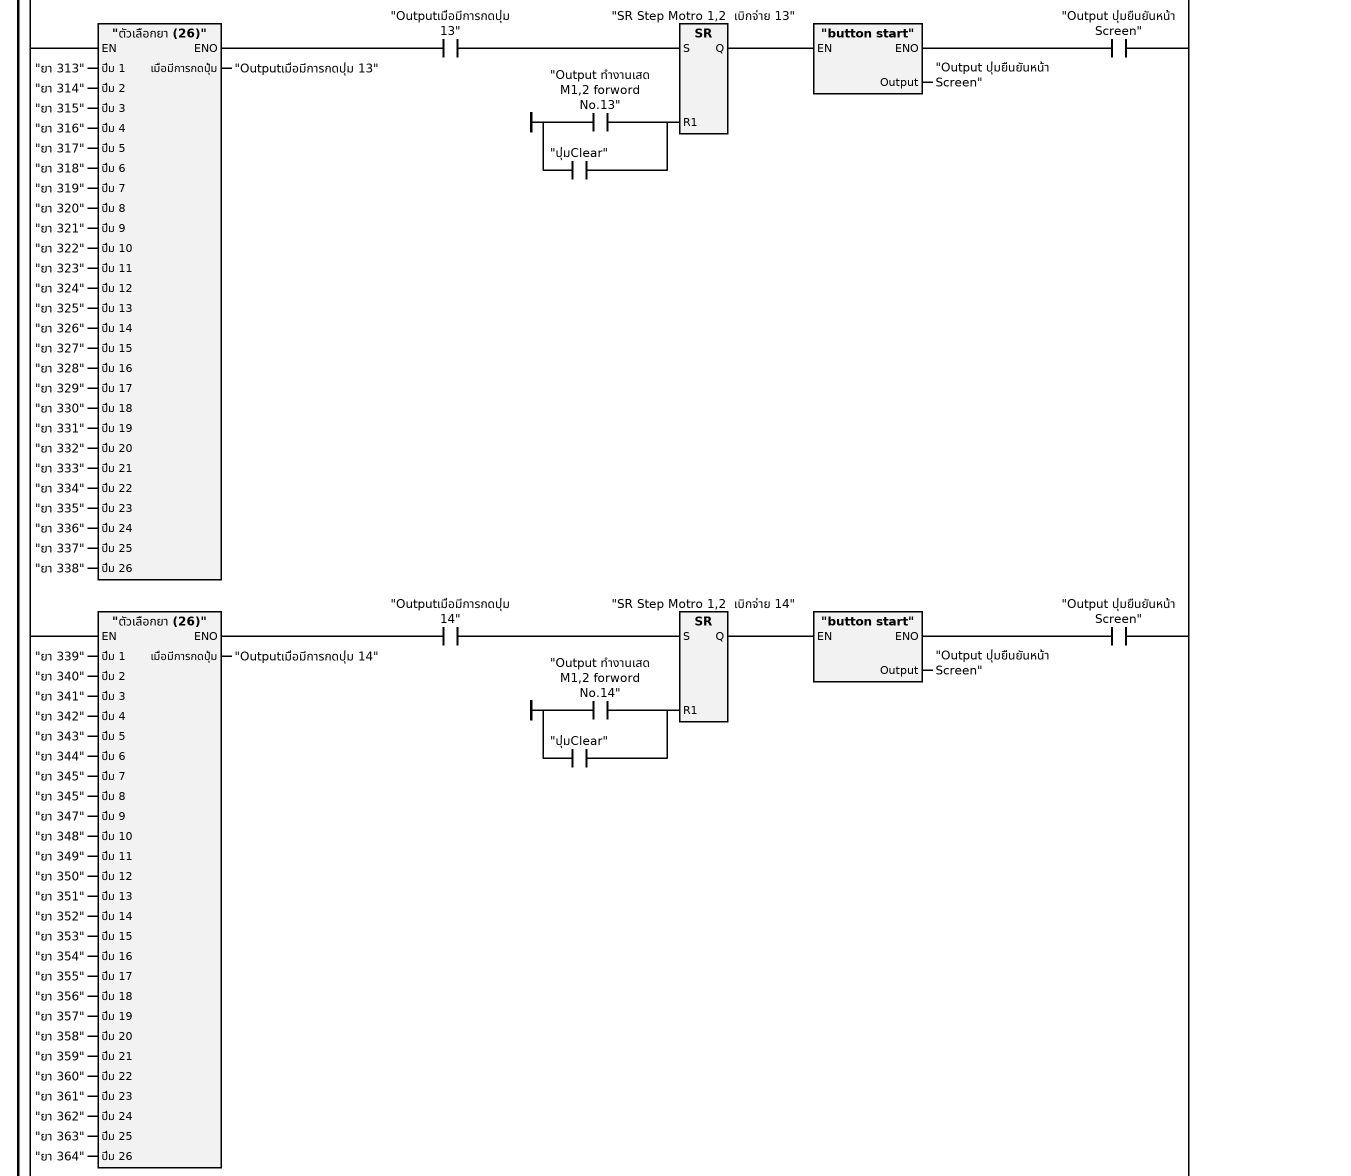
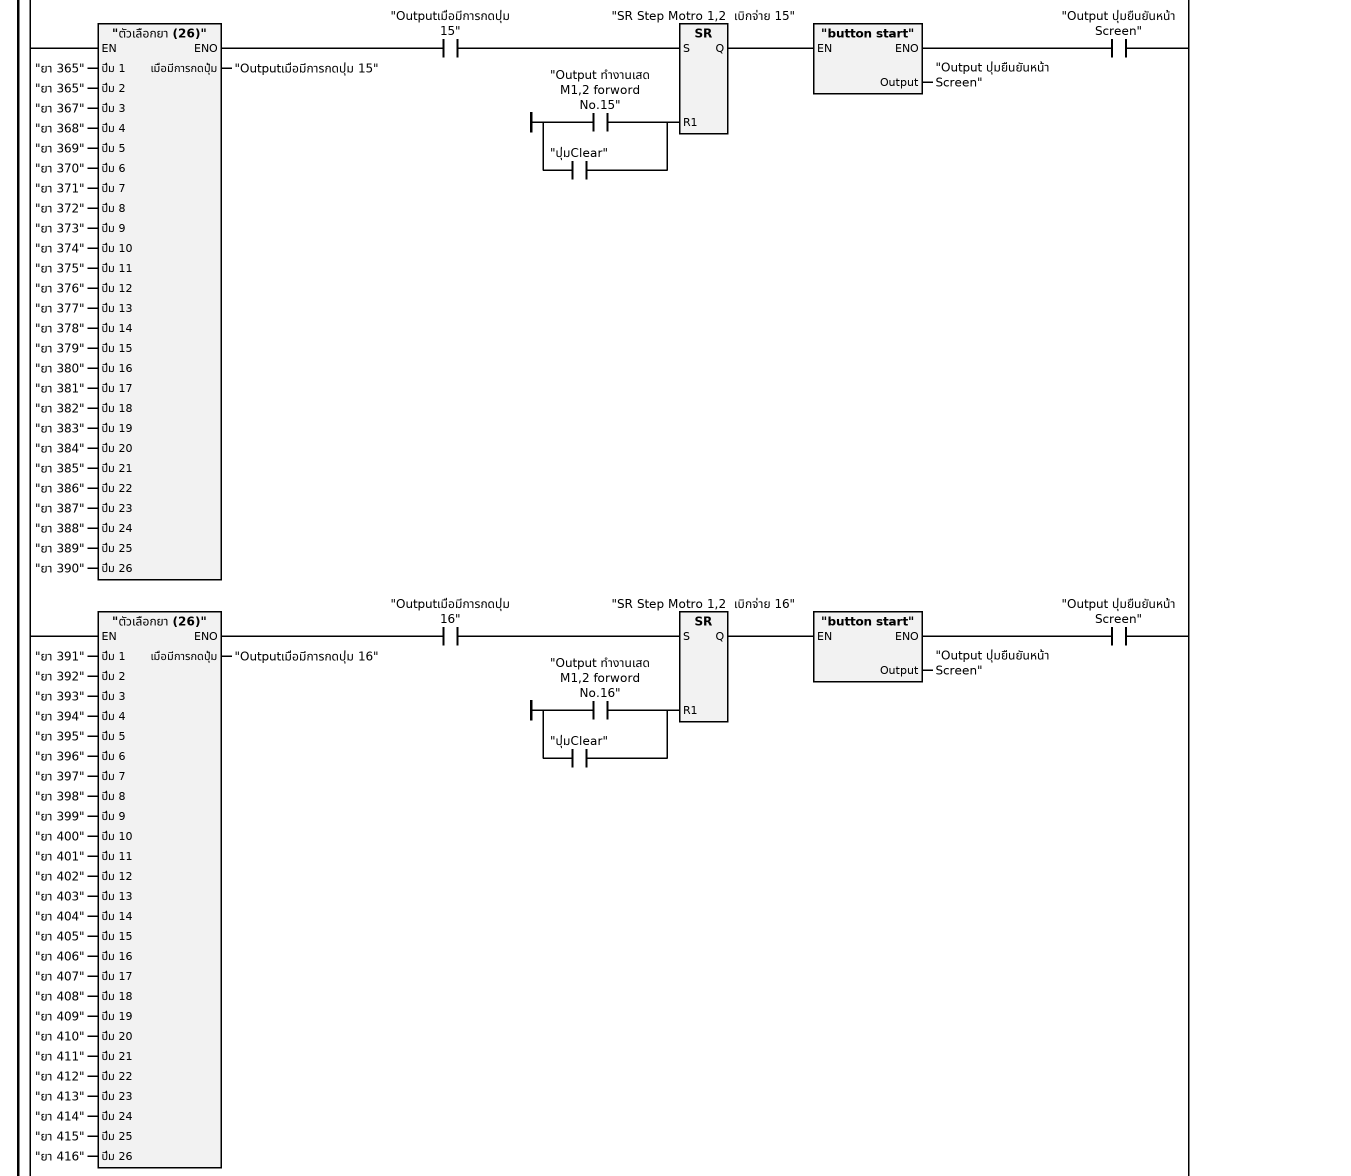
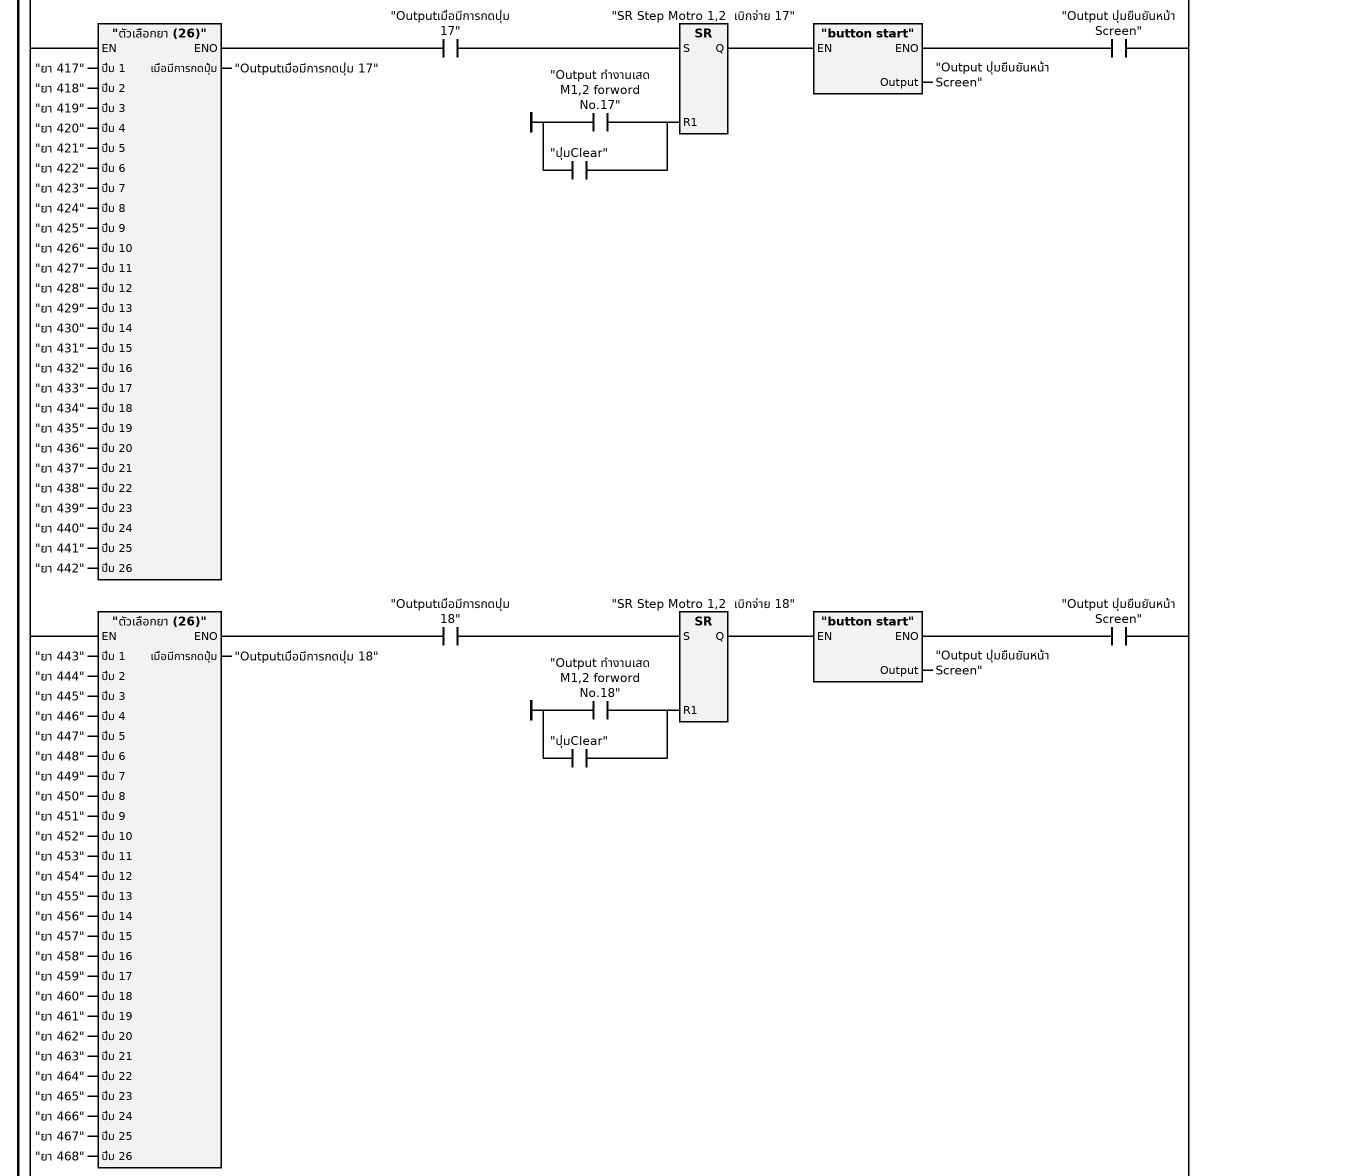
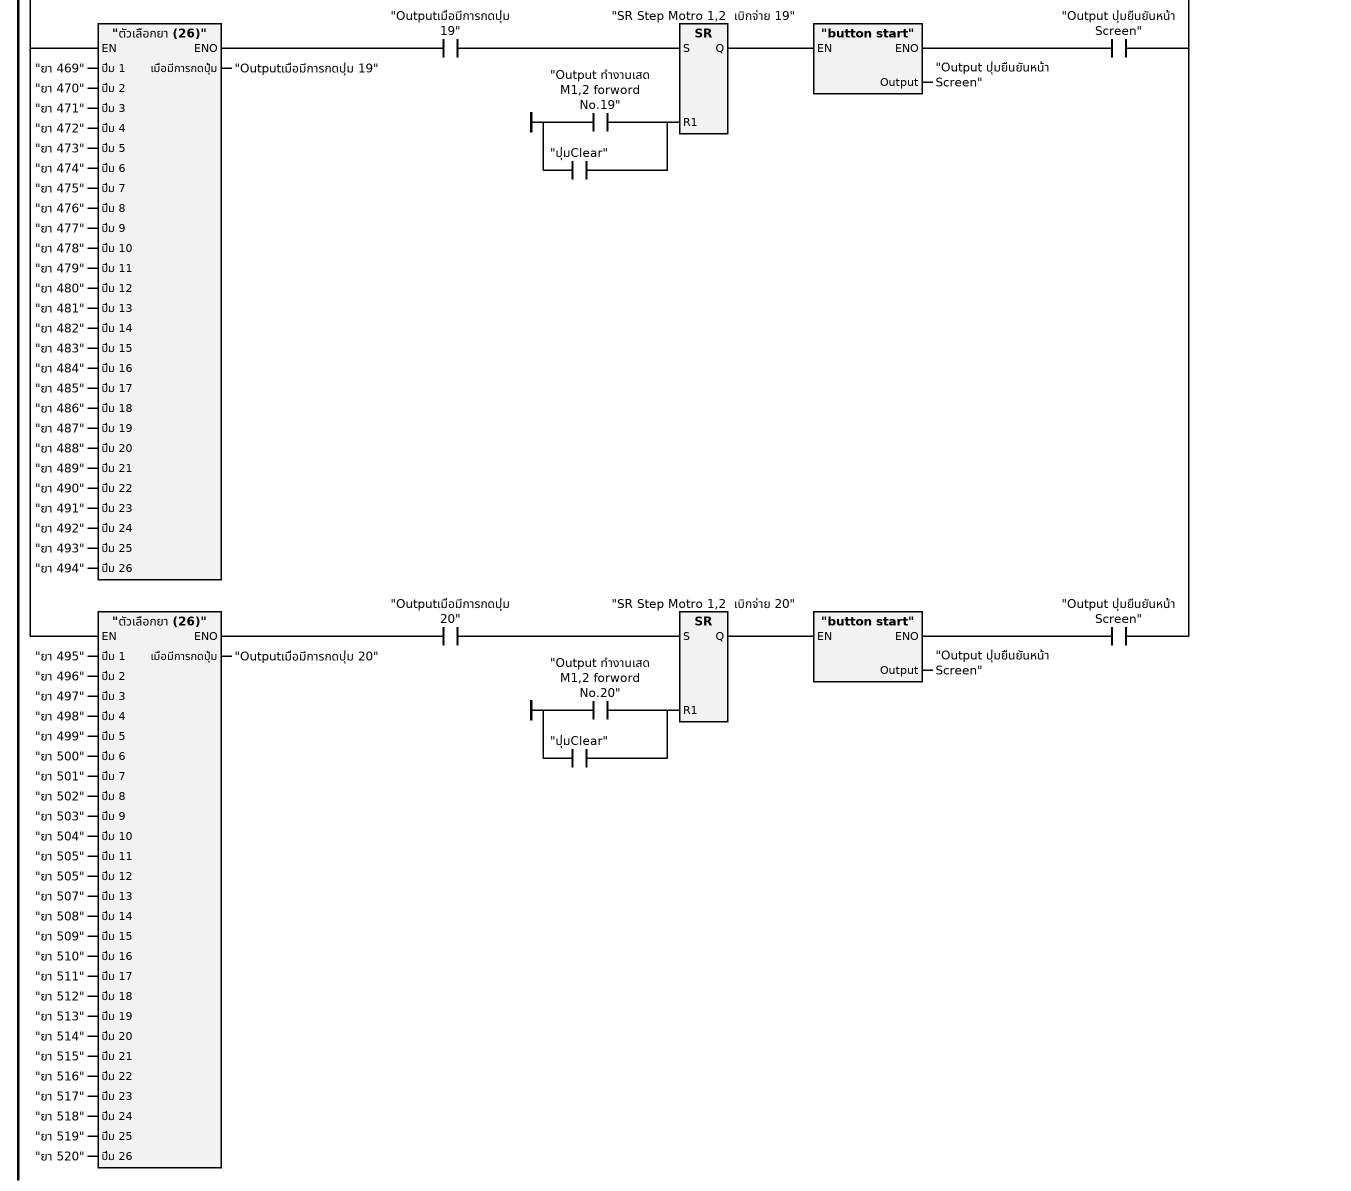
   RUNG wire#powerrail
      "ตัวเลือกยา (26)"("ปึ่ม 1" := "ยา 1", "ปึ่ม 2" := "ยา 2", "ปึ่ม 3" := "ยา 3", "ปึ่ม 4" := "ยา 4", "ปึ่ม 5" := "ยา 5", "ปึ่ม 6" := "ยา 6", "ปึ่ม 7" := "ยา 7", "ปึ่ม 8" := "ยา 8", "ปึ่ม 9" := "ยา 9", "ปึ่ม 10" := "ยา 10", "ปึ่ม 11" := "ยา 11", "ปึ่ม 12" := "ยา 12", "ปึ่ม 13" := "ยา 13", "ปึ่ม 14" := "ยา 14", "ปึ่ม 15" := "ยา 15", "ปึ่ม 16" := "ยา 16", "ปึ่ม 17" := "ยา 17", "ปึ่ม 18" := "ยา 18", "ปึ่ม 19" := "ยา 19", "ปึ่ม 20" := "ยา 20", "ปึ่ม 21" := "ยา 21", "ปึ่ม 22" := "ยา 22", "ปึ่ม 23" := "ยา 23", "ปึ่ม 24" := "ยา 24", "ปึ่ม 25" := "ยา 25", "ปึ่ม 26" := "ยา 26", "เมื่ิอมีการกดปุ้ม" => "Outputเมื่อมีการกดปุ่ม 1")
      Contact( "Outputเมื่อมีการกดปุ่ม 1" )
      S_SR(operand := "SR Step Motro 1,2  เบิกจ่าย 1", r1 := wire#w1)
      "button start"(Output => "Output ปุ่มยืนยันหน้า Screen")
      Contact( "Output ปุ่มยืนยันหน้า Screen" )
      wire#w2
      Coil( #"Stepper Motor  ทำงาน" )
   END_RUNG
   RUNG wire#powerrail
      Contact( "Output ทำงานเสด M1,2 forword No.1" )
   END_RUNG wire#w1
   RUNG wire#powerrail
      Contact( "ปุ่มClear" )
   END_RUNG wire#w1
   RUNG wire#powerrail
      "ตัวเลือกยา (26)"("ปึ่ม 1" := "ยา 27", "ปึ่ม 2" := "ยา 28", "ปึ่ม 3" := "ยา 29", "ปึ่ม 4" := "ยา 30", "ปึ่ม 5" := "ยา 31", "ปึ่ม 6" := "ยา 32", "ปึ่ม 7" := "ยา 33", "ปึ่ม 8" := "ยา 34", "ปึ่ม 9" := "ยา 35", "ปึ่ม 10" := "ยา 36", "ปึ่ม 11" := "ยา 37", "ปึ่ม 12" := "ยา 38", "ปึ่ม 13" := "ยา 39", "ปึ่ม 14" := "ยา 40", "ปึ่ม 15" := "ยา 41", "ปึ่ม 16" := "ยา 42", "ปึ่ม 17" := "ยา 43", "ปึ่ม 18" := "ยา 44", "ปึ่ม 19" := "ยา 45", "ปึ่ม 20" := "ยา 46", "ปึ่ม 21" := "ยา 47", "ปึ่ม 22" := "ยา 48", "ปึ่ม 23" := "ยา 49", "ปึ่ม 24" := "ยา 50", "ปึ่ม 25" := "ยา 51", "ปึ่ม 26" := "ยา 52", "เมื่ิอมีการกดปุ้ม" => "Outputเมื่อมีการกดปุ่ม 2")
      Contact( "Outputเมื่อมีการกดปุ่ม 2" )
      S_SR(operand := "SR Step Motro 1,2  เบิกจ่าย 2", r1 := wire#w3)
      "button start"(Output => "Output ปุ่มยืนยันหน้า Screen")
      Contact( "Output ปุ่มยืนยันหน้า Screen" )
   END_RUNG wire#w2
   RUNG wire#powerrail
      Contact( "Output ทำงานเสด M1,2 forword No.2" )
   END_RUNG wire#w3
   RUNG wire#powerrail
      Contact( "ปุ่มClear" )
   END_RUNG wire#w3
   RUNG wire#powerrail
      "ตัวเลือกยา (26)"("ปึ่ม 1" := "ยา 53", "ปึ่ม 2" := "ยา 54", "ปึ่ม 3" := "ยา 55", "ปึ่ม 4" := "ยา 56", "ปึ่ม 5" := "ยา 57", "ปึ่ม 6" := "ยา 58", "ปึ่ม 7" := "ยา 59", "ปึ่ม 8" := "ยา 60", "ปึ่ม 9" := "ยา 61", "ปึ่ม 10" := "ยา 62", "ปึ่ม 11" := "ยา 63", "ปึ่ม 12" := "ยา 64", "ปึ่ม 13" := "ยา 65", "ปึ่ม 14" := "ยา 66", "ปึ่ม 15" := "ยา 67", "ปึ่ม 16" := "ยา 68", "ปึ่ม 17" := "ยา 69", "ปึ่ม 18" := "ยา 70", "ปึ่ม 19" := "ยา 71", "ปึ่ม 20" := "ยา 72", "ปึ่ม 21" := "ยา 73", "ปึ่ม 22" := "ยา 74", "ปึ่ม 23" := "ยา 75", "ปึ่ม 24" := "ยา 76", "ปึ่ม 25" := "ยา 77", "ปึ่ม 26" := "ยา 78", "เมื่ิอมีการกดปุ้ม" => "Outputเมื่อมีการกดปุ่ม 3")
      Contact( "Outputเมื่อมีการกดปุ่ม 3" )
      S_SR(operand := "SR Step Motro 1,2  เบิกจ่าย 3", r1 := wire#w4)
      "button start"(Output => "Output ปุ่มยืนยันหน้า Screen")
      Contact( "Output ปุ่มยืนยันหน้า Screen" )
   END_RUNG wire#w2
   RUNG wire#powerrail
      Contact( "Output ทำงานเสด M1,2 forword No.3" )
   END_RUNG wire#w4
   RUNG wire#powerrail
      Contact( "ปุ่มClear" )
   END_RUNG wire#w4
   RUNG wire#powerrail
      "ตัวเลือกยา (26)"("ปึ่ม 1" := "ยา 79", "ปึ่ม 2" := "ยา 80", "ปึ่ม 3" := "ยา 81", "ปึ่ม 4" := "ยา 82", "ปึ่ม 5" := "ยา 83", "ปึ่ม 6" := "ยา 84", "ปึ่ม 7" := "ยา 85", "ปึ่ม 8" := "ยา 86", "ปึ่ม 9" := "ยา 87", "ปึ่ม 10" := "ยา 88", "ปึ่ม 11" := "ยา 89", "ปึ่ม 12" := "ยา 90", "ปึ่ม 13" := "ยา 91", "ปึ่ม 14" := "ยา 92", "ปึ่ม 15" := "ยา 93", "ปึ่ม 16" := "ยา 94", "ปึ่ม 17" := "ยา 95", "ปึ่ม 18" := "ยา 96", "ปึ่ม 19" := "ยา 97", "ปึ่ม 20" := "ยา 98", "ปึ่ม 21" := "ยา 99", "ปึ่ม 22" := "ยา 100", "ปึ่ม 23" := "ยา 101", "ปึ่ม 24" := "ยา 102", "ปึ่ม 25" := "ยา 103", "ปึ่ม 26" := "ยา 104", "เมื่ิอมีการกดปุ้ม" => "Outputเมื่อมีการกดปุ่ม 4")
      Contact( "Outputเมื่อมีการกดปุ่ม 4" )
      S_SR(operand := "SR Step Motro 1,2  เบิกจ่าย 4", r1 := wire#w5)
      "button start"(Output => "Output ปุ่มยืนยันหน้า Screen")
      Contact( "Output ปุ่มยืนยันหน้า Screen" )
   END_RUNG wire#w2
   RUNG wire#powerrail
      Contact( "Output ทำงานเสด M1,2 forword No.4" )
   END_RUNG wire#w5
   RUNG wire#powerrail
      Contact( "ปุ่มClear" )
   END_RUNG wire#w5
   RUNG wire#powerrail
      "ตัวเลือกยา (26)"("ปึ่ม 1" := "ยา 105", "ปึ่ม 2" := "ยา 106", "ปึ่ม 3" := "ยา 107", "ปึ่ม 4" := "ยา 108", "ปึ่ม 5" := "ยา 109", "ปึ่ม 6" := "ยา 110", "ปึ่ม 7" := "ยา 111", "ปึ่ม 8" := "ยา 112", "ปึ่ม 9" := "ยา 113", "ปึ่ม 10" := "ยา 114", "ปึ่ม 11" := "ยา 115", "ปึ่ม 12" := "ยา 116", "ปึ่ม 13" := "ยา 117", "ปึ่ม 14" := "ยา 118", "ปึ่ม 15" := "ยา 119", "ปึ่ม 16" := "ยา 120", "ปึ่ม 17" := "ยา 121", "ปึ่ม 18" := "ยา 122", "ปึ่ม 19" := "ยา 123", "ปึ่ม 20" := "ยา 124", "ปึ่ม 21" := "ยา 125", "ปึ่ม 22" := "ยา 126", "ปึ่ม 23" := "ยา 127", "ปึ่ม 24" := "ยา 128", "ปึ่ม 25" := "ยา 129", "ปึ่ม 26" := "ยา 130", "เมื่ิอมีการกดปุ้ม" => "Outputเมื่อมีการกดปุ่ม 5")
      Contact( "Outputเมื่อมีการกดปุ่ม 5" )
      S_SR(operand := "SR Step Motro 1,2  เบิกจ่าย 5", r1 := wire#w6)
      "button start"(Output => "Output ปุ่มยืนยันหน้า Screen")
      Contact( "Output ปุ่มยืนยันหน้า Screen" )
   END_RUNG wire#w2
   RUNG wire#powerrail
      Contact( "Output ทำงานเสด M1,2 forword No.5" )
   END_RUNG wire#w6
   RUNG wire#powerrail
      Contact( "ปุ่มClear" )
   END_RUNG wire#w6
   RUNG wire#powerrail
      "ตัวเลือกยา (26)"("ปึ่ม 1" := "ยา 131", "ปึ่ม 2" := "ยา 132", "ปึ่ม 3" := "ยา 133", "ปึ่ม 4" := "ยา 134", "ปึ่ม 5" := "ยา 135", "ปึ่ม 6" := "ยา 136", "ปึ่ม 7" := "ยา 137", "ปึ่ม 8" := "ยา 138", "ปึ่ม 9" := "ยา 139", "ปึ่ม 10" := "ยา 140", "ปึ่ม 11" := "ยา 141", "ปึ่ม 12" := "ยา 142", "ปึ่ม 13" := "ยา 143", "ปึ่ม 14" := "ยา 144", "ปึ่ม 15" := "ยา 145", "ปึ่ม 16" := "ยา 146", "ปึ่ม 17" := "ยา 147", "ปึ่ม 18" := "ยา 148", "ปึ่ม 19" := "ยา 149", "ปึ่ม 20" := "ยา 150", "ปึ่ม 21" := "ยา 151", "ปึ่ม 22" := "ยา 152", "ปึ่ม 23" := "ยา 153", "ปึ่ม 24" := "ยา 154", "ปึ่ม 25" := "ยา 155", "ปึ่ม 26" := "ยา 156", "เมื่ิอมีการกดปุ้ม" => "Outputเมื่อมีการกดปุ่ม 6")
      Contact( "Outputเมื่อมีการกดปุ่ม 6" )
      S_SR(operand := "SR Step Motro 1,2  เบิกจ่าย 6", r1 := wire#w7)
      "button start"(Output => "Output ปุ่มยืนยันหน้า Screen")
      Contact( "Output ปุ่มยืนยันหน้า Screen" )
   END_RUNG wire#w2
   RUNG wire#powerrail
      Contact( "Output ทำงานเสด M1,2 forword No.6" )
   END_RUNG wire#w7
   RUNG wire#powerrail
      Contact( "ปุ่มClear" )
   END_RUNG wire#w7
   RUNG wire#powerrail
      "ตัวเลือกยา (26)"("ปึ่ม 1" := "ยา 157", "ปึ่ม 2" := "ยา 158", "ปึ่ม 3" := "ยา 159", "ปึ่ม 4" := "ยา 160", "ปึ่ม 5" := "ยา 161", "ปึ่ม 6" := "ยา 162", "ปึ่ม 7" := "ยา 163", "ปึ่ม 8" := "ยา 164", "ปึ่ม 9" := "ยา 165", "ปึ่ม 10" := "ยา 166", "ปึ่ม 11" := "ยา 167", "ปึ่ม 12" := "ยา 168", "ปึ่ม 13" := "ยา 169", "ปึ่ม 14" := "ยา 170", "ปึ่ม 15" := "ยา 171", "ปึ่ม 16" := "ยา 172", "ปึ่ม 17" := "ยา 173", "ปึ่ม 18" := "ยา 174", "ปึ่ม 19" := "ยา 175", "ปึ่ม 20" := "ยา 176", "ปึ่ม 21" := "ยา 177", "ปึ่ม 22" := "ยา 178", "ปึ่ม 23" := "ยา 179", "ปึ่ม 24" := "ยา 180", "ปึ่ม 25" := "ยา 181", "ปึ่ม 26" := "ยา 182", "เมื่ิอมีการกดปุ้ม" => "Outputเมื่อมีการกดปุ่ม 7")
      Contact( "Outputเมื่อมีการกดปุ่ม 7" )
      S_SR(operand := "SR Step Motro 1,2  เบิกจ่าย 7", r1 := wire#w8)
      "button start"(Output => "Output ปุ่มยืนยันหน้า Screen")
      Contact( "Output ปุ่มยืนยันหน้า Screen" )
   END_RUNG wire#w2
   RUNG wire#powerrail
      Contact( "Output ทำงานเสด M1,2 forword No.7" )
   END_RUNG wire#w8
   RUNG wire#powerrail
      Contact( "ปุ่มClear" )
   END_RUNG wire#w8
   RUNG wire#powerrail
      "ตัวเลือกยา (26)"("ปึ่ม 1" := "ยา 183", "ปึ่ม 2" := "ยา 184", "ปึ่ม 3" := "ยา 185", "ปึ่ม 4" := "ยา 186", "ปึ่ม 5" := "ยา 187", "ปึ่ม 6" := "ยา 188", "ปึ่ม 7" := "ยา 189", "ปึ่ม 8" := "ยา 190", "ปึ่ม 9" := "ยา 191", "ปึ่ม 10" := "ยา 192", "ปึ่ม 11" := "ยา 193", "ปึ่ม 12" := "ยา 194", "ปึ่ม 13" := "ยา 195", "ปึ่ม 14" := "ยา 196", "ปึ่ม 15" := "ยา 197", "ปึ่ม 16" := "ยา 198", "ปึ่ม 17" := "ยา 199", "ปึ่ม 18" := "ยา 200", "ปึ่ม 19" := "ยา 201", "ปึ่ม 20" := "ยา 202", "ปึ่ม 21" := "ยา 203", "ปึ่ม 22" := "ยา 204", "ปึ่ม 23" := "ยา 205", "ปึ่ม 24" := "ยา 206", "ปึ่ม 25" := "ยา 207", "ปึ่ม 26" := "ยา 208", "เมื่ิอมีการกดปุ้ม" => "Outputเมื่อมีการกดปุ่ม 8")
      Contact( "Outputเมื่อมีการกดปุ่ม 8" )
      S_SR(operand := "SR Step Motro 1,2  เบิกจ่าย 8", r1 := wire#w9)
      "button start"(Output => "Output ปุ่มยืนยันหน้า Screen")
      Contact( "Output ปุ่มยืนยันหน้า Screen" )
   END_RUNG wire#w2
   RUNG wire#powerrail
      Contact( "Output ทำงานเสด M1,2 forword No.8" )
   END_RUNG wire#w9
   RUNG wire#powerrail
      Contact( "ปุ่มClear" )
   END_RUNG wire#w9
   RUNG wire#powerrail
      "ตัวเลือกยา (26)"("ปึ่ม 1" := "ยา 209", "ปึ่ม 2" := "ยา 210", "ปึ่ม 3" := "ยา 211", "ปึ่ม 4" := "ยา 212", "ปึ่ม 5" := "ยา 213", "ปึ่ม 6" := "ยา 214", "ปึ่ม 7" := "ยา 215", "ปึ่ม 8" := "ยา 216", "ปึ่ม 9" := "ยา 217", "ปึ่ม 10" := "ยา 218", "ปึ่ม 11" := "ยา 219", "ปึ่ม 12" := "ยา 220", "ปึ่ม 13" := "ยา 221", "ปึ่ม 14" := "ยา 222", "ปึ่ม 15" := "ยา 223", "ปึ่ม 16" := "ยา 224", "ปึ่ม 17" := "ยา 225", "ปึ่ม 18" := "ยา 226", "ปึ่ม 19" := "ยา 227", "ปึ่ม 20" := "ยา 228", "ปึ่ม 21" := "ยา 229", "ปึ่ม 22" := "ยา 230", "ปึ่ม 23" := "ยา 231", "ปึ่ม 24" := "ยา 232", "ปึ่ม 25" := "ยา 233", "ปึ่ม 26" := "ยา 234", "เมื่ิอมีการกดปุ้ม" => "Outputเมื่อมีการกดปุ่ม 9")
      Contact( "Outputเมื่อมีการกดปุ่ม 9" )
      S_SR(operand := "SR Step Motro 1,2  เบิกจ่าย 9", r1 := wire#w10)
      "button start"(Output => "Output ปุ่มยืนยันหน้า Screen")
      Contact( "Output ปุ่มยืนยันหน้า Screen" )
   END_RUNG wire#w2
   RUNG wire#powerrail
      Contact( "Output ทำงานเสด M1,2 forword No.9" )
   END_RUNG wire#w10
   RUNG wire#powerrail
      Contact( "ปุ่มClear" )
   END_RUNG wire#w10
   RUNG wire#powerrail
      "ตัวเลือกยา (26)"("ปึ่ม 1" := "ยา 235", "ปึ่ม 2" := "ยา 236", "ปึ่ม 3" := "ยา 234", "ปึ่ม 4" := "ยา 238", "ปึ่ม 5" := "ยา 239", "ปึ่ม 6" := "ยา 240", "ปึ่ม 7" := "ยา 241", "ปึ่ม 8" := "ยา 242", "ปึ่ม 9" := "ยา 243", "ปึ่ม 10" := "ยา 244", "ปึ่ม 11" := "ยา 245", "ปึ่ม 12" := "ยา 246", "ปึ่ม 13" := "ยา 247", "ปึ่ม 14" := "ยา 248", "ปึ่ม 15" := "ยา 249", "ปึ่ม 16" := "ยา 250", "ปึ่ม 17" := "ยา 251", "ปึ่ม 18" := "ยา 252", "ปึ่ม 19" := "ยา 253", "ปึ่ม 20" := "ยา 254", "ปึ่ม 21" := "ยา 255", "ปึ่ม 22" := "ยา 256", "ปึ่ม 23" := "ยา 257", "ปึ่ม 24" := "ยา 258", "ปึ่ม 25" := "ยา 259", "ปึ่ม 26" := "ยา 260", "เมื่ิอมีการกดปุ้ม" => "Outputเมื่อมีการกดปุ่ม 10")
      Contact( "Outputเมื่อมีการกดปุ่ม 10" )
      S_SR(operand := "SR Step Motro 1,2  เบิกจ่าย 10", r1 := wire#w11)
      "button start"(Output => "Output ปุ่มยืนยันหน้า Screen")
      Contact( "Output ปุ่มยืนยันหน้า Screen" )
   END_RUNG wire#w2
   RUNG wire#powerrail
      Contact( "Output ทำงานเสด M1,2 forword No.10" )
   END_RUNG wire#w11
   RUNG wire#powerrail
      Contact( "ปุ่มClear" )
   END_RUNG wire#w11
   RUNG wire#powerrail
      "ตัวเลือกยา (26)"("ปึ่ม 1" := "ยา 261", "ปึ่ม 2" := "ยา 262", "ปึ่ม 3" := "ยา 263", "ปึ่ม 4" := "ยา 264", "ปึ่ม 5" := "ยา 265", "ปึ่ม 6" := "ยา 266", "ปึ่ม 7" := "ยา 267", "ปึ่ม 8" := "ยา 268", "ปึ่ม 9" := "ยา 269", "ปึ่ม 10" := "ยา 270", "ปึ่ม 11" := "ยา 271", "ปึ่ม 12" := "ยา 272", "ปึ่ม 13" := "ยา 273", "ปึ่ม 14" := "ยา 274", "ปึ่ม 15" := "ยา 275", "ปึ่ม 16" := "ยา 276", "ปึ่ม 17" := "ยา 277", "ปึ่ม 18" := "ยา 278", "ปึ่ม 19" := "ยา 279", "ปึ่ม 20" := "ยา 280", "ปึ่ม 21" := "ยา 281", "ปึ่ม 22" := "ยา 282", "ปึ่ม 23" := "ยา 283", "ปึ่ม 24" := "ยา 284", "ปึ่ม 25" := "ยา 285", "ปึ่ม 26" := "ยา 286", "เมื่ิอมีการกดปุ้ม" => "Outputเมื่อมีการกดปุ่ม 11")
      Contact( "Outputเมื่อมีการกดปุ่ม 11" )
      S_SR(operand := "SR Step Motro 1,2  เบิกจ่าย 11", r1 := wire#w12)
      "button start"(Output => "Output ปุ่มยืนยันหน้า Screen")
      Contact( "Output ปุ่มยืนยันหน้า Screen" )
   END_RUNG wire#w2
   RUNG wire#powerrail
      Contact( "Output ทำงานเสด M1,2 forword No.11" )
   END_RUNG wire#w12
   RUNG wire#powerrail
      Contact( "ปุ่มClear" )
   END_RUNG wire#w12
   RUNG wire#powerrail
      "ตัวเลือกยา (26)"("ปึ่ม 1" := "ยา 287", "ปึ่ม 2" := "ยา 288", "ปึ่ม 3" := "ยา 289", "ปึ่ม 4" := "ยา 290", "ปึ่ม 5" := "ยา 291", "ปึ่ม 6" := "ยา 292", "ปึ่ม 7" := "ยา 293", "ปึ่ม 8" := "ยา 294", "ปึ่ม 9" := "ยา 295", "ปึ่ม 10" := "ยา 296", "ปึ่ม 11" := "ยา 297", "ปึ่ม 12" := "ยา 298", "ปึ่ม 13" := "ยา 299", "ปึ่ม 14" := "ยา 300", "ปึ่ม 15" := "ยา 301", "ปึ่ม 16" := "ยา 302", "ปึ่ม 17" := "ยา 303", "ปึ่ม 18" := "ยา 304", "ปึ่ม 19" := "ยา 305", "ปึ่ม 20" := "ยา 306", "ปึ่ม 21" := "ยา 307", "ปึ่ม 22" := "ยา 308", "ปึ่ม 23" := "ยา 309", "ปึ่ม 24" := "ยา 310", "ปึ่ม 25" := "ยา 311", "ปึ่ม 26" := "ยา 312", "เมื่ิอมีการกดปุ้ม" => "Outputเมื่อมีการกดปุ่ม 12")
      Contact( "Outputเมื่อมีการกดปุ่ม 12" )
      S_SR(operand := "SR Step Motro 1,2  เบิกจ่าย 12", r1 := wire#w13)
      "button start"(Output => "Output ปุ่มยืนยันหน้า Screen")
      Contact( "Output ปุ่มยืนยันหน้า Screen" )
   END_RUNG wire#w2
   RUNG wire#powerrail
      Contact( "Output ทำงานเสด M1,2 forword No.12" )
   END_RUNG wire#w13
   RUNG wire#powerrail
      Contact( "ปุ่มClear" )
   END_RUNG wire#w13
   RUNG wire#powerrail
      "ตัวเลือกยา (26)"("ปึ่ม 1" := "ยา 313", "ปึ่ม 2" := "ยา 314", "ปึ่ม 3" := "ยา 315", "ปึ่ม 4" := "ยา 316", "ปึ่ม 5" := "ยา 317", "ปึ่ม 6" := "ยา 318", "ปึ่ม 7" := "ยา 319", "ปึ่ม 8" := "ยา 320", "ปึ่ม 9" := "ยา 321", "ปึ่ม 10" := "ยา 322", "ปึ่ม 11" := "ยา 323", "ปึ่ม 12" := "ยา 324", "ปึ่ม 13" := "ยา 325", "ปึ่ม 14" := "ยา 326", "ปึ่ม 15" := "ยา 327", "ปึ่ม 16" := "ยา 328", "ปึ่ม 17" := "ยา 329", "ปึ่ม 18" := "ยา 330", "ปึ่ม 19" := "ยา 331", "ปึ่ม 20" := "ยา 332", "ปึ่ม 21" := "ยา 333", "ปึ่ม 22" := "ยา 334", "ปึ่ม 23" := "ยา 335", "ปึ่ม 24" := "ยา 336", "ปึ่ม 25" := "ยา 337", "ปึ่ม 26" := "ยา 338", "เมื่ิอมีการกดปุ้ม" => "Outputเมื่อมีการกดปุ่ม 13")
      Contact( "Outputเมื่อมีการกดปุ่ม 13" )
      S_SR(operand := "SR Step Motro 1,2  เบิกจ่าย 13", r1 := wire#w14)
      "button start"(Output => "Output ปุ่มยืนยันหน้า Screen")
      Contact( "Output ปุ่มยืนยันหน้า Screen" )
   END_RUNG wire#w2
   RUNG wire#powerrail
      Contact( "Output ทำงานเสด M1,2 forword No.13" )
   END_RUNG wire#w14
   RUNG wire#powerrail
      Contact( "ปุ่มClear" )
   END_RUNG wire#w14
   RUNG wire#powerrail
      "ตัวเลือกยา (26)"("ปึ่ม 1" := "ยา 339", "ปึ่ม 2" := "ยา 340", "ปึ่ม 3" := "ยา 341", "ปึ่ม 4" := "ยา 342", "ปึ่ม 5" := "ยา 343", "ปึ่ม 6" := "ยา 344", "ปึ่ม 7" := "ยา 345", "ปึ่ม 8" := "ยา 345", "ปึ่ม 9" := "ยา 347", "ปึ่ม 10" := "ยา 348", "ปึ่ม 11" := "ยา 349", "ปึ่ม 12" := "ยา 350", "ปึ่ม 13" := "ยา 351", "ปึ่ม 14" := "ยา 352", "ปึ่ม 15" := "ยา 353", "ปึ่ม 16" := "ยา 354", "ปึ่ม 17" := "ยา 355", "ปึ่ม 18" := "ยา 356", "ปึ่ม 19" := "ยา 357", "ปึ่ม 20" := "ยา 358", "ปึ่ม 21" := "ยา 359", "ปึ่ม 22" := "ยา 360", "ปึ่ม 23" := "ยา 361", "ปึ่ม 24" := "ยา 362", "ปึ่ม 25" := "ยา 363", "ปึ่ม 26" := "ยา 364", "เมื่ิอมีการกดปุ้ม" => "Outputเมื่อมีการกดปุ่ม 14")
      Contact( "Outputเมื่อมีการกดปุ่ม 14" )
      S_SR(operand := "SR Step Motro 1,2  เบิกจ่าย 14", r1 := wire#w15)
      "button start"(Output => "Output ปุ่มยืนยันหน้า Screen")
      Contact( "Output ปุ่มยืนยันหน้า Screen" )
   END_RUNG wire#w2
   RUNG wire#powerrail
      Contact( "Output ทำงานเสด M1,2 forword No.14" )
   END_RUNG wire#w15
   RUNG wire#powerrail
      Contact( "ปุ่มClear" )
   END_RUNG wire#w15
   RUNG wire#powerrail
      "ตัวเลือกยา (26)"("ปึ่ม 1" := "ยา 365", "ปึ่ม 2" := "ยา 365", "ปึ่ม 3" := "ยา 367", "ปึ่ม 4" := "ยา 368", "ปึ่ม 5" := "ยา 369", "ปึ่ม 6" := "ยา 370", "ปึ่ม 7" := "ยา 371", "ปึ่ม 8" := "ยา 372", "ปึ่ม 9" := "ยา 373", "ปึ่ม 10" := "ยา 374", "ปึ่ม 11" := "ยา 375", "ปึ่ม 12" := "ยา 376", "ปึ่ม 13" := "ยา 377", "ปึ่ม 14" := "ยา 378", "ปึ่ม 15" := "ยา 379", "ปึ่ม 16" := "ยา 380", "ปึ่ม 17" := "ยา 381", "ปึ่ม 18" := "ยา 382", "ปึ่ม 19" := "ยา 383", "ปึ่ม 20" := "ยา 384", "ปึ่ม 21" := "ยา 385", "ปึ่ม 22" := "ยา 386", "ปึ่ม 23" := "ยา 387", "ปึ่ม 24" := "ยา 388", "ปึ่ม 25" := "ยา 389", "ปึ่ม 26" := "ยา 390", "เมื่ิอมีการกดปุ้ม" => "Outputเมื่อมีการกดปุ่ม 15")
      Contact( "Outputเมื่อมีการกดปุ่ม 15" )
      S_SR(operand := "SR Step Motro 1,2  เบิกจ่าย 15", r1 := wire#w16)
      "button start"(Output => "Output ปุ่มยืนยันหน้า Screen")
      Contact( "Output ปุ่มยืนยันหน้า Screen" )
   END_RUNG wire#w2
   RUNG wire#powerrail
      Contact( "Output ทำงานเสด M1,2 forword No.15" )
   END_RUNG wire#w16
   RUNG wire#powerrail
      Contact( "ปุ่มClear" )
   END_RUNG wire#w16
   RUNG wire#powerrail
      "ตัวเลือกยา (26)"("ปึ่ม 1" := "ยา 391", "ปึ่ม 2" := "ยา 392", "ปึ่ม 3" := "ยา 393", "ปึ่ม 4" := "ยา 394", "ปึ่ม 5" := "ยา 395", "ปึ่ม 6" := "ยา 396", "ปึ่ม 7" := "ยา 397", "ปึ่ม 8" := "ยา 398", "ปึ่ม 9" := "ยา 399", "ปึ่ม 10" := "ยา 400", "ปึ่ม 11" := "ยา 401", "ปึ่ม 12" := "ยา 402", "ปึ่ม 13" := "ยา 403", "ปึ่ม 14" := "ยา 404", "ปึ่ม 15" := "ยา 405", "ปึ่ม 16" := "ยา 406", "ปึ่ม 17" := "ยา 407", "ปึ่ม 18" := "ยา 408", "ปึ่ม 19" := "ยา 409", "ปึ่ม 20" := "ยา 410", "ปึ่ม 21" := "ยา 411", "ปึ่ม 22" := "ยา 412", "ปึ่ม 23" := "ยา 413", "ปึ่ม 24" := "ยา 414", "ปึ่ม 25" := "ยา 415", "ปึ่ม 26" := "ยา 416", "เมื่ิอมีการกดปุ้ม" => "Outputเมื่อมีการกดปุ่ม 16")
      Contact( "Outputเมื่อมีการกดปุ่ม 16" )
      S_SR(operand := "SR Step Motro 1,2  เบิกจ่าย 16", r1 := wire#w17)
      "button start"(Output => "Output ปุ่มยืนยันหน้า Screen")
      Contact( "Output ปุ่มยืนยันหน้า Screen" )
   END_RUNG wire#w2
   RUNG wire#powerrail
      Contact( "Output ทำงานเสด M1,2 forword No.16" )
   END_RUNG wire#w17
   RUNG wire#powerrail
      Contact( "ปุ่มClear" )
   END_RUNG wire#w17
   RUNG wire#powerrail
      "ตัวเลือกยา (26)"("ปึ่ม 1" := "ยา 417", "ปึ่ม 2" := "ยา 418", "ปึ่ม 3" := "ยา 419", "ปึ่ม 4" := "ยา 420", "ปึ่ม 5" := "ยา 421", "ปึ่ม 6" := "ยา 422", "ปึ่ม 7" := "ยา 423", "ปึ่ม 8" := "ยา 424", "ปึ่ม 9" := "ยา 425", "ปึ่ม 10" := "ยา 426", "ปึ่ม 11" := "ยา 427", "ปึ่ม 12" := "ยา 428", "ปึ่ม 13" := "ยา 429", "ปึ่ม 14" := "ยา 430", "ปึ่ม 15" := "ยา 431", "ปึ่ม 16" := "ยา 432", "ปึ่ม 17" := "ยา 433", "ปึ่ม 18" := "ยา 434", "ปึ่ม 19" := "ยา 435", "ปึ่ม 20" := "ยา 436", "ปึ่ม 21" := "ยา 437", "ปึ่ม 22" := "ยา 438", "ปึ่ม 23" := "ยา 439", "ปึ่ม 24" := "ยา 440", "ปึ่ม 25" := "ยา 441", "ปึ่ม 26" := "ยา 442", "เมื่ิอมีการกดปุ้ม" => "Outputเมื่อมีการกดปุ่ม 17")
      Contact( "Outputเมื่อมีการกดปุ่ม 17" )
      S_SR(operand := "SR Step Motro 1,2  เบิกจ่าย 17", r1 := wire#w18)
      "button start"(Output => "Output ปุ่มยืนยันหน้า Screen")
      Contact( "Output ปุ่มยืนยันหน้า Screen" )
   END_RUNG wire#w2
   RUNG wire#powerrail
      Contact( "Output ทำงานเสด M1,2 forword No.17" )
   END_RUNG wire#w18
   RUNG wire#powerrail
      Contact( "ปุ่มClear" )
   END_RUNG wire#w18
   RUNG wire#powerrail
      "ตัวเลือกยา (26)"("ปึ่ม 1" := "ยา 443", "ปึ่ม 2" := "ยา 444", "ปึ่ม 3" := "ยา 445", "ปึ่ม 4" := "ยา 446", "ปึ่ม 5" := "ยา 447", "ปึ่ม 6" := "ยา 448", "ปึ่ม 7" := "ยา 449", "ปึ่ม 8" := "ยา 450", "ปึ่ม 9" := "ยา 451", "ปึ่ม 10" := "ยา 452", "ปึ่ม 11" := "ยา 453", "ปึ่ม 12" := "ยา 454", "ปึ่ม 13" := "ยา 455", "ปึ่ม 14" := "ยา 456", "ปึ่ม 15" := "ยา 457", "ปึ่ม 16" := "ยา 458", "ปึ่ม 17" := "ยา 459", "ปึ่ม 18" := "ยา 460", "ปึ่ม 19" := "ยา 461", "ปึ่ม 20" := "ยา 462", "ปึ่ม 21" := "ยา 463", "ปึ่ม 22" := "ยา 464", "ปึ่ม 23" := "ยา 465", "ปึ่ม 24" := "ยา 466", "ปึ่ม 25" := "ยา 467", "ปึ่ม 26" := "ยา 468", "เมื่ิอมีการกดปุ้ม" => "Outputเมื่อมีการกดปุ่ม 18")
      Contact( "Outputเมื่อมีการกดปุ่ม 18" )
      S_SR(operand := "SR Step Motro 1,2  เบิกจ่าย 18", r1 := wire#w19)
      "button start"(Output => "Output ปุ่มยืนยันหน้า Screen")
      Contact( "Output ปุ่มยืนยันหน้า Screen" )
   END_RUNG wire#w2
   RUNG wire#powerrail
      Contact( "Output ทำงานเสด M1,2 forword No.18" )
   END_RUNG wire#w19
   RUNG wire#powerrail
      Contact( "ปุ่มClear" )
   END_RUNG wire#w19
   RUNG wire#powerrail
      "ตัวเลือกยา (26)"("ปึ่ม 1" := "ยา 469", "ปึ่ม 2" := "ยา 470", "ปึ่ม 3" := "ยา 471", "ปึ่ม 4" := "ยา 472", "ปึ่ม 5" := "ยา 473", "ปึ่ม 6" := "ยา 474", "ปึ่ม 7" := "ยา 475", "ปึ่ม 8" := "ยา 476", "ปึ่ม 9" := "ยา 477", "ปึ่ม 10" := "ยา 478", "ปึ่ม 11" := "ยา 479", "ปึ่ม 12" := "ยา 480", "ปึ่ม 13" := "ยา 481", "ปึ่ม 14" := "ยา 482", "ปึ่ม 15" := "ยา 483", "ปึ่ม 16" := "ยา 484", "ปึ่ม 17" := "ยา 485", "ปึ่ม 18" := "ยา 486", "ปึ่ม 19" := "ยา 487", "ปึ่ม 20" := "ยา 488", "ปึ่ม 21" := "ยา 489", "ปึ่ม 22" := "ยา 490", "ปึ่ม 23" := "ยา 491", "ปึ่ม 24" := "ยา 492", "ปึ่ม 25" := "ยา 493", "ปึ่ม 26" := "ยา 494", "เมื่ิอมีการกดปุ้ม" => "Outputเมื่อมีการกดปุ่ม 19")
      Contact( "Outputเมื่อมีการกดปุ่ม 19" )
      S_SR(operand := "SR Step Motro 1,2  เบิกจ่าย 19", r1 := wire#w20)
      "button start"(Output => "Output ปุ่มยืนยันหน้า Screen")
      Contact( "Output ปุ่มยืนยันหน้า Screen" )
   END_RUNG wire#w2
   RUNG wire#powerrail
      Contact( "Output ทำงานเสด M1,2 forword No.19" )
   END_RUNG wire#w20
   RUNG wire#powerrail
      Contact( "ปุ่มClear" )
   END_RUNG wire#w20
   RUNG wire#powerrail
      "ตัวเลือกยา (26)"("ปึ่ม 1" := "ยา 495", "ปึ่ม 2" := "ยา 496", "ปึ่ม 3" := "ยา 497", "ปึ่ม 4" := "ยา 498", "ปึ่ม 5" := "ยา 499", "ปึ่ม 6" := "ยา 500", "ปึ่ม 7" := "ยา 501", "ปึ่ม 8" := "ยา 502", "ปึ่ม 9" := "ยา 503", "ปึ่ม 10" := "ยา 504", "ปึ่ม 11" := "ยา 505", "ปึ่ม 12" := "ยา 505", "ปึ่ม 13" := "ยา 507", "ปึ่ม 14" := "ยา 508", "ปึ่ม 15" := "ยา 509", "ปึ่ม 16" := "ยา 510", "ปึ่ม 17" := "ยา 511", "ปึ่ม 18" := "ยา 512", "ปึ่ม 19" := "ยา 513", "ปึ่ม 20" := "ยา 514", "ปึ่ม 21" := "ยา 515", "ปึ่ม 22" := "ยา 516", "ปึ่ม 23" := "ยา 517", "ปึ่ม 24" := "ยา 518", "ปึ่ม 25" := "ยา 519", "ปึ่ม 26" := "ยา 520", "เมื่ิอมีการกดปุ้ม" => "Outputเมื่อมีการกดปุ่ม 20")
      Contact( "Outputเมื่อมีการกดปุ่ม 20" )
      S_SR(operand := "SR Step Motro 1,2  เบิกจ่าย 20", r1 := wire#w21)
      "button start"(Output => "Output ปุ่มยืนยันหน้า Screen")
      Contact( "Output ปุ่มยืนยันหน้า Screen" )
   END_RUNG wire#w2
   RUNG wire#powerrail
      Contact( "Output ทำงานเสด M1,2 forword No.20" )
   END_RUNG wire#w21
   RUNG wire#powerrail
      Contact( "ปุ่มClear" )
   END_RUNG wire#w21
   // the same network as SCL:
   "ตัวเลือกยา (26)"("ปึ่ม 1" := "ยา 1",
                     "ปึ่ม 2" := "ยา 2",
                     "ปึ่ม 3" := "ยา 3",
                     "ปึ่ม 4" := "ยา 4",
                     "ปึ่ม 5" := "ยา 5",
                     "ปึ่ม 6" := "ยา 6",
                     "ปึ่ม 7" := "ยา 7",
                     "ปึ่ม 8" := "ยา 8",
                     "ปึ่ม 9" := "ยา 9",
                     "ปึ่ม 10" := "ยา 10",
                     "ปึ่ม 11" := "ยา 11",
                     "ปึ่ม 12" := "ยา 12",
                     "ปึ่ม 13" := "ยา 13",
                     "ปึ่ม 14" := "ยา 14",
                     "ปึ่ม 15" := "ยา 15",
                     "ปึ่ม 16" := "ยา 16",
                     "ปึ่ม 17" := "ยา 17",
                     "ปึ่ม 18" := "ยา 18",
                     "ปึ่ม 19" := "ยา 19",
                     "ปึ่ม 20" := "ยา 20",
                     "ปึ่ม 21" := "ยา 21",
                     "ปึ่ม 22" := "ยา 22",
                     "ปึ่ม 23" := "ยา 23",
                     "ปึ่ม 24" := "ยา 24",
                     "ปึ่ม 25" := "ยา 25",
                     "ปึ่ม 26" := "ยา 26",
                     "เมื่ิอมีการกดปุ้ม" => "Outputเมื่อมีการกดปุ่ม 1",
                     ENO => #_w1);
   IF #_w1 AND "Outputเมื่อมีการกดปุ่ม 1" THEN
       "SR Step Motro 1,2  เบิกจ่าย 1" := TRUE;   // SR flip-flop
   END_IF;
   IF "Output ทำงานเสด M1,2 forword No.1" OR "ปุ่มClear" THEN
       "SR Step Motro 1,2  เบิกจ่าย 1" := FALSE;
   END_IF;
   "button start"(EN := "SR Step Motro 1,2  เบิกจ่าย 1", Output => "Output ปุ่มยืนยันหน้า Screen", ENO => #_w2);
   #_w4 := #_w2 AND "Output ปุ่มยืนยันหน้า Screen";
   "ตัวเลือกยา (26)"("ปึ่ม 1" := "ยา 27",
                     "ปึ่ม 2" := "ยา 28",
                     "ปึ่ม 3" := "ยา 29",
                     "ปึ่ม 4" := "ยา 30",
                     "ปึ่ม 5" := "ยา 31",
                     "ปึ่ม 6" := "ยา 32",
                     "ปึ่ม 7" := "ยา 33",
                     "ปึ่ม 8" := "ยา 34",
                     "ปึ่ม 9" := "ยา 35",
                     "ปึ่ม 10" := "ยา 36",
                     "ปึ่ม 11" := "ยา 37",
                     "ปึ่ม 12" := "ยา 38",
                     "ปึ่ม 13" := "ยา 39",
                     "ปึ่ม 14" := "ยา 40",
                     "ปึ่ม 15" := "ยา 41",
                     "ปึ่ม 16" := "ยา 42",
                     "ปึ่ม 17" := "ยา 43",
                     "ปึ่ม 18" := "ยา 44",
                     "ปึ่ม 19" := "ยา 45",
                     "ปึ่ม 20" := "ยา 46",
                     "ปึ่ม 21" := "ยา 47",
                     "ปึ่ม 22" := "ยา 48",
                     "ปึ่ม 23" := "ยา 49",
                     "ปึ่ม 24" := "ยา 50",
                     "ปึ่ม 25" := "ยา 51",
                     "ปึ่ม 26" := "ยา 52",
                     "เมื่ิอมีการกดปุ้ม" => "Outputเมื่อมีการกดปุ่ม 2",
                     ENO => #_w3);
   IF #_w3 AND "Outputเมื่อมีการกดปุ่ม 2" THEN
       "SR Step Motro 1,2  เบิกจ่าย 2" := TRUE;   // SR flip-flop
   END_IF;
   IF "Output ทำงานเสด M1,2 forword No.2" OR "ปุ่มClear" THEN
       "SR Step Motro 1,2  เบิกจ่าย 2" := FALSE;
   END_IF;
   "button start"(EN := "SR Step Motro 1,2  เบิกจ่าย 2", Output => "Output ปุ่มยืนยันหน้า Screen", ENO => #_w5);
   #_w7 := #_w5 AND "Output ปุ่มยืนยันหน้า Screen";
   "ตัวเลือกยา (26)"("ปึ่ม 1" := "ยา 53",
                     "ปึ่ม 2" := "ยา 54",
                     "ปึ่ม 3" := "ยา 55",
                     "ปึ่ม 4" := "ยา 56",
                     "ปึ่ม 5" := "ยา 57",
                     "ปึ่ม 6" := "ยา 58",
                     "ปึ่ม 7" := "ยา 59",
                     "ปึ่ม 8" := "ยา 60",
                     "ปึ่ม 9" := "ยา 61",
                     "ปึ่ม 10" := "ยา 62",
                     "ปึ่ม 11" := "ยา 63",
                     "ปึ่ม 12" := "ยา 64",
                     "ปึ่ม 13" := "ยา 65",
                     "ปึ่ม 14" := "ยา 66",
                     "ปึ่ม 15" := "ยา 67",
                     "ปึ่ม 16" := "ยา 68",
                     "ปึ่ม 17" := "ยา 69",
                     "ปึ่ม 18" := "ยา 70",
                     "ปึ่ม 19" := "ยา 71",
                     "ปึ่ม 20" := "ยา 72",
                     "ปึ่ม 21" := "ยา 73",
                     "ปึ่ม 22" := "ยา 74",
                     "ปึ่ม 23" := "ยา 75",
                     "ปึ่ม 24" := "ยา 76",
                     "ปึ่ม 25" := "ยา 77",
                     "ปึ่ม 26" := "ยา 78",
                     "เมื่ิอมีการกดปุ้ม" => "Outputเมื่อมีการกดปุ่ม 3",
                     ENO => #_w6);
   IF #_w6 AND "Outputเมื่อมีการกดปุ่ม 3" THEN
       "SR Step Motro 1,2  เบิกจ่าย 3" := TRUE;   // SR flip-flop
   END_IF;
   IF "Output ทำงานเสด M1,2 forword No.3" OR "ปุ่มClear" THEN
       "SR Step Motro 1,2  เบิกจ่าย 3" := FALSE;
   END_IF;
   "button start"(EN := "SR Step Motro 1,2  เบิกจ่าย 3", Output => "Output ปุ่มยืนยันหน้า Screen", ENO => #_w8);
   #_w10 := #_w8 AND "Output ปุ่มยืนยันหน้า Screen";
   "ตัวเลือกยา (26)"("ปึ่ม 1" := "ยา 79",
                     "ปึ่ม 2" := "ยา 80",
                     "ปึ่ม 3" := "ยา 81",
                     "ปึ่ม 4" := "ยา 82",
                     "ปึ่ม 5" := "ยา 83",
                     "ปึ่ม 6" := "ยา 84",
                     "ปึ่ม 7" := "ยา 85",
                     "ปึ่ม 8" := "ยา 86",
                     "ปึ่ม 9" := "ยา 87",
                     "ปึ่ม 10" := "ยา 88",
                     "ปึ่ม 11" := "ยา 89",
                     "ปึ่ม 12" := "ยา 90",
                     "ปึ่ม 13" := "ยา 91",
                     "ปึ่ม 14" := "ยา 92",
                     "ปึ่ม 15" := "ยา 93",
                     "ปึ่ม 16" := "ยา 94",
                     "ปึ่ม 17" := "ยา 95",
                     "ปึ่ม 18" := "ยา 96",
                     "ปึ่ม 19" := "ยา 97",
                     "ปึ่ม 20" := "ยา 98",
                     "ปึ่ม 21" := "ยา 99",
                     "ปึ่ม 22" := "ยา 100",
                     "ปึ่ม 23" := "ยา 101",
                     "ปึ่ม 24" := "ยา 102",
                     "ปึ่ม 25" := "ยา 103",
                     "ปึ่ม 26" := "ยา 104",
                     "เมื่ิอมีการกดปุ้ม" => "Outputเมื่อมีการกดปุ่ม 4",
                     ENO => #_w9);
   IF #_w9 AND "Outputเมื่อมีการกดปุ่ม 4" THEN
       "SR Step Motro 1,2  เบิกจ่าย 4" := TRUE;   // SR flip-flop
   END_IF;
   IF "Output ทำงานเสด M1,2 forword No.4" OR "ปุ่มClear" THEN
       "SR Step Motro 1,2  เบิกจ่าย 4" := FALSE;
   END_IF;
   "button start"(EN := "SR Step Motro 1,2  เบิกจ่าย 4", Output => "Output ปุ่มยืนยันหน้า Screen", ENO => #_w11);
   #_w13 := #_w11 AND "Output ปุ่มยืนยันหน้า Screen";
   "ตัวเลือกยา (26)"("ปึ่ม 1" := "ยา 105",
                     "ปึ่ม 2" := "ยา 106",
                     "ปึ่ม 3" := "ยา 107",
                     "ปึ่ม 4" := "ยา 108",
                     "ปึ่ม 5" := "ยา 109",
                     "ปึ่ม 6" := "ยา 110",
                     "ปึ่ม 7" := "ยา 111",
                     "ปึ่ม 8" := "ยา 112",
                     "ปึ่ม 9" := "ยา 113",
                     "ปึ่ม 10" := "ยา 114",
                     "ปึ่ม 11" := "ยา 115",
                     "ปึ่ม 12" := "ยา 116",
                     "ปึ่ม 13" := "ยา 117",
                     "ปึ่ม 14" := "ยา 118",
                     "ปึ่ม 15" := "ยา 119",
                     "ปึ่ม 16" := "ยา 120",
                     "ปึ่ม 17" := "ยา 121",
                     "ปึ่ม 18" := "ยา 122",
                     "ปึ่ม 19" := "ยา 123",
                     "ปึ่ม 20" := "ยา 124",
                     "ปึ่ม 21" := "ยา 125",
                     "ปึ่ม 22" := "ยา 126",
                     "ปึ่ม 23" := "ยา 127",
                     "ปึ่ม 24" := "ยา 128",
                     "ปึ่ม 25" := "ยา 129",
                     "ปึ่ม 26" := "ยา 130",
                     "เมื่ิอมีการกดปุ้ม" => "Outputเมื่อมีการกดปุ่ม 5",
                     ENO => #_w12);
   IF #_w12 AND "Outputเมื่อมีการกดปุ่ม 5" THEN
       "SR Step Motro 1,2  เบิกจ่าย 5" := TRUE;   // SR flip-flop
   END_IF;
   IF "Output ทำงานเสด M1,2 forword No.5" OR "ปุ่มClear" THEN
       "SR Step Motro 1,2  เบิกจ่าย 5" := FALSE;
   END_IF;
   "button start"(EN := "SR Step Motro 1,2  เบิกจ่าย 5", Output => "Output ปุ่มยืนยันหน้า Screen", ENO => #_w14);
   #_w16 := #_w14 AND "Output ปุ่มยืนยันหน้า Screen";
   "ตัวเลือกยา (26)"("ปึ่ม 1" := "ยา 131",
                     "ปึ่ม 2" := "ยา 132",
                     "ปึ่ม 3" := "ยา 133",
                     "ปึ่ม 4" := "ยา 134",
                     "ปึ่ม 5" := "ยา 135",
                     "ปึ่ม 6" := "ยา 136",
                     "ปึ่ม 7" := "ยา 137",
                     "ปึ่ม 8" := "ยา 138",
                     "ปึ่ม 9" := "ยา 139",
                     "ปึ่ม 10" := "ยา 140",
                     "ปึ่ม 11" := "ยา 141",
                     "ปึ่ม 12" := "ยา 142",
                     "ปึ่ม 13" := "ยา 143",
                     "ปึ่ม 14" := "ยา 144",
                     "ปึ่ม 15" := "ยา 145",
                     "ปึ่ม 16" := "ยา 146",
                     "ปึ่ม 17" := "ยา 147",
                     "ปึ่ม 18" := "ยา 148",
                     "ปึ่ม 19" := "ยา 149",
                     "ปึ่ม 20" := "ยา 150",
                     "ปึ่ม 21" := "ยา 151",
                     "ปึ่ม 22" := "ยา 152",
                     "ปึ่ม 23" := "ยา 153",
                     "ปึ่ม 24" := "ยา 154",
                     "ปึ่ม 25" := "ยา 155",
                     "ปึ่ม 26" := "ยา 156",
                     "เมื่ิอมีการกดปุ้ม" => "Outputเมื่อมีการกดปุ่ม 6",
                     ENO => #_w15);
   IF #_w15 AND "Outputเมื่อมีการกดปุ่ม 6" THEN
       "SR Step Motro 1,2  เบิกจ่าย 6" := TRUE;   // SR flip-flop
   END_IF;
   IF "Output ทำงานเสด M1,2 forword No.6" OR "ปุ่มClear" THEN
       "SR Step Motro 1,2  เบิกจ่าย 6" := FALSE;
   END_IF;
   "button start"(EN := "SR Step Motro 1,2  เบิกจ่าย 6", Output => "Output ปุ่มยืนยันหน้า Screen", ENO => #_w17);
   #_w19 := #_w17 AND "Output ปุ่มยืนยันหน้า Screen";
   "ตัวเลือกยา (26)"("ปึ่ม 1" := "ยา 157",
                     "ปึ่ม 2" := "ยา 158",
                     "ปึ่ม 3" := "ยา 159",
                     "ปึ่ม 4" := "ยา 160",
                     "ปึ่ม 5" := "ยา 161",
                     "ปึ่ม 6" := "ยา 162",
                     "ปึ่ม 7" := "ยา 163",
                     "ปึ่ม 8" := "ยา 164",
                     "ปึ่ม 9" := "ยา 165",
                     "ปึ่ม 10" := "ยา 166",
                     "ปึ่ม 11" := "ยา 167",
                     "ปึ่ม 12" := "ยา 168",
                     "ปึ่ม 13" := "ยา 169",
                     "ปึ่ม 14" := "ยา 170",
                     "ปึ่ม 15" := "ยา 171",
                     "ปึ่ม 16" := "ยา 172",
                     "ปึ่ม 17" := "ยา 173",
                     "ปึ่ม 18" := "ยา 174",
                     "ปึ่ม 19" := "ยา 175",
                     "ปึ่ม 20" := "ยา 176",
                     "ปึ่ม 21" := "ยา 177",
                     "ปึ่ม 22" := "ยา 178",
                     "ปึ่ม 23" := "ยา 179",
                     "ปึ่ม 24" := "ยา 180",
                     "ปึ่ม 25" := "ยา 181",
                     "ปึ่ม 26" := "ยา 182",
                     "เมื่ิอมีการกดปุ้ม" => "Outputเมื่อมีการกดปุ่ม 7",
                     ENO => #_w18);
   IF #_w18 AND "Outputเมื่อมีการกดปุ่ม 7" THEN
       "SR Step Motro 1,2  เบิกจ่าย 7" := TRUE;   // SR flip-flop
   END_IF;
   IF "Output ทำงานเสด M1,2 forword No.7" OR "ปุ่มClear" THEN
       "SR Step Motro 1,2  เบิกจ่าย 7" := FALSE;
   END_IF;
   "button start"(EN := "SR Step Motro 1,2  เบิกจ่าย 7", Output => "Output ปุ่มยืนยันหน้า Screen", ENO => #_w20);
   #_w22 := #_w20 AND "Output ปุ่มยืนยันหน้า Screen";
   "ตัวเลือกยา (26)"("ปึ่ม 1" := "ยา 183",
                     "ปึ่ม 2" := "ยา 184",
                     "ปึ่ม 3" := "ยา 185",
                     "ปึ่ม 4" := "ยา 186",
                     "ปึ่ม 5" := "ยา 187",
                     "ปึ่ม 6" := "ยา 188",
                     "ปึ่ม 7" := "ยา 189",
                     "ปึ่ม 8" := "ยา 190",
                     "ปึ่ม 9" := "ยา 191",
                     "ปึ่ม 10" := "ยา 192",
                     "ปึ่ม 11" := "ยา 193",
                     "ปึ่ม 12" := "ยา 194",
                     "ปึ่ม 13" := "ยา 195",
                     "ปึ่ม 14" := "ยา 196",
                     "ปึ่ม 15" := "ยา 197",
                     "ปึ่ม 16" := "ยา 198",
                     "ปึ่ม 17" := "ยา 199",
                     "ปึ่ม 18" := "ยา 200",
                     "ปึ่ม 19" := "ยา 201",
                     "ปึ่ม 20" := "ยา 202",
                     "ปึ่ม 21" := "ยา 203",
                     "ปึ่ม 22" := "ยา 204",
                     "ปึ่ม 23" := "ยา 205",
                     "ปึ่ม 24" := "ยา 206",
                     "ปึ่ม 25" := "ยา 207",
                     "ปึ่ม 26" := "ยา 208",
                     "เมื่ิอมีการกดปุ้ม" => "Outputเมื่อมีการกดปุ่ม 8",
                     ENO => #_w21);
   IF #_w21 AND "Outputเมื่อมีการกดปุ่ม 8" THEN
       "SR Step Motro 1,2  เบิกจ่าย 8" := TRUE;   // SR flip-flop
   END_IF;
   IF "Output ทำงานเสด M1,2 forword No.8" OR "ปุ่มClear" THEN
       "SR Step Motro 1,2  เบิกจ่าย 8" := FALSE;
   END_IF;
   "button start"(EN := "SR Step Motro 1,2  เบิกจ่าย 8", Output => "Output ปุ่มยืนยันหน้า Screen", ENO => #_w23);
   #_w25 := #_w23 AND "Output ปุ่มยืนยันหน้า Screen";
   "ตัวเลือกยา (26)"("ปึ่ม 1" := "ยา 209",
                     "ปึ่ม 2" := "ยา 210",
                     "ปึ่ม 3" := "ยา 211",
                     "ปึ่ม 4" := "ยา 212",
                     "ปึ่ม 5" := "ยา 213",
                     "ปึ่ม 6" := "ยา 214",
                     "ปึ่ม 7" := "ยา 215",
                     "ปึ่ม 8" := "ยา 216",
                     "ปึ่ม 9" := "ยา 217",
                     "ปึ่ม 10" := "ยา 218",
                     "ปึ่ม 11" := "ยา 219",
                     "ปึ่ม 12" := "ยา 220",
                     "ปึ่ม 13" := "ยา 221",
                     "ปึ่ม 14" := "ยา 222",
                     "ปึ่ม 15" := "ยา 223",
                     "ปึ่ม 16" := "ยา 224",
                     "ปึ่ม 17" := "ยา 225",
                     "ปึ่ม 18" := "ยา 226",
                     "ปึ่ม 19" := "ยา 227",
                     "ปึ่ม 20" := "ยา 228",
                     "ปึ่ม 21" := "ยา 229",
                     "ปึ่ม 22" := "ยา 230",
                     "ปึ่ม 23" := "ยา 231",
                     "ปึ่ม 24" := "ยา 232",
                     "ปึ่ม 25" := "ยา 233",
                     "ปึ่ม 26" := "ยา 234",
                     "เมื่ิอมีการกดปุ้ม" => "Outputเมื่อมีการกดปุ่ม 9",
                     ENO => #_w24);
   IF #_w24 AND "Outputเมื่อมีการกดปุ่ม 9" THEN
       "SR Step Motro 1,2  เบิกจ่าย 9" := TRUE;   // SR flip-flop
   END_IF;
   IF "Output ทำงานเสด M1,2 forword No.9" OR "ปุ่มClear" THEN
       "SR Step Motro 1,2  เบิกจ่าย 9" := FALSE;
   END_IF;
   "button start"(EN := "SR Step Motro 1,2  เบิกจ่าย 9", Output => "Output ปุ่มยืนยันหน้า Screen", ENO => #_w26);
   #_w28 := #_w26 AND "Output ปุ่มยืนยันหน้า Screen";
   "ตัวเลือกยา (26)"("ปึ่ม 1" := "ยา 235",
                     "ปึ่ม 2" := "ยา 236",
                     "ปึ่ม 3" := "ยา 234",
                     "ปึ่ม 4" := "ยา 238",
                     "ปึ่ม 5" := "ยา 239",
                     "ปึ่ม 6" := "ยา 240",
                     "ปึ่ม 7" := "ยา 241",
                     "ปึ่ม 8" := "ยา 242",
                     "ปึ่ม 9" := "ยา 243",
                     "ปึ่ม 10" := "ยา 244",
                     "ปึ่ม 11" := "ยา 245",
                     "ปึ่ม 12" := "ยา 246",
                     "ปึ่ม 13" := "ยา 247",
                     "ปึ่ม 14" := "ยา 248",
                     "ปึ่ม 15" := "ยา 249",
                     "ปึ่ม 16" := "ยา 250",
                     "ปึ่ม 17" := "ยา 251",
                     "ปึ่ม 18" := "ยา 252",
                     "ปึ่ม 19" := "ยา 253",
                     "ปึ่ม 20" := "ยา 254",
                     "ปึ่ม 21" := "ยา 255",
                     "ปึ่ม 22" := "ยา 256",
                     "ปึ่ม 23" := "ยา 257",
                     "ปึ่ม 24" := "ยา 258",
                     "ปึ่ม 25" := "ยา 259",
                     "ปึ่ม 26" := "ยา 260",
                     "เมื่ิอมีการกดปุ้ม" => "Outputเมื่อมีการกดปุ่ม 10",
                     ENO => #_w27);
   IF #_w27 AND "Outputเมื่อมีการกดปุ่ม 10" THEN
       "SR Step Motro 1,2  เบิกจ่าย 10" := TRUE;   // SR flip-flop
   END_IF;
   IF "Output ทำงานเสด M1,2 forword No.10" OR "ปุ่มClear" THEN
       "SR Step Motro 1,2  เบิกจ่าย 10" := FALSE;
   END_IF;
   "button start"(EN := "SR Step Motro 1,2  เบิกจ่าย 10",
                  Output => "Output ปุ่มยืนยันหน้า Screen",
                  ENO => #_w29);
   #_w31 := #_w29 AND "Output ปุ่มยืนยันหน้า Screen";
   "ตัวเลือกยา (26)"("ปึ่ม 1" := "ยา 261",
                     "ปึ่ม 2" := "ยา 262",
                     "ปึ่ม 3" := "ยา 263",
                     "ปึ่ม 4" := "ยา 264",
                     "ปึ่ม 5" := "ยา 265",
                     "ปึ่ม 6" := "ยา 266",
                     "ปึ่ม 7" := "ยา 267",
                     "ปึ่ม 8" := "ยา 268",
                     "ปึ่ม 9" := "ยา 269",
                     "ปึ่ม 10" := "ยา 270",
                     "ปึ่ม 11" := "ยา 271",
                     "ปึ่ม 12" := "ยา 272",
                     "ปึ่ม 13" := "ยา 273",
                     "ปึ่ม 14" := "ยา 274",
                     "ปึ่ม 15" := "ยา 275",
                     "ปึ่ม 16" := "ยา 276",
                     "ปึ่ม 17" := "ยา 277",
                     "ปึ่ม 18" := "ยา 278",
                     "ปึ่ม 19" := "ยา 279",
                     "ปึ่ม 20" := "ยา 280",
                     "ปึ่ม 21" := "ยา 281",
                     "ปึ่ม 22" := "ยา 282",
                     "ปึ่ม 23" := "ยา 283",
                     "ปึ่ม 24" := "ยา 284",
                     "ปึ่ม 25" := "ยา 285",
                     "ปึ่ม 26" := "ยา 286",
                     "เมื่ิอมีการกดปุ้ม" => "Outputเมื่อมีการกดปุ่ม 11",
                     ENO => #_w30);
   IF #_w30 AND "Outputเมื่อมีการกดปุ่ม 11" THEN
       "SR Step Motro 1,2  เบิกจ่าย 11" := TRUE;   // SR flip-flop
   END_IF;
   IF "Output ทำงานเสด M1,2 forword No.11" OR "ปุ่มClear" THEN
       "SR Step Motro 1,2  เบิกจ่าย 11" := FALSE;
   END_IF;
   "button start"(EN := "SR Step Motro 1,2  เบิกจ่าย 11",
                  Output => "Output ปุ่มยืนยันหน้า Screen",
                  ENO => #_w32);
   #_w34 := #_w32 AND "Output ปุ่มยืนยันหน้า Screen";
   "ตัวเลือกยา (26)"("ปึ่ม 1" := "ยา 287",
                     "ปึ่ม 2" := "ยา 288",
                     "ปึ่ม 3" := "ยา 289",
                     "ปึ่ม 4" := "ยา 290",
                     "ปึ่ม 5" := "ยา 291",
                     "ปึ่ม 6" := "ยา 292",
                     "ปึ่ม 7" := "ยา 293",
                     "ปึ่ม 8" := "ยา 294",
                     "ปึ่ม 9" := "ยา 295",
                     "ปึ่ม 10" := "ยา 296",
                     "ปึ่ม 11" := "ยา 297",
                     "ปึ่ม 12" := "ยา 298",
                     "ปึ่ม 13" := "ยา 299",
                     "ปึ่ม 14" := "ยา 300",
                     "ปึ่ม 15" := "ยา 301",
                     "ปึ่ม 16" := "ยา 302",
                     "ปึ่ม 17" := "ยา 303",
                     "ปึ่ม 18" := "ยา 304",
                     "ปึ่ม 19" := "ยา 305",
                     "ปึ่ม 20" := "ยา 306",
                     "ปึ่ม 21" := "ยา 307",
                     "ปึ่ม 22" := "ยา 308",
                     "ปึ่ม 23" := "ยา 309",
                     "ปึ่ม 24" := "ยา 310",
                     "ปึ่ม 25" := "ยา 311",
                     "ปึ่ม 26" := "ยา 312",
                     "เมื่ิอมีการกดปุ้ม" => "Outputเมื่อมีการกดปุ่ม 12",
                     ENO => #_w33);
   IF #_w33 AND "Outputเมื่อมีการกดปุ่ม 12" THEN
       "SR Step Motro 1,2  เบิกจ่าย 12" := TRUE;   // SR flip-flop
   END_IF;
   IF "Output ทำงานเสด M1,2 forword No.12" OR "ปุ่มClear" THEN
       "SR Step Motro 1,2  เบิกจ่าย 12" := FALSE;
   END_IF;
   "button start"(EN := "SR Step Motro 1,2  เบิกจ่าย 12",
                  Output => "Output ปุ่มยืนยันหน้า Screen",
                  ENO => #_w35);
   #_w37 := #_w35 AND "Output ปุ่มยืนยันหน้า Screen";
   "ตัวเลือกยา (26)"("ปึ่ม 1" := "ยา 313",
                     "ปึ่ม 2" := "ยา 314",
                     "ปึ่ม 3" := "ยา 315",
                     "ปึ่ม 4" := "ยา 316",
                     "ปึ่ม 5" := "ยา 317",
                     "ปึ่ม 6" := "ยา 318",
                     "ปึ่ม 7" := "ยา 319",
                     "ปึ่ม 8" := "ยา 320",
                     "ปึ่ม 9" := "ยา 321",
                     "ปึ่ม 10" := "ยา 322",
                     "ปึ่ม 11" := "ยา 323",
                     "ปึ่ม 12" := "ยา 324",
                     "ปึ่ม 13" := "ยา 325",
                     "ปึ่ม 14" := "ยา 326",
                     "ปึ่ม 15" := "ยา 327",
                     "ปึ่ม 16" := "ยา 328",
                     "ปึ่ม 17" := "ยา 329",
                     "ปึ่ม 18" := "ยา 330",
                     "ปึ่ม 19" := "ยา 331",
                     "ปึ่ม 20" := "ยา 332",
                     "ปึ่ม 21" := "ยา 333",
                     "ปึ่ม 22" := "ยา 334",
                     "ปึ่ม 23" := "ยา 335",
                     "ปึ่ม 24" := "ยา 336",
                     "ปึ่ม 25" := "ยา 337",
                     "ปึ่ม 26" := "ยา 338",
                     "เมื่ิอมีการกดปุ้ม" => "Outputเมื่อมีการกดปุ่ม 13",
                     ENO => #_w36);
   IF #_w36 AND "Outputเมื่อมีการกดปุ่ม 13" THEN
       "SR Step Motro 1,2  เบิกจ่าย 13" := TRUE;   // SR flip-flop
   END_IF;
   IF "Output ทำงานเสด M1,2 forword No.13" OR "ปุ่มClear" THEN
       "SR Step Motro 1,2  เบิกจ่าย 13" := FALSE;
   END_IF;
   "button start"(EN := "SR Step Motro 1,2  เบิกจ่าย 13",
                  Output => "Output ปุ่มยืนยันหน้า Screen",
                  ENO => #_w38);
   #_w40 := #_w38 AND "Output ปุ่มยืนยันหน้า Screen";
   "ตัวเลือกยา (26)"("ปึ่ม 1" := "ยา 339",
                     "ปึ่ม 2" := "ยา 340",
                     "ปึ่ม 3" := "ยา 341",
                     "ปึ่ม 4" := "ยา 342",
                     "ปึ่ม 5" := "ยา 343",
                     "ปึ่ม 6" := "ยา 344",
                     "ปึ่ม 7" := "ยา 345",
                     "ปึ่ม 8" := "ยา 345",
                     "ปึ่ม 9" := "ยา 347",
                     "ปึ่ม 10" := "ยา 348",
                     "ปึ่ม 11" := "ยา 349",
                     "ปึ่ม 12" := "ยา 350",
                     "ปึ่ม 13" := "ยา 351",
                     "ปึ่ม 14" := "ยา 352",
                     "ปึ่ม 15" := "ยา 353",
                     "ปึ่ม 16" := "ยา 354",
                     "ปึ่ม 17" := "ยา 355",
                     "ปึ่ม 18" := "ยา 356",
                     "ปึ่ม 19" := "ยา 357",
                     "ปึ่ม 20" := "ยา 358",
                     "ปึ่ม 21" := "ยา 359",
                     "ปึ่ม 22" := "ยา 360",
                     "ปึ่ม 23" := "ยา 361",
                     "ปึ่ม 24" := "ยา 362",
                     "ปึ่ม 25" := "ยา 363",
                     "ปึ่ม 26" := "ยา 364",
                     "เมื่ิอมีการกดปุ้ม" => "Outputเมื่อมีการกดปุ่ม 14",
                     ENO => #_w39);
   IF #_w39 AND "Outputเมื่อมีการกดปุ่ม 14" THEN
       "SR Step Motro 1,2  เบิกจ่าย 14" := TRUE;   // SR flip-flop
   END_IF;
   IF "Output ทำงานเสด M1,2 forword No.14" OR "ปุ่มClear" THEN
       "SR Step Motro 1,2  เบิกจ่าย 14" := FALSE;
   END_IF;
   "button start"(EN := "SR Step Motro 1,2  เบิกจ่าย 14",
                  Output => "Output ปุ่มยืนยันหน้า Screen",
                  ENO => #_w41);
   #_w43 := #_w41 AND "Output ปุ่มยืนยันหน้า Screen";
   "ตัวเลือกยา (26)"("ปึ่ม 1" := "ยา 365",
                     "ปึ่ม 2" := "ยา 365",
                     "ปึ่ม 3" := "ยา 367",
                     "ปึ่ม 4" := "ยา 368",
                     "ปึ่ม 5" := "ยา 369",
                     "ปึ่ม 6" := "ยา 370",
                     "ปึ่ม 7" := "ยา 371",
                     "ปึ่ม 8" := "ยา 372",
                     "ปึ่ม 9" := "ยา 373",
                     "ปึ่ม 10" := "ยา 374",
                     "ปึ่ม 11" := "ยา 375",
                     "ปึ่ม 12" := "ยา 376",
                     "ปึ่ม 13" := "ยา 377",
                     "ปึ่ม 14" := "ยา 378",
                     "ปึ่ม 15" := "ยา 379",
                     "ปึ่ม 16" := "ยา 380",
                     "ปึ่ม 17" := "ยา 381",
                     "ปึ่ม 18" := "ยา 382",
                     "ปึ่ม 19" := "ยา 383",
                     "ปึ่ม 20" := "ยา 384",
                     "ปึ่ม 21" := "ยา 385",
                     "ปึ่ม 22" := "ยา 386",
                     "ปึ่ม 23" := "ยา 387",
                     "ปึ่ม 24" := "ยา 388",
                     "ปึ่ม 25" := "ยา 389",
                     "ปึ่ม 26" := "ยา 390",
                     "เมื่ิอมีการกดปุ้ม" => "Outputเมื่อมีการกดปุ่ม 15",
                     ENO => #_w42);
   IF #_w42 AND "Outputเมื่อมีการกดปุ่ม 15" THEN
       "SR Step Motro 1,2  เบิกจ่าย 15" := TRUE;   // SR flip-flop
   END_IF;
   IF "Output ทำงานเสด M1,2 forword No.15" OR "ปุ่มClear" THEN
       "SR Step Motro 1,2  เบิกจ่าย 15" := FALSE;
   END_IF;
   "button start"(EN := "SR Step Motro 1,2  เบิกจ่าย 15",
                  Output => "Output ปุ่มยืนยันหน้า Screen",
                  ENO => #_w44);
   #_w46 := #_w44 AND "Output ปุ่มยืนยันหน้า Screen";
   "ตัวเลือกยา (26)"("ปึ่ม 1" := "ยา 391",
                     "ปึ่ม 2" := "ยา 392",
                     "ปึ่ม 3" := "ยา 393",
                     "ปึ่ม 4" := "ยา 394",
                     "ปึ่ม 5" := "ยา 395",
                     "ปึ่ม 6" := "ยา 396",
                     "ปึ่ม 7" := "ยา 397",
                     "ปึ่ม 8" := "ยา 398",
                     "ปึ่ม 9" := "ยา 399",
                     "ปึ่ม 10" := "ยา 400",
                     "ปึ่ม 11" := "ยา 401",
                     "ปึ่ม 12" := "ยา 402",
                     "ปึ่ม 13" := "ยา 403",
                     "ปึ่ม 14" := "ยา 404",
                     "ปึ่ม 15" := "ยา 405",
                     "ปึ่ม 16" := "ยา 406",
                     "ปึ่ม 17" := "ยา 407",
                     "ปึ่ม 18" := "ยา 408",
                     "ปึ่ม 19" := "ยา 409",
                     "ปึ่ม 20" := "ยา 410",
                     "ปึ่ม 21" := "ยา 411",
                     "ปึ่ม 22" := "ยา 412",
                     "ปึ่ม 23" := "ยา 413",
                     "ปึ่ม 24" := "ยา 414",
                     "ปึ่ม 25" := "ยา 415",
                     "ปึ่ม 26" := "ยา 416",
                     "เมื่ิอมีการกดปุ้ม" => "Outputเมื่อมีการกดปุ่ม 16",
                     ENO => #_w45);
   IF #_w45 AND "Outputเมื่อมีการกดปุ่ม 16" THEN
       "SR Step Motro 1,2  เบิกจ่าย 16" := TRUE;   // SR flip-flop
   END_IF;
   IF "Output ทำงานเสด M1,2 forword No.16" OR "ปุ่มClear" THEN
       "SR Step Motro 1,2  เบิกจ่าย 16" := FALSE;
   END_IF;
   "button start"(EN := "SR Step Motro 1,2  เบิกจ่าย 16",
                  Output => "Output ปุ่มยืนยันหน้า Screen",
                  ENO => #_w47);
   #_w49 := #_w47 AND "Output ปุ่มยืนยันหน้า Screen";
   "ตัวเลือกยา (26)"("ปึ่ม 1" := "ยา 417",
                     "ปึ่ม 2" := "ยา 418",
                     "ปึ่ม 3" := "ยา 419",
                     "ปึ่ม 4" := "ยา 420",
                     "ปึ่ม 5" := "ยา 421",
                     "ปึ่ม 6" := "ยา 422",
                     "ปึ่ม 7" := "ยา 423",
                     "ปึ่ม 8" := "ยา 424",
                     "ปึ่ม 9" := "ยา 425",
                     "ปึ่ม 10" := "ยา 426",
                     "ปึ่ม 11" := "ยา 427",
                     "ปึ่ม 12" := "ยา 428",
                     "ปึ่ม 13" := "ยา 429",
                     "ปึ่ม 14" := "ยา 430",
                     "ปึ่ม 15" := "ยา 431",
                     "ปึ่ม 16" := "ยา 432",
                     "ปึ่ม 17" := "ยา 433",
                     "ปึ่ม 18" := "ยา 434",
                     "ปึ่ม 19" := "ยา 435",
                     "ปึ่ม 20" := "ยา 436",
                     "ปึ่ม 21" := "ยา 437",
                     "ปึ่ม 22" := "ยา 438",
                     "ปึ่ม 23" := "ยา 439",
                     "ปึ่ม 24" := "ยา 440",
                     "ปึ่ม 25" := "ยา 441",
                     "ปึ่ม 26" := "ยา 442",
                     "เมื่ิอมีการกดปุ้ม" => "Outputเมื่อมีการกดปุ่ม 17",
                     ENO => #_w48);
   IF #_w48 AND "Outputเมื่อมีการกดปุ่ม 17" THEN
       "SR Step Motro 1,2  เบิกจ่าย 17" := TRUE;   // SR flip-flop
   END_IF;
   IF "Output ทำงานเสด M1,2 forword No.17" OR "ปุ่มClear" THEN
       "SR Step Motro 1,2  เบิกจ่าย 17" := FALSE;
   END_IF;
   "button start"(EN := "SR Step Motro 1,2  เบิกจ่าย 17",
                  Output => "Output ปุ่มยืนยันหน้า Screen",
                  ENO => #_w50);
   #_w52 := #_w50 AND "Output ปุ่มยืนยันหน้า Screen";
   "ตัวเลือกยา (26)"("ปึ่ม 1" := "ยา 443",
                     "ปึ่ม 2" := "ยา 444",
                     "ปึ่ม 3" := "ยา 445",
                     "ปึ่ม 4" := "ยา 446",
                     "ปึ่ม 5" := "ยา 447",
                     "ปึ่ม 6" := "ยา 448",
                     "ปึ่ม 7" := "ยา 449",
                     "ปึ่ม 8" := "ยา 450",
                     "ปึ่ม 9" := "ยา 451",
                     "ปึ่ม 10" := "ยา 452",
                     "ปึ่ม 11" := "ยา 453",
                     "ปึ่ม 12" := "ยา 454",
                     "ปึ่ม 13" := "ยา 455",
                     "ปึ่ม 14" := "ยา 456",
                     "ปึ่ม 15" := "ยา 457",
                     "ปึ่ม 16" := "ยา 458",
                     "ปึ่ม 17" := "ยา 459",
                     "ปึ่ม 18" := "ยา 460",
                     "ปึ่ม 19" := "ยา 461",
                     "ปึ่ม 20" := "ยา 462",
                     "ปึ่ม 21" := "ยา 463",
                     "ปึ่ม 22" := "ยา 464",
                     "ปึ่ม 23" := "ยา 465",
                     "ปึ่ม 24" := "ยา 466",
                     "ปึ่ม 25" := "ยา 467",
                     "ปึ่ม 26" := "ยา 468",
                     "เมื่ิอมีการกดปุ้ม" => "Outputเมื่อมีการกดปุ่ม 18",
                     ENO => #_w51);
   IF #_w51 AND "Outputเมื่อมีการกดปุ่ม 18" THEN
       "SR Step Motro 1,2  เบิกจ่าย 18" := TRUE;   // SR flip-flop
   END_IF;
   IF "Output ทำงานเสด M1,2 forword No.18" OR "ปุ่มClear" THEN
       "SR Step Motro 1,2  เบิกจ่าย 18" := FALSE;
   END_IF;
   "button start"(EN := "SR Step Motro 1,2  เบิกจ่าย 18",
                  Output => "Output ปุ่มยืนยันหน้า Screen",
                  ENO => #_w53);
   #_w55 := #_w53 AND "Output ปุ่มยืนยันหน้า Screen";
   "ตัวเลือกยา (26)"("ปึ่ม 1" := "ยา 469",
                     "ปึ่ม 2" := "ยา 470",
                     "ปึ่ม 3" := "ยา 471",
                     "ปึ่ม 4" := "ยา 472",
                     "ปึ่ม 5" := "ยา 473",
                     "ปึ่ม 6" := "ยา 474",
                     "ปึ่ม 7" := "ยา 475",
                     "ปึ่ม 8" := "ยา 476",
                     "ปึ่ม 9" := "ยา 477",
                     "ปึ่ม 10" := "ยา 478",
                     "ปึ่ม 11" := "ยา 479",
                     "ปึ่ม 12" := "ยา 480",
                     "ปึ่ม 13" := "ยา 481",
                     "ปึ่ม 14" := "ยา 482",
                     "ปึ่ม 15" := "ยา 483",
                     "ปึ่ม 16" := "ยา 484",
                     "ปึ่ม 17" := "ยา 485",
                     "ปึ่ม 18" := "ยา 486",
                     "ปึ่ม 19" := "ยา 487",
                     "ปึ่ม 20" := "ยา 488",
                     "ปึ่ม 21" := "ยา 489",
                     "ปึ่ม 22" := "ยา 490",
                     "ปึ่ม 23" := "ยา 491",
                     "ปึ่ม 24" := "ยา 492",
                     "ปึ่ม 25" := "ยา 493",
                     "ปึ่ม 26" := "ยา 494",
                     "เมื่ิอมีการกดปุ้ม" => "Outputเมื่อมีการกดปุ่ม 19",
                     ENO => #_w54);
   IF #_w54 AND "Outputเมื่อมีการกดปุ่ม 19" THEN
       "SR Step Motro 1,2  เบิกจ่าย 19" := TRUE;   // SR flip-flop
   END_IF;
   IF "Output ทำงานเสด M1,2 forword No.19" OR "ปุ่มClear" THEN
       "SR Step Motro 1,2  เบิกจ่าย 19" := FALSE;
   END_IF;
   "button start"(EN := "SR Step Motro 1,2  เบิกจ่าย 19",
                  Output => "Output ปุ่มยืนยันหน้า Screen",
                  ENO => #_w56);
   #_w58 := #_w56 AND "Output ปุ่มยืนยันหน้า Screen";
   "ตัวเลือกยา (26)"("ปึ่ม 1" := "ยา 495",
                     "ปึ่ม 2" := "ยา 496",
                     "ปึ่ม 3" := "ยา 497",
                     "ปึ่ม 4" := "ยา 498",
                     "ปึ่ม 5" := "ยา 499",
                     "ปึ่ม 6" := "ยา 500",
                     "ปึ่ม 7" := "ยา 501",
                     "ปึ่ม 8" := "ยา 502",
                     "ปึ่ม 9" := "ยา 503",
                     "ปึ่ม 10" := "ยา 504",
                     "ปึ่ม 11" := "ยา 505",
                     "ปึ่ม 12" := "ยา 505",
                     "ปึ่ม 13" := "ยา 507",
                     "ปึ่ม 14" := "ยา 508",
                     "ปึ่ม 15" := "ยา 509",
                     "ปึ่ม 16" := "ยา 510",
                     "ปึ่ม 17" := "ยา 511",
                     "ปึ่ม 18" := "ยา 512",
                     "ปึ่ม 19" := "ยา 513",
                     "ปึ่ม 20" := "ยา 514",
                     "ปึ่ม 21" := "ยา 515",
                     "ปึ่ม 22" := "ยา 516",
                     "ปึ่ม 23" := "ยา 517",
                     "ปึ่ม 24" := "ยา 518",
                     "ปึ่ม 25" := "ยา 519",
                     "ปึ่ม 26" := "ยา 520",
                     "เมื่ิอมีการกดปุ้ม" => "Outputเมื่อมีการกดปุ่ม 20",
                     ENO => #_w57);
   IF #_w57 AND "Outputเมื่อมีการกดปุ่ม 20" THEN
       "SR Step Motro 1,2  เบิกจ่าย 20" := TRUE;   // SR flip-flop
   END_IF;
   IF "Output ทำงานเสด M1,2 forword No.20" OR "ปุ่มClear" THEN
       "SR Step Motro 1,2  เบิกจ่าย 20" := FALSE;
   END_IF;
   "button start"(EN := "SR Step Motro 1,2  เบิกจ่าย 20",
                  Output => "Output ปุ่มยืนยันหน้า Screen",
                  ENO => #_w59);
   #"Stepper Motor  ทำงาน" := #_w4 OR #_w7 OR #_w10 OR #_w13 OR #_w16 OR #_w19 OR #_w22 OR #_w25 OR #_w28 OR #_w31 OR #_w34 OR #_w37 OR #_w40 OR #_w43 OR #_w46 OR #_w49 OR #_w52 OR #_w55 OR #_w58 OR (#_w59 AND "Output ปุ่มยืนยันหน้า Screen");
END_REGION

REGION Network 2
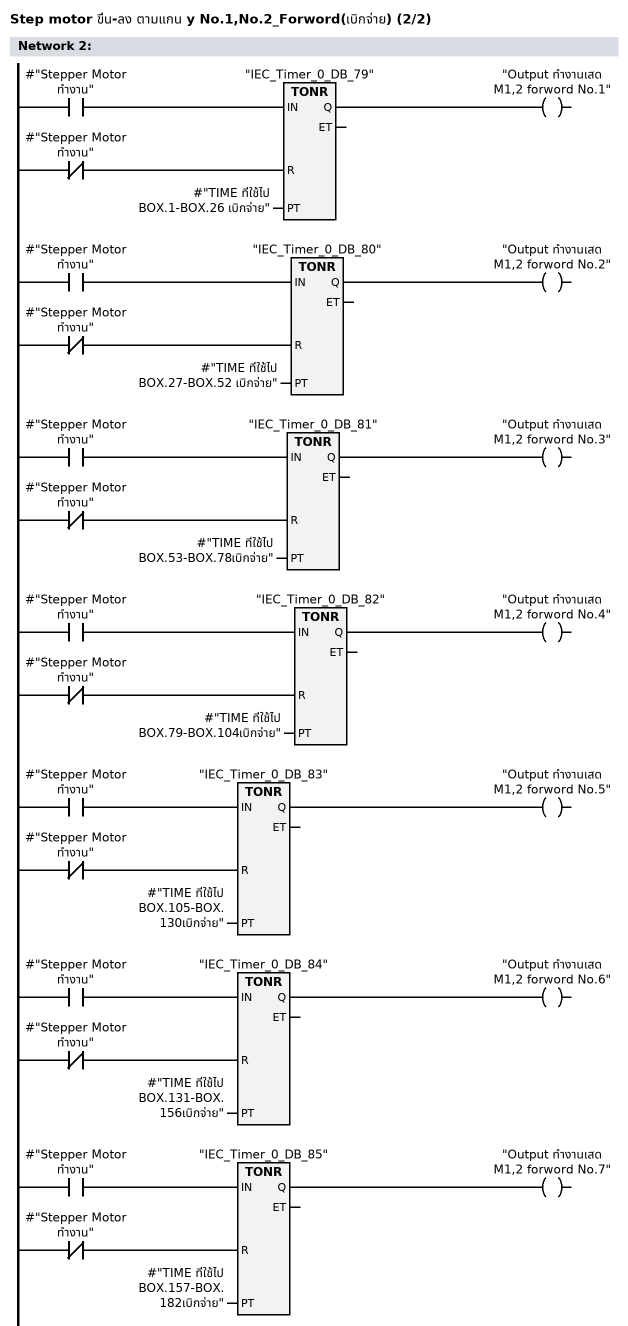
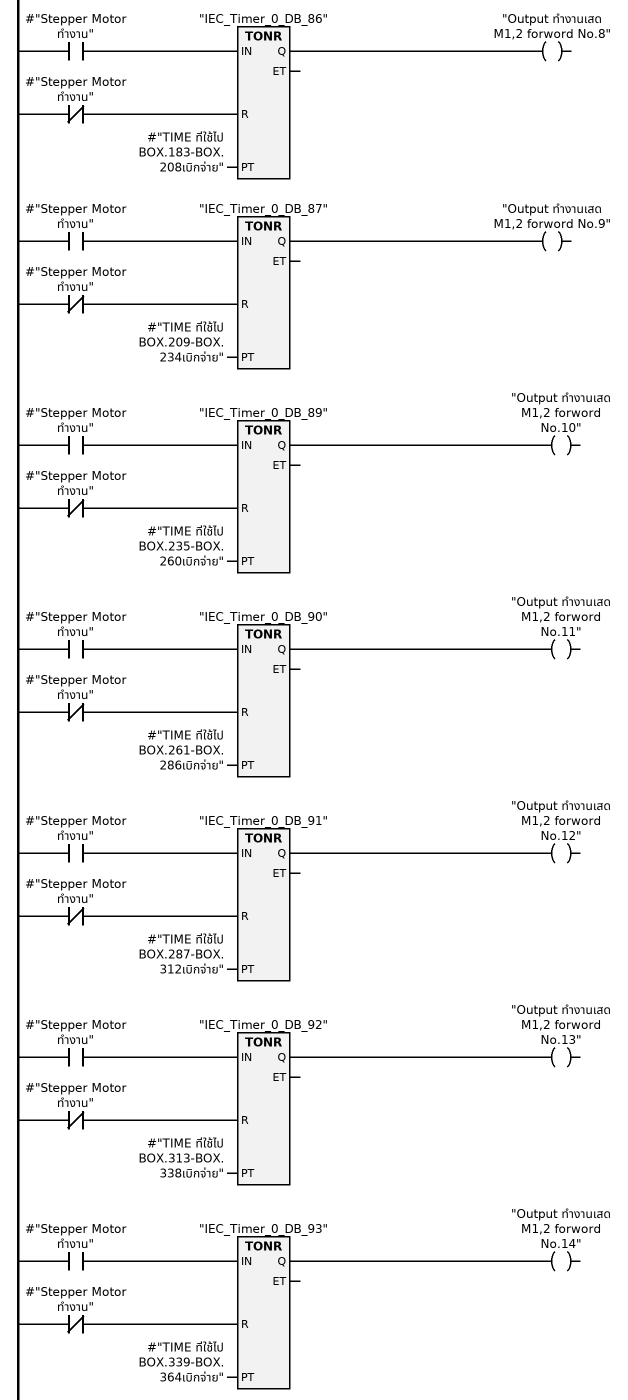
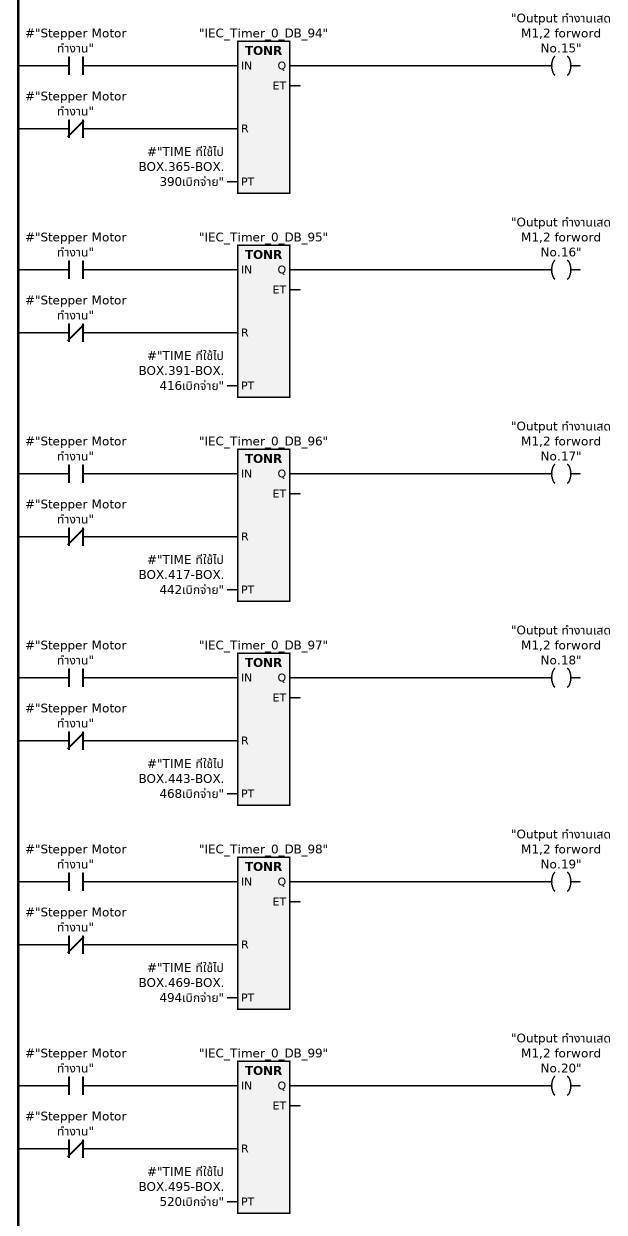
   "IEC_Timer_0_DB_79".TONR(IN := #"Stepper Motor  ทำงาน",
                           R := NOT #"Stepper Motor  ทำงาน",
                           PT := #"TIME ที่ใช้ไป BOX.1-BOX.26 เบิกจ่าย");
   "Output ทำงานเสด M1,2 forword No.1" := "IEC_Timer_0_DB_79".Q;
   "IEC_Timer_0_DB_80".TONR(IN := #"Stepper Motor  ทำงาน",
                           R := NOT #"Stepper Motor  ทำงาน",
                           PT := #"TIME ที่ใช้ไป BOX.27-BOX.52 เบิกจ่าย");
   "Output ทำงานเสด M1,2 forword No.2" := "IEC_Timer_0_DB_80".Q;
   "IEC_Timer_0_DB_81".TONR(IN := #"Stepper Motor  ทำงาน",
                           R := NOT #"Stepper Motor  ทำงาน",
                           PT := #"TIME ที่ใช้ไป BOX.53-BOX.78เบิกจ่าย");
   "Output ทำงานเสด M1,2 forword No.3" := "IEC_Timer_0_DB_81".Q;
   "IEC_Timer_0_DB_82".TONR(IN := #"Stepper Motor  ทำงาน",
                           R := NOT #"Stepper Motor  ทำงาน",
                           PT := #"TIME ที่ใช้ไป BOX.79-BOX.104เบิกจ่าย");
   "Output ทำงานเสด M1,2 forword No.4" := "IEC_Timer_0_DB_82".Q;
   "IEC_Timer_0_DB_83".TONR(IN := #"Stepper Motor  ทำงาน",
                           R := NOT #"Stepper Motor  ทำงาน",
                           PT := #"TIME ที่ใช้ไป BOX.105-BOX.130เบิกจ่าย");
   "Output ทำงานเสด M1,2 forword No.5" := "IEC_Timer_0_DB_83".Q;
   "IEC_Timer_0_DB_84".TONR(IN := #"Stepper Motor  ทำงาน",
                           R := NOT #"Stepper Motor  ทำงาน",
                           PT := #"TIME ที่ใช้ไป BOX.131-BOX.156เบิกจ่าย");
   "Output ทำงานเสด M1,2 forword No.6" := "IEC_Timer_0_DB_84".Q;
   "IEC_Timer_0_DB_85".TONR(IN := #"Stepper Motor  ทำงาน",
                           R := NOT #"Stepper Motor  ทำงาน",
                           PT := #"TIME ที่ใช้ไป BOX.157-BOX.182เบิกจ่าย");
   "Output ทำงานเสด M1,2 forword No.7" := "IEC_Timer_0_DB_85".Q;
   "IEC_Timer_0_DB_86".TONR(IN := #"Stepper Motor  ทำงาน",
                           R := NOT #"Stepper Motor  ทำงาน",
                           PT := #"TIME ที่ใช้ไป BOX.183-BOX.208เบิกจ่าย");
   "Output ทำงานเสด M1,2 forword No.8" := "IEC_Timer_0_DB_86".Q;
   "IEC_Timer_0_DB_87".TONR(IN := #"Stepper Motor  ทำงาน",
                           R := NOT #"Stepper Motor  ทำงาน",
                           PT := #"TIME ที่ใช้ไป BOX.209-BOX.234เบิกจ่าย");
   "Output ทำงานเสด M1,2 forword No.9" := "IEC_Timer_0_DB_87".Q;
   "IEC_Timer_0_DB_89".TONR(IN := #"Stepper Motor  ทำงาน",
                           R := NOT #"Stepper Motor  ทำงาน",
                           PT := #"TIME ที่ใช้ไป BOX.235-BOX.260เบิกจ่าย");
   "Output ทำงานเสด M1,2 forword No.10" := "IEC_Timer_0_DB_89".Q;
   "IEC_Timer_0_DB_90".TONR(IN := #"Stepper Motor  ทำงาน",
                           R := NOT #"Stepper Motor  ทำงาน",
                           PT := #"TIME ที่ใช้ไป BOX.261-BOX.286เบิกจ่าย");
   "Output ทำงานเสด M1,2 forword No.11" := "IEC_Timer_0_DB_90".Q;
   "IEC_Timer_0_DB_91".TONR(IN := #"Stepper Motor  ทำงาน",
                           R := NOT #"Stepper Motor  ทำงาน",
                           PT := #"TIME ที่ใช้ไป BOX.287-BOX.312เบิกจ่าย");
   "Output ทำงานเสด M1,2 forword No.12" := "IEC_Timer_0_DB_91".Q;
   "IEC_Timer_0_DB_92".TONR(IN := #"Stepper Motor  ทำงาน",
                           R := NOT #"Stepper Motor  ทำงาน",
                           PT := #"TIME ที่ใช้ไป BOX.313-BOX.338เบิกจ่าย");
   "Output ทำงานเสด M1,2 forword No.13" := "IEC_Timer_0_DB_92".Q;
   "IEC_Timer_0_DB_93".TONR(IN := #"Stepper Motor  ทำงาน",
                           R := NOT #"Stepper Motor  ทำงาน",
                           PT := #"TIME ที่ใช้ไป BOX.339-BOX.364เบิกจ่าย");
   "Output ทำงานเสด M1,2 forword No.14" := "IEC_Timer_0_DB_93".Q;
   "IEC_Timer_0_DB_94".TONR(IN := #"Stepper Motor  ทำงาน",
                           R := NOT #"Stepper Motor  ทำงาน",
                           PT := #"TIME ที่ใช้ไป BOX.365-BOX.390เบิกจ่าย");
   "Output ทำงานเสด M1,2 forword No.15" := "IEC_Timer_0_DB_94".Q;
   "IEC_Timer_0_DB_95".TONR(IN := #"Stepper Motor  ทำงาน",
                           R := NOT #"Stepper Motor  ทำงาน",
                           PT := #"TIME ที่ใช้ไป BOX.391-BOX.416เบิกจ่าย");
   "Output ทำงานเสด M1,2 forword No.16" := "IEC_Timer_0_DB_95".Q;
   "IEC_Timer_0_DB_96".TONR(IN := #"Stepper Motor  ทำงาน",
                           R := NOT #"Stepper Motor  ทำงาน",
                           PT := #"TIME ที่ใช้ไป BOX.417-BOX.442เบิกจ่าย");
   "Output ทำงานเสด M1,2 forword No.17" := "IEC_Timer_0_DB_96".Q;
   "IEC_Timer_0_DB_97".TONR(IN := #"Stepper Motor  ทำงาน",
                           R := NOT #"Stepper Motor  ทำงาน",
                           PT := #"TIME ที่ใช้ไป BOX.443-BOX.468เบิกจ่าย");
   "Output ทำงานเสด M1,2 forword No.18" := "IEC_Timer_0_DB_97".Q;
   "IEC_Timer_0_DB_98".TONR(IN := #"Stepper Motor  ทำงาน",
                           R := NOT #"Stepper Motor  ทำงาน",
                           PT := #"TIME ที่ใช้ไป BOX.469-BOX.494เบิกจ่าย");
   "Output ทำงานเสด M1,2 forword No.19" := "IEC_Timer_0_DB_98".Q;
   "IEC_Timer_0_DB_99".TONR(IN := #"Stepper Motor  ทำงาน",
                           R := NOT #"Stepper Motor  ทำงาน",
                           PT := #"TIME ที่ใช้ไป BOX.495-BOX.520เบิกจ่าย");
   "Output ทำงานเสด M1,2 forword No.20" := "IEC_Timer_0_DB_99".Q;
END_REGION
END_FUNCTION_BLOCK

FUNCTION_BLOCK "Step motor ขึ่น-ลง ตามแกน y No.1,No.2_Blackword(เบิกจ่าย)"   // FB7, LAD
{ S7_Optimized_Access := 'TRUE' }
VERSION : 0.1
   VAR_INPUT
      "TIME ที่ใช้ไป BOX.1-BOX.26" : Time;
      "TIME ที่ใช้ไป BOX.27-BOX.52" : Time;
      "TIME ที่ใช้ไป BOX.53-BOX.78" : Time;
      "TIME ที่ใช้ไป BOX.79-BOX.104" : Time;
      "TIME ที่ใช้ไป BOX.105-BOX.130" : Time;
      "TIME ที่ใช้ไป BOX.131-BOX.156" : Time;
      "TIME ที่ใช้ไป BOX.157-BOX.182" : Time;
      "TIME ที่ใช้ไป BOX.183-BOX.208" : Time;
      "TIME ที่ใช้ไป BOX.209-BOX.234" : Time;
      "TIME ที่ใช้ไป BOX.235-BOX.260" : Time;
      "TIME ที่ใช้ไป BOX.261-BOX.286" : Time;
      "TIME ที่ใช้ไป BOX.287-BOX.312" : Time;
      "TIME ที่ใช้ไป BOX.313-BOX.338" : Time;
      "TIME ที่ใช้ไป BOX.339-BOX.364" : Time;
      "TIME ที่ใช้ไป BOX.365-BOX.390" : Time;
      "TIME ที่ใช้ไป BOX.391-BOX.416" : Time;
      "TIME ที่ใช้ไป BOX.417-BOX.442" : Time;
      "TIME ที่ใช้ไป BOX.443-BOX.468" : Time;
      "TIME ที่ใช้ไป BOX.469-BOX.494" : Time;
      "TIME ที่ใช้ไป BOX.495-BOX.520" : Time;
   END_VAR
   VAR_IN_OUT
      "Stepper Motor  ทำงาน" : Bool;
   END_VAR
   VAR_TEMP   // added for the SCL form of the ladder/FBD networks
      _w1 : Bool;
      _w2 : Bool;
      _w3 : Bool;
      _w4 : Bool;
      _w5 : Bool;
      _w6 : Bool;
      _w7 : Bool;
      _w8 : Bool;
      _w9 : Bool;
      _w10 : Bool;
      _w11 : Bool;
      _w12 : Bool;
      _w13 : Bool;
      _w14 : Bool;
      _w15 : Bool;
      _w16 : Bool;
      _w17 : Bool;
      _w18 : Bool;
      _w19 : Bool;
      _w20 : Bool;
      _w21 : Bool;
      _w22 : Bool;
      _w23 : Bool;
      _w24 : Bool;
      _w25 : Bool;
      _w26 : Bool;
      _w27 : Bool;
      _w28 : Bool;
      _w29 : Bool;
      _w30 : Bool;
      _w31 : Bool;
      _w32 : Bool;
      _w33 : Bool;
      _w34 : Bool;
      _w35 : Bool;
      _w36 : Bool;
      _w37 : Bool;
      _w38 : Bool;
      _w39 : Bool;
      _w40 : Bool;
      _w41 : Bool;
      _w42 : Bool;
      _w43 : Bool;
      _w44 : Bool;
      _w45 : Bool;
      _w46 : Bool;
      _w47 : Bool;
      _w48 : Bool;
      _w49 : Bool;
      _w50 : Bool;
      _w51 : Bool;
      _w52 : Bool;
      _w53 : Bool;
      _w54 : Bool;
      _w55 : Bool;
      _w56 : Bool;
      _w57 : Bool;
      _w58 : Bool;
      _w59 : Bool;
   END_VAR
BEGIN

REGION Network 1
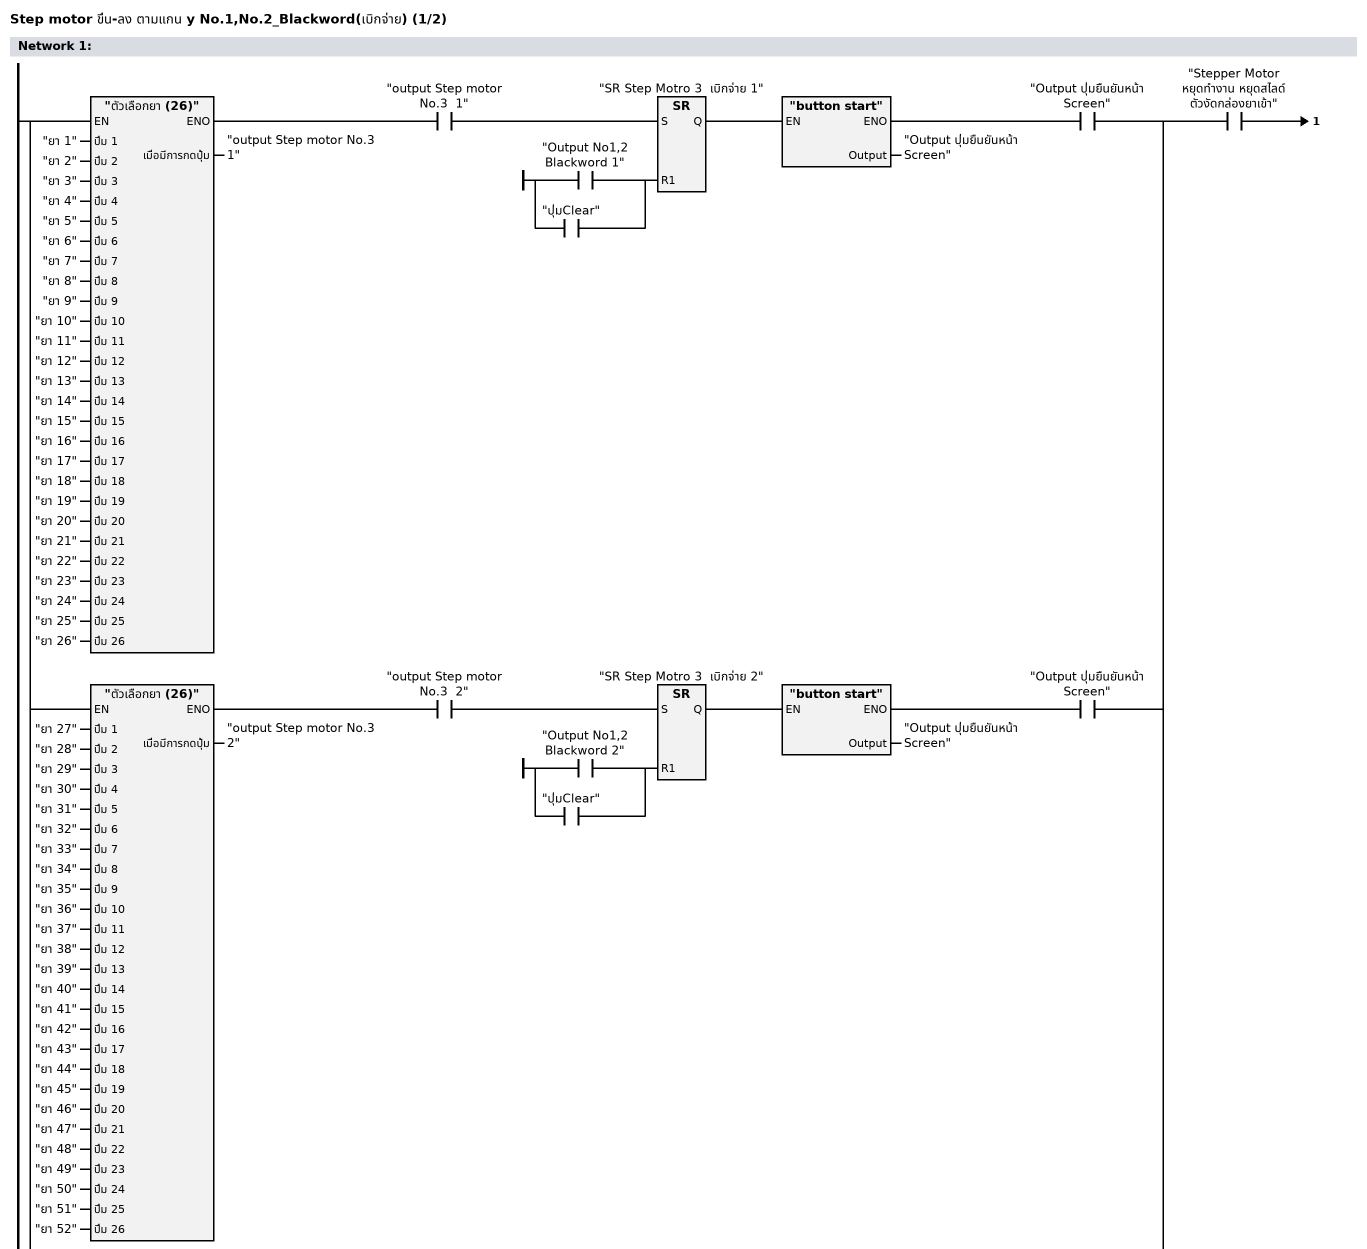
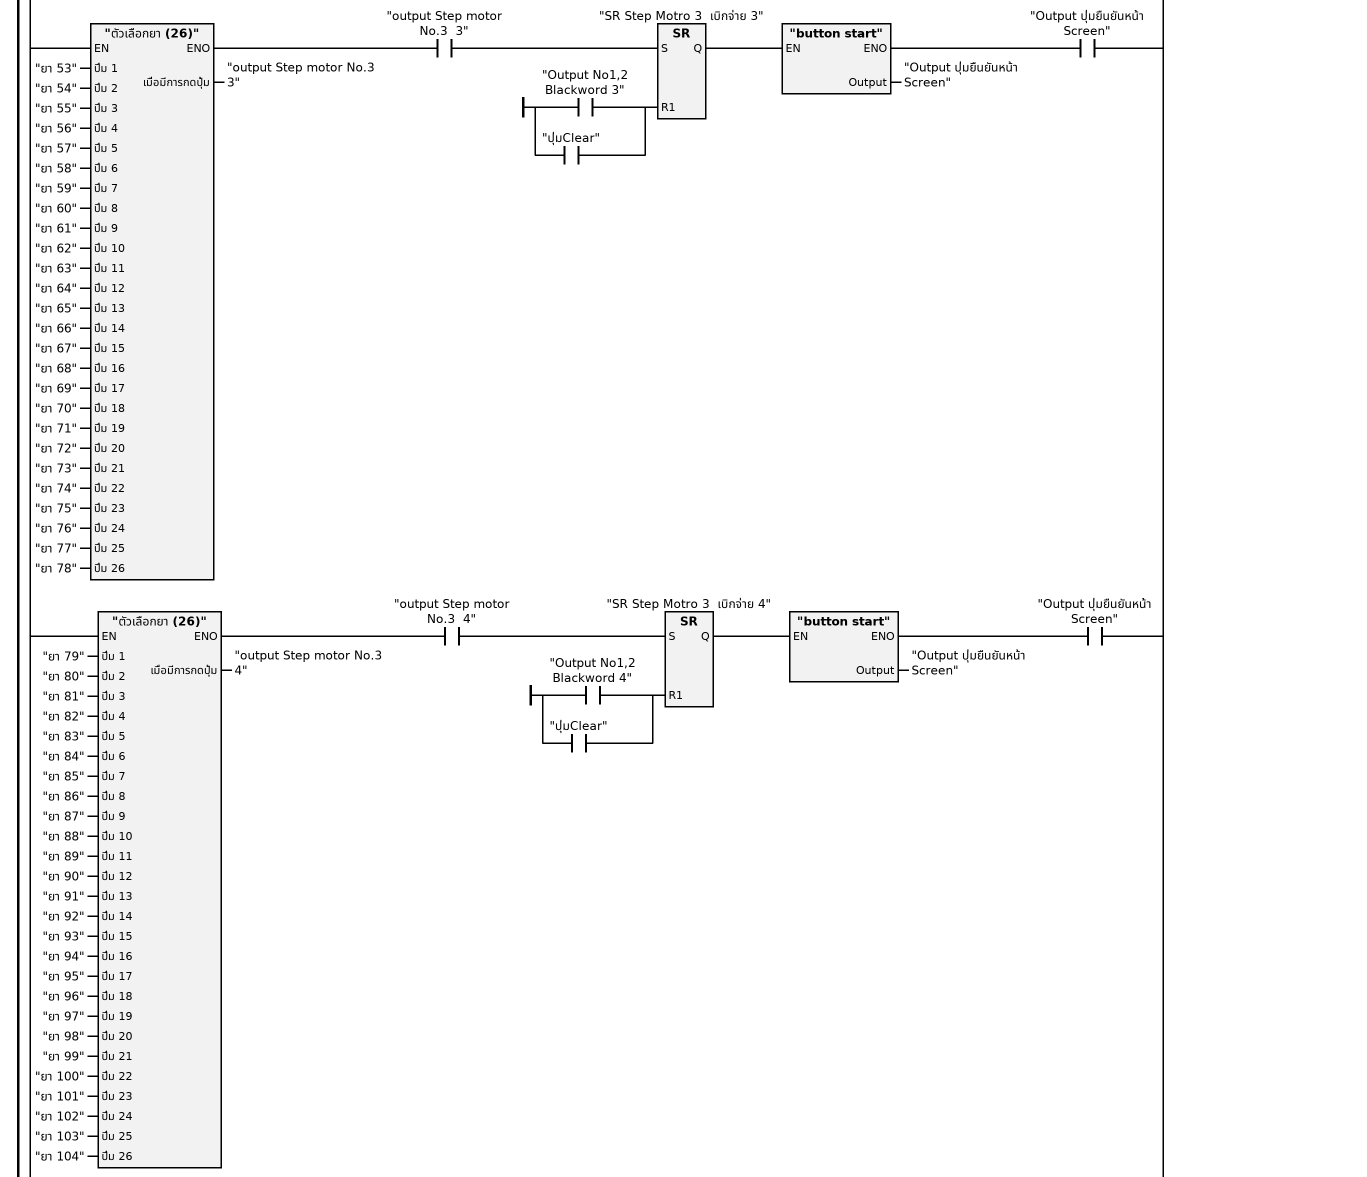
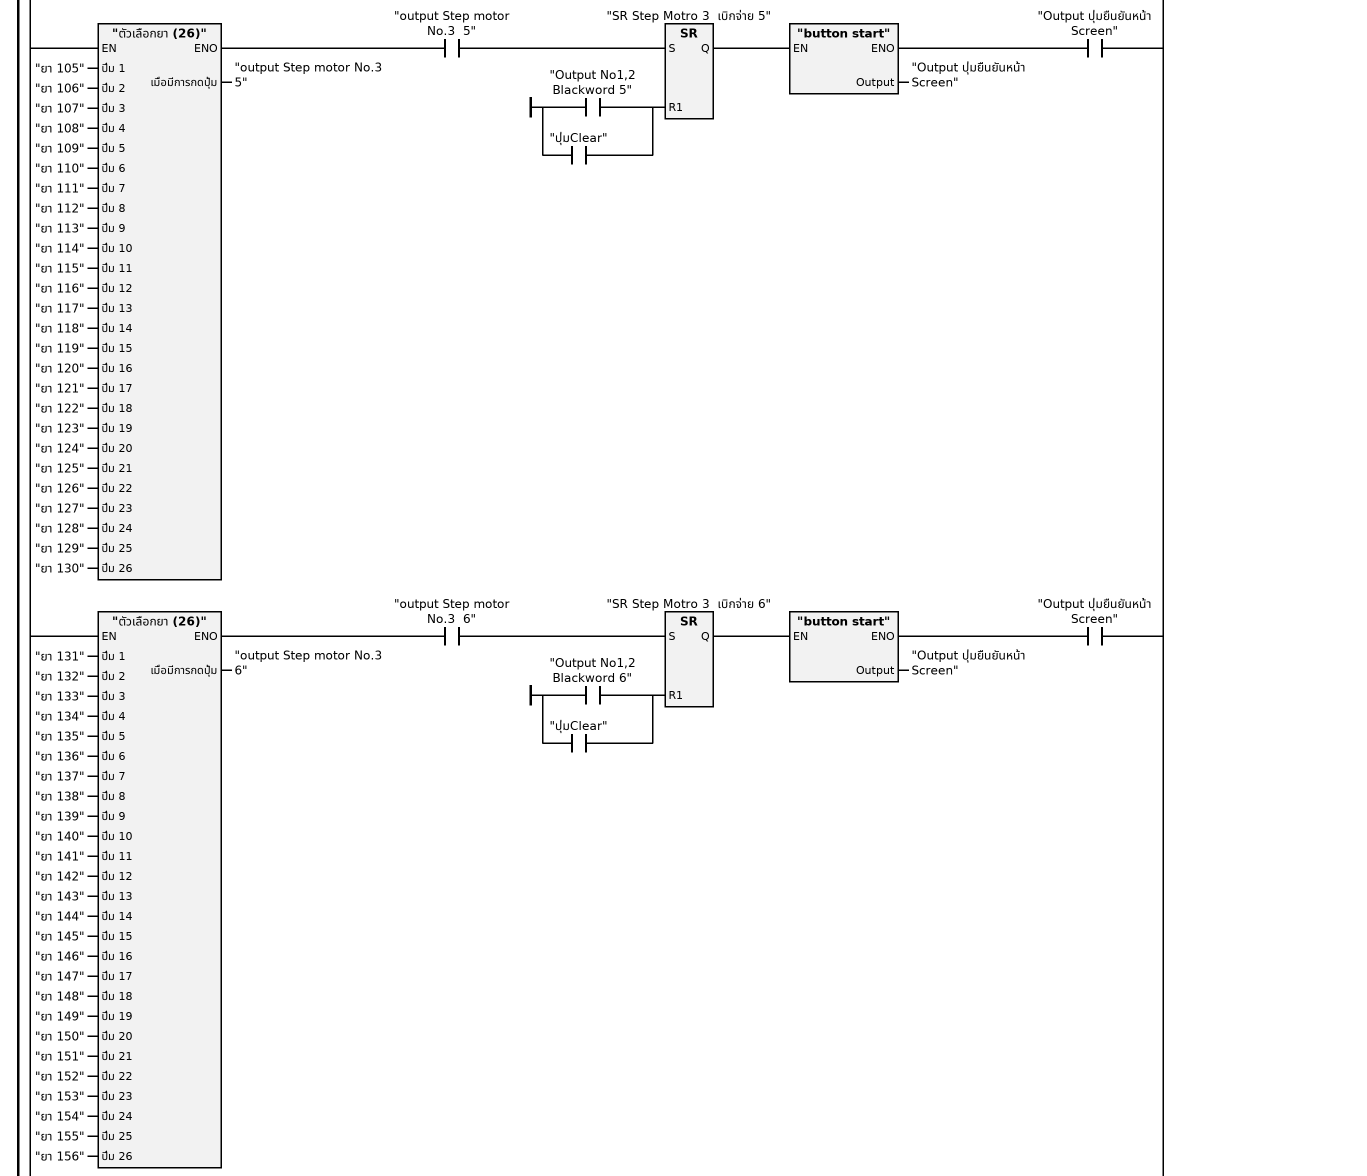
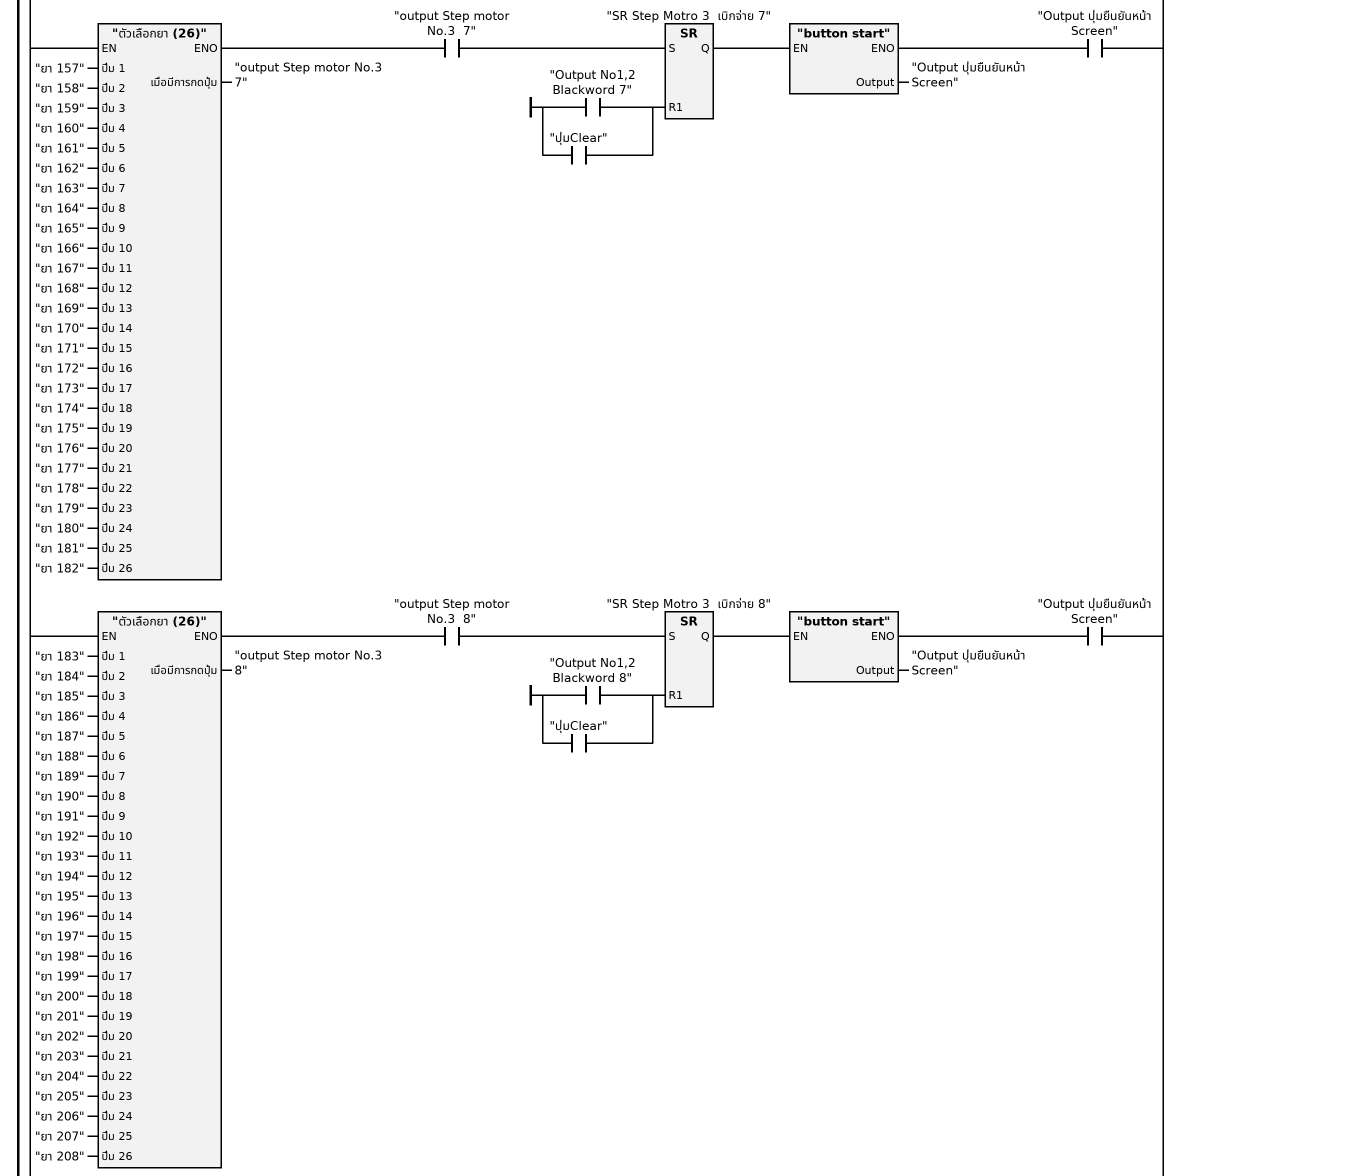
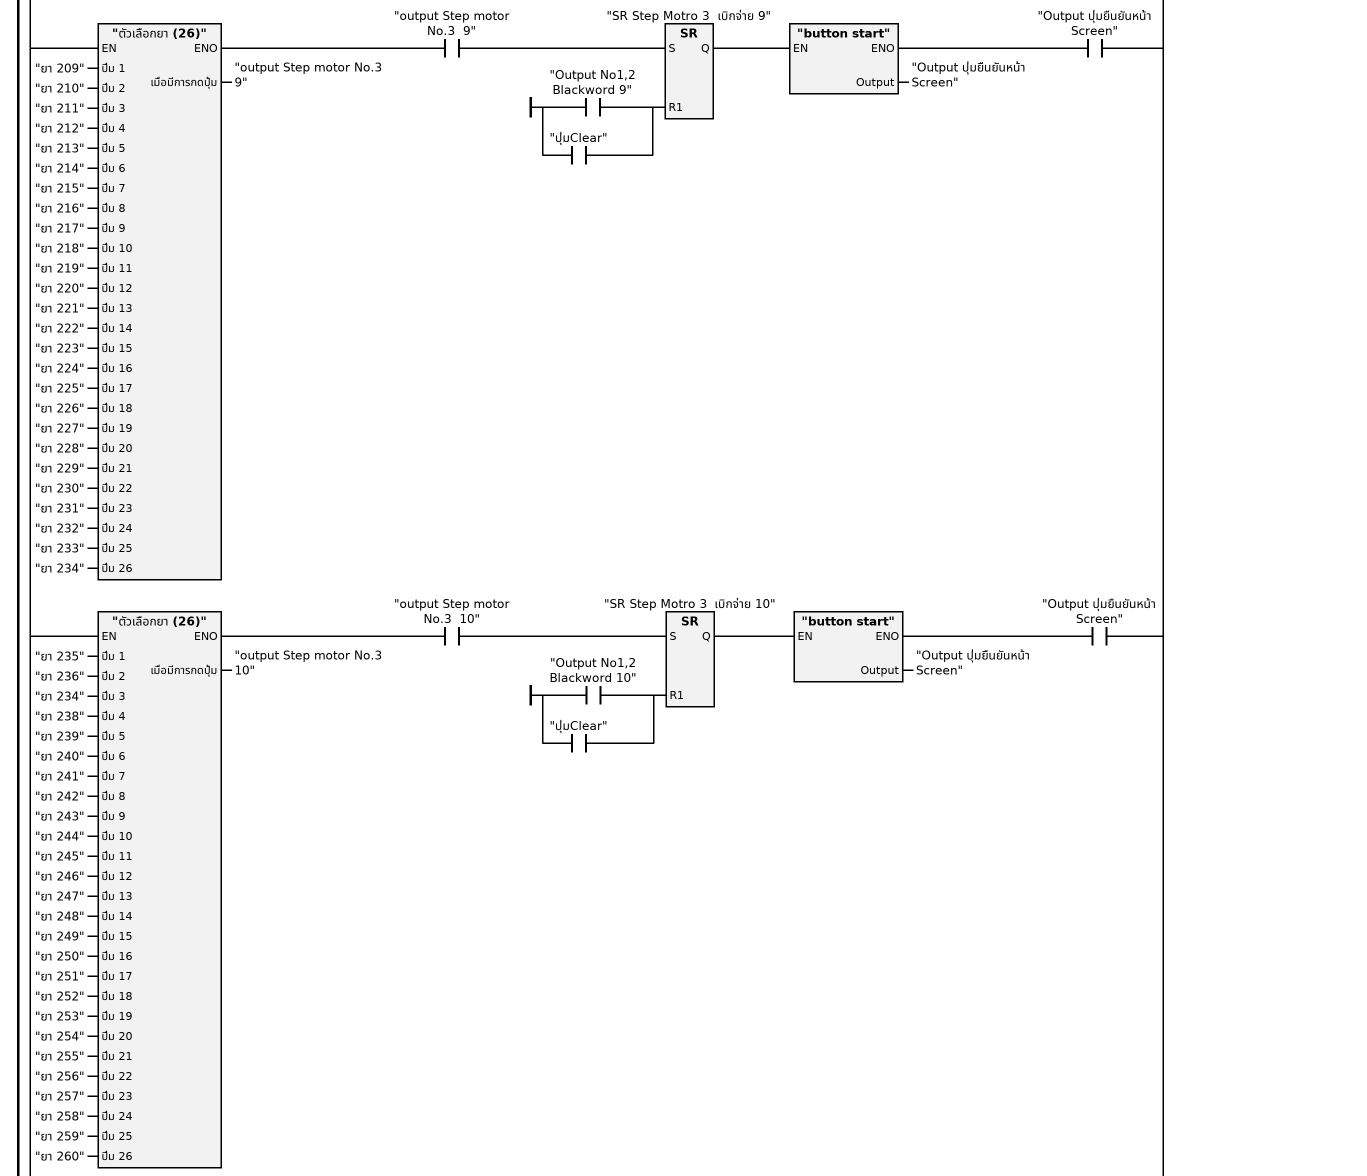
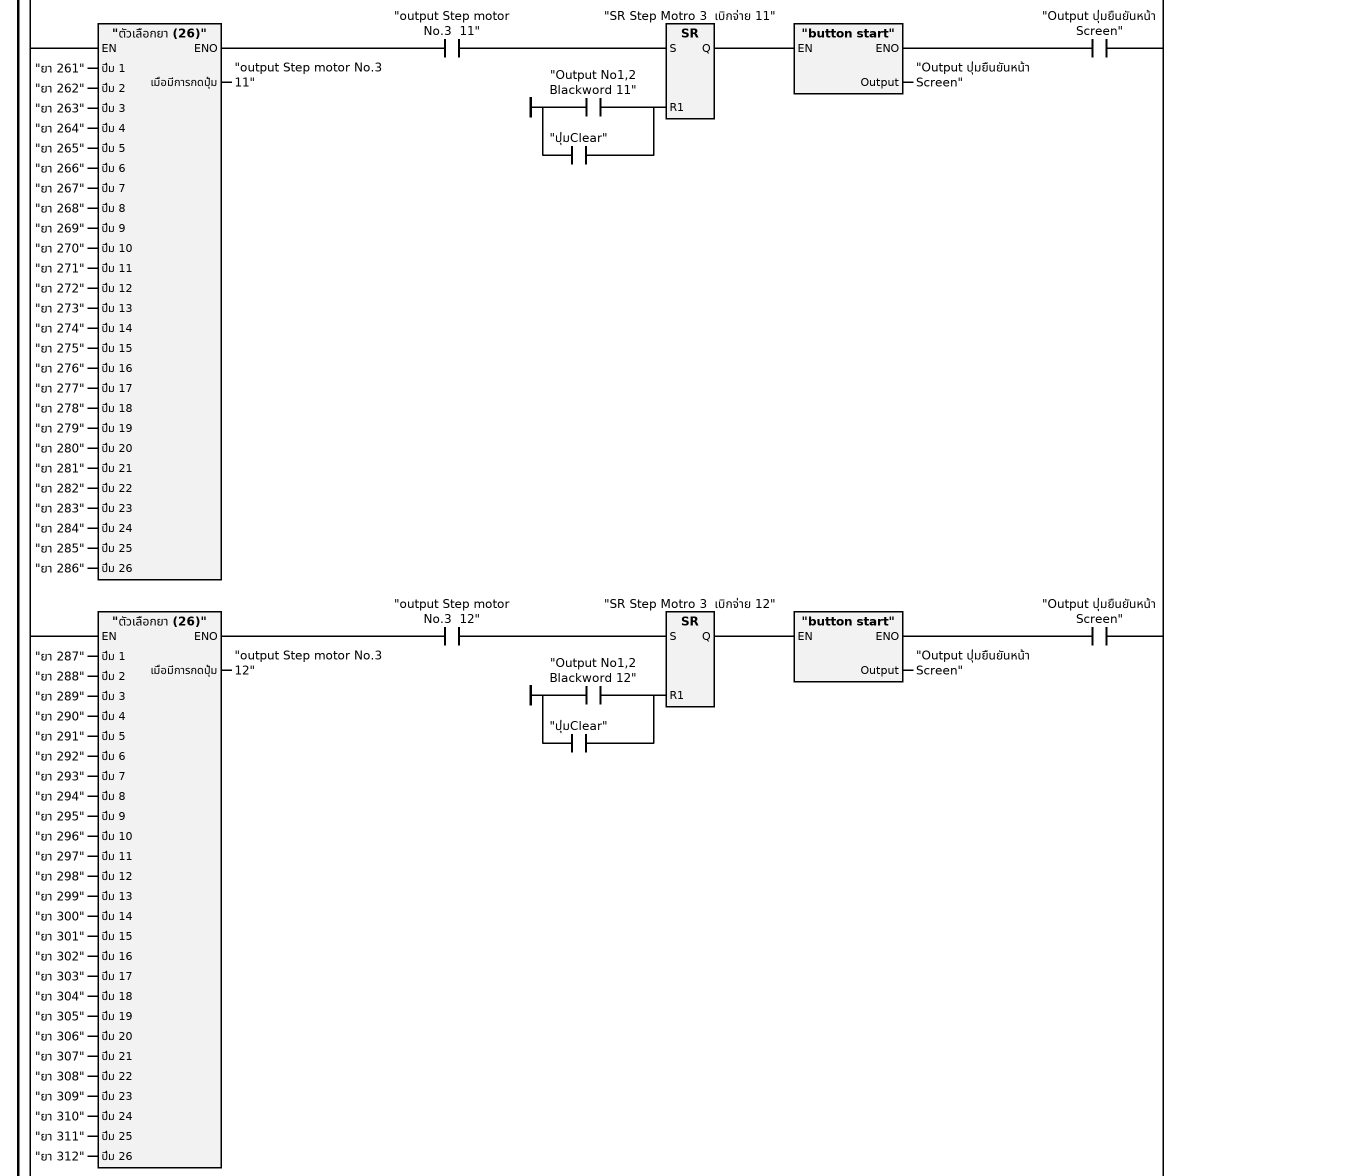
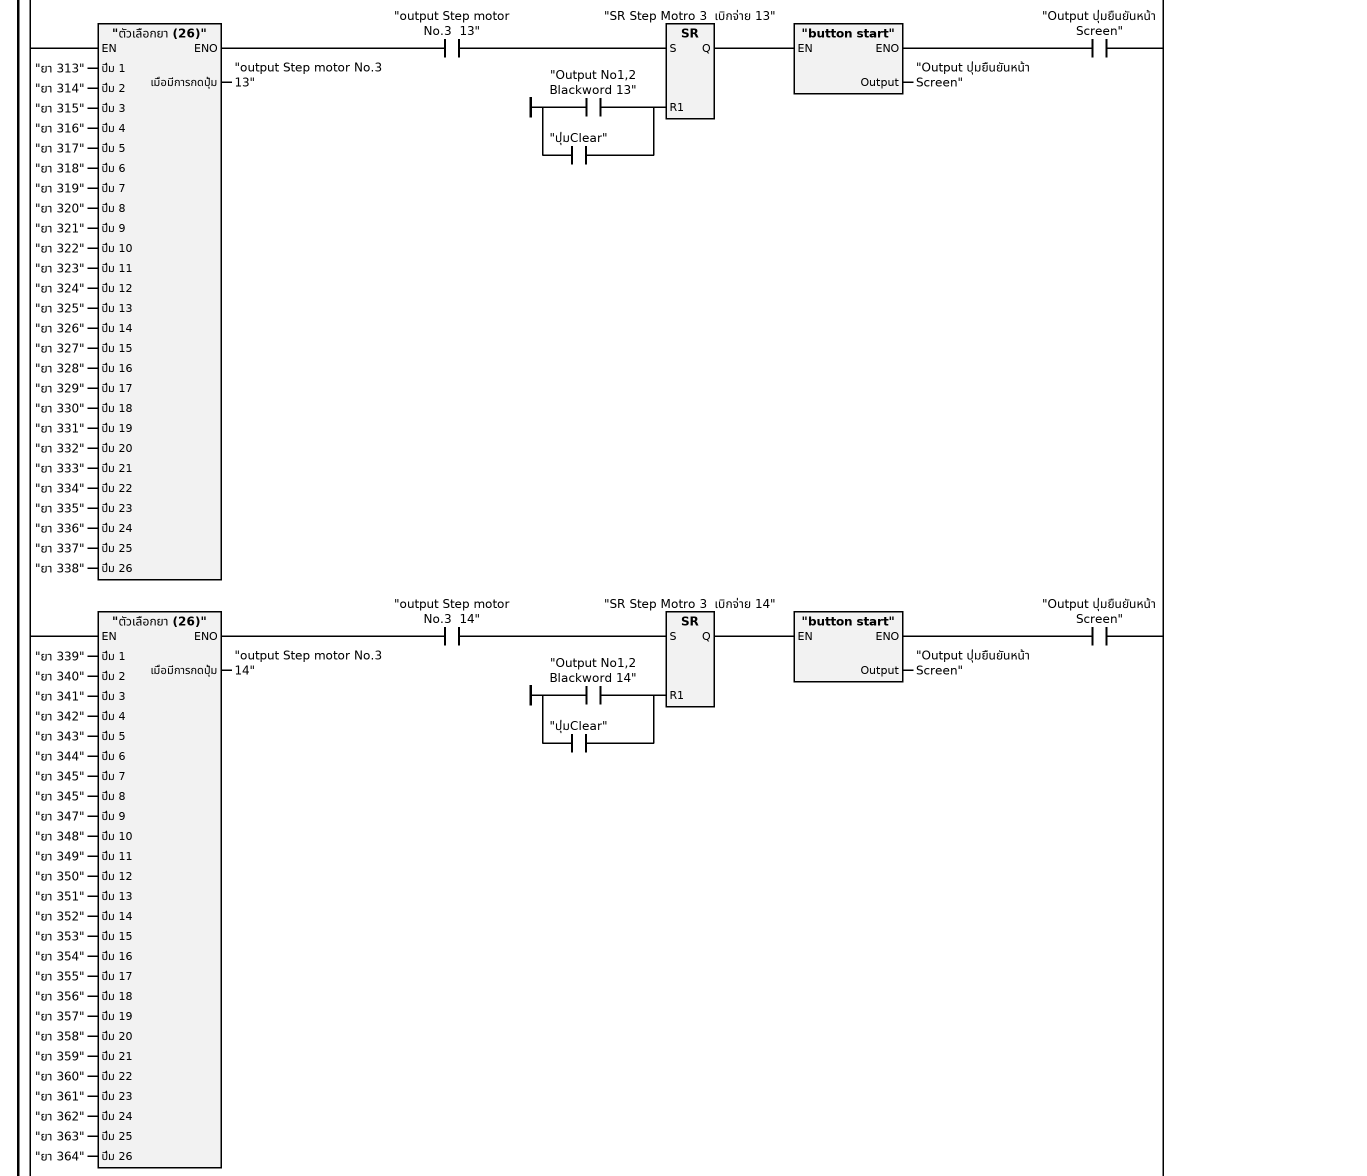
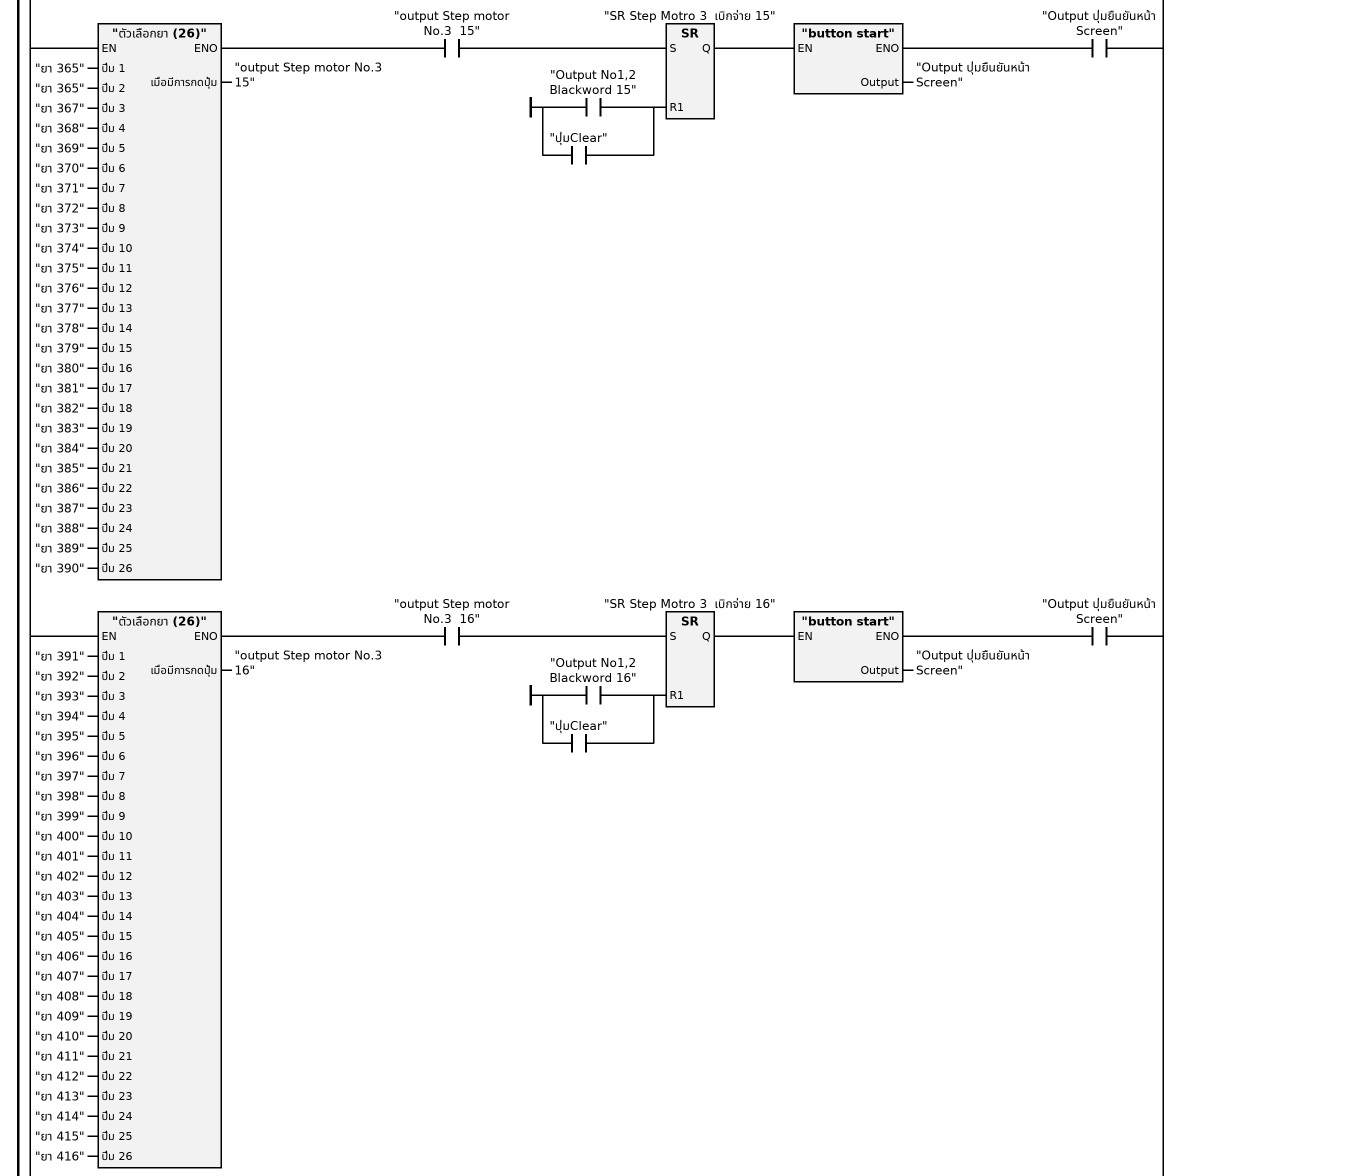
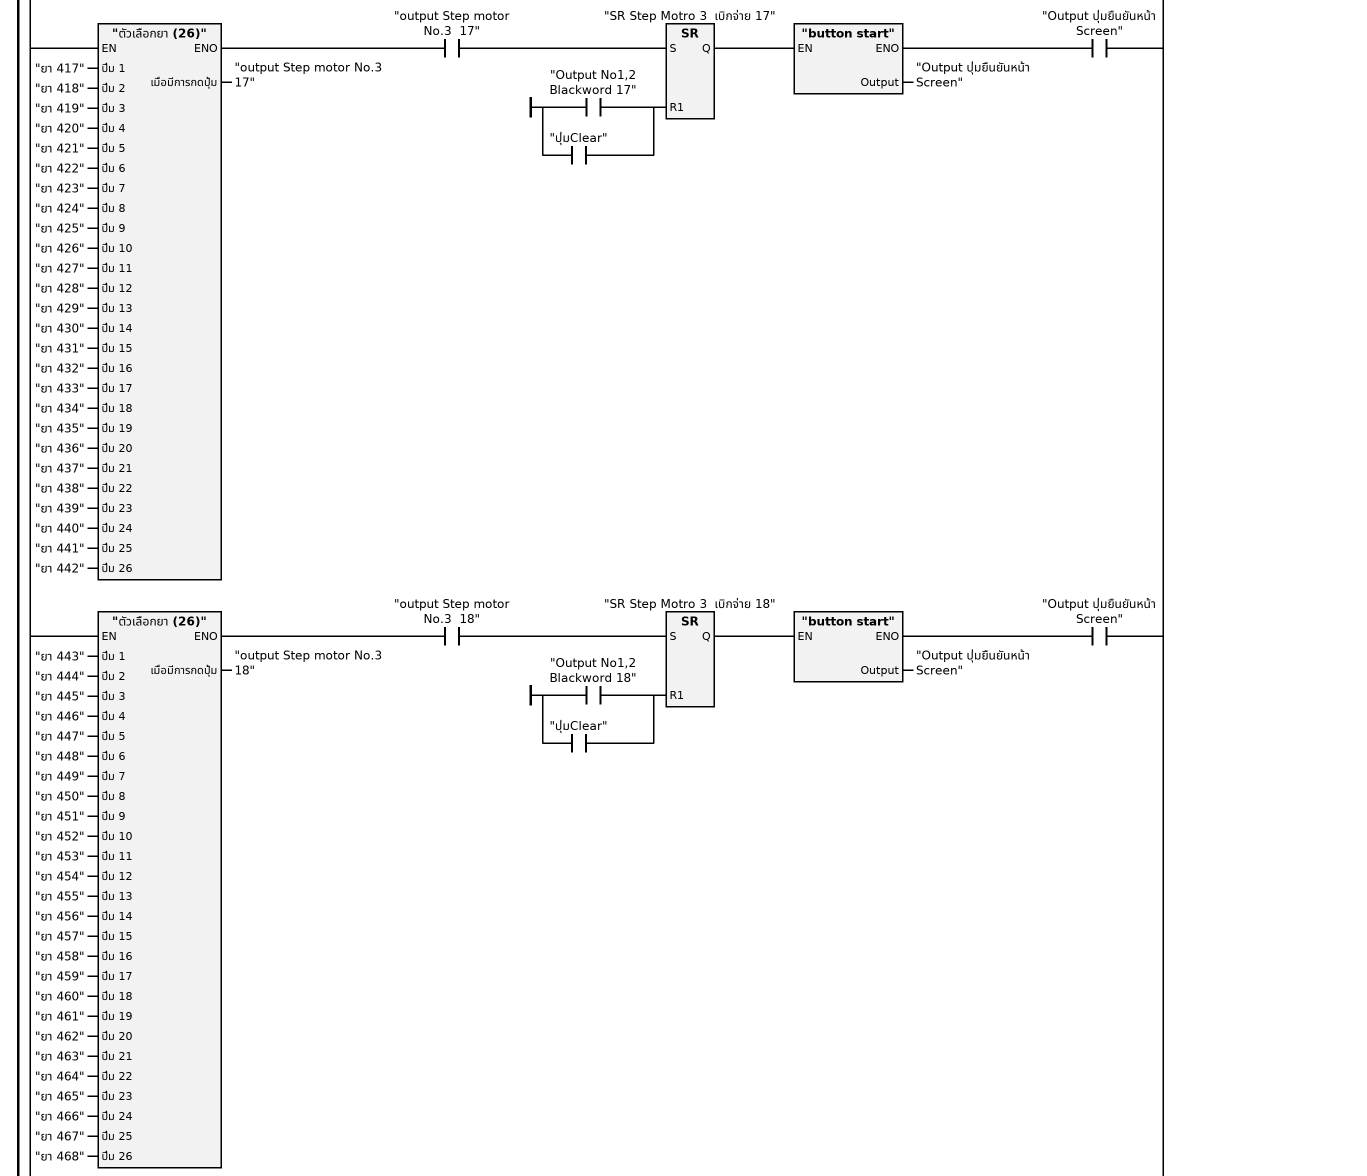
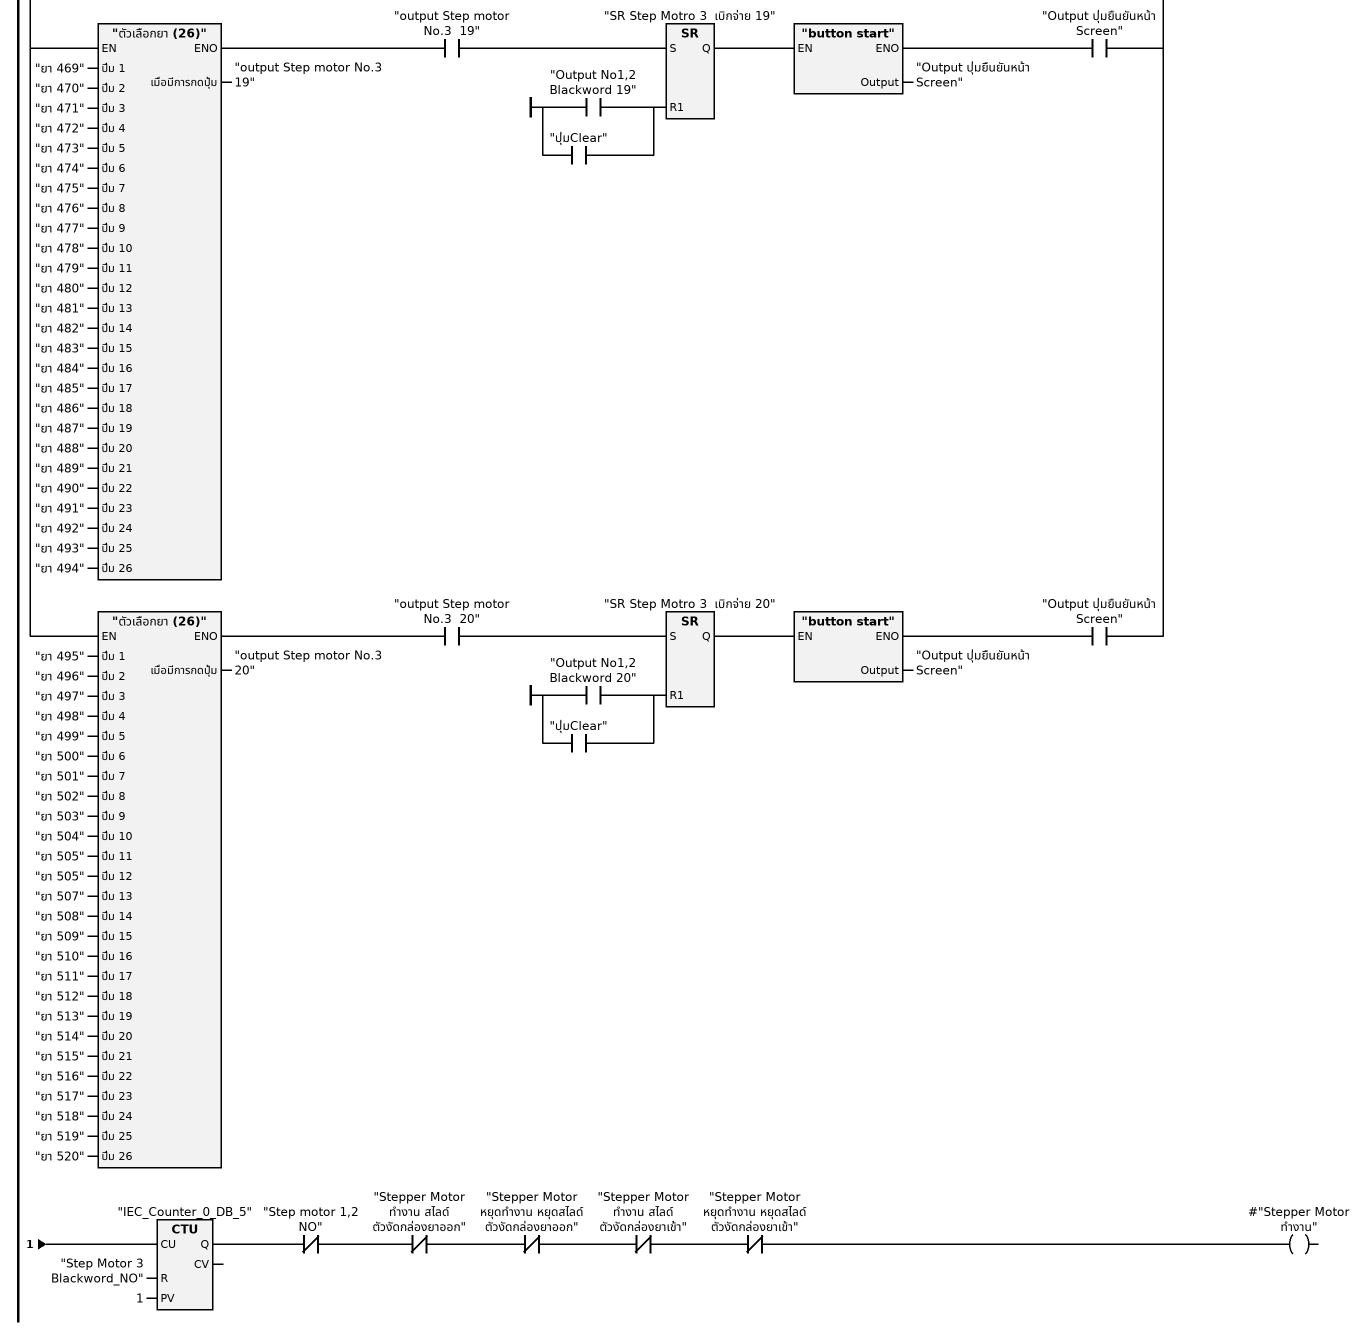
   "ตัวเลือกยา (26)"("ปึ่ม 1" := "ยา 1",
                     "ปึ่ม 2" := "ยา 2",
                     "ปึ่ม 3" := "ยา 3",
                     "ปึ่ม 4" := "ยา 4",
                     "ปึ่ม 5" := "ยา 5",
                     "ปึ่ม 6" := "ยา 6",
                     "ปึ่ม 7" := "ยา 7",
                     "ปึ่ม 8" := "ยา 8",
                     "ปึ่ม 9" := "ยา 9",
                     "ปึ่ม 10" := "ยา 10",
                     "ปึ่ม 11" := "ยา 11",
                     "ปึ่ม 12" := "ยา 12",
                     "ปึ่ม 13" := "ยา 13",
                     "ปึ่ม 14" := "ยา 14",
                     "ปึ่ม 15" := "ยา 15",
                     "ปึ่ม 16" := "ยา 16",
                     "ปึ่ม 17" := "ยา 17",
                     "ปึ่ม 18" := "ยา 18",
                     "ปึ่ม 19" := "ยา 19",
                     "ปึ่ม 20" := "ยา 20",
                     "ปึ่ม 21" := "ยา 21",
                     "ปึ่ม 22" := "ยา 22",
                     "ปึ่ม 23" := "ยา 23",
                     "ปึ่ม 24" := "ยา 24",
                     "ปึ่ม 25" := "ยา 25",
                     "ปึ่ม 26" := "ยา 26",
                     "เมื่ิอมีการกดปุ้ม" => "output Step motor No.3  1",
                     ENO => #_w1);
   IF #_w1 AND "output Step motor No.3  1" THEN
       "SR Step Motro 3  เบิกจ่าย 1" := TRUE;   // SR flip-flop
   END_IF;
   IF "Output No1,2 Blackword 1" OR "ปุ่มClear" THEN "SR Step Motro 3  เบิกจ่าย 1" := FALSE; END_IF;
   "button start"(EN := "SR Step Motro 3  เบิกจ่าย 1", Output => "Output ปุ่มยืนยันหน้า Screen", ENO => #_w2);
   #_w4 := #_w2 AND "Output ปุ่มยืนยันหน้า Screen";
   "ตัวเลือกยา (26)"("ปึ่ม 1" := "ยา 27",
                     "ปึ่ม 2" := "ยา 28",
                     "ปึ่ม 3" := "ยา 29",
                     "ปึ่ม 4" := "ยา 30",
                     "ปึ่ม 5" := "ยา 31",
                     "ปึ่ม 6" := "ยา 32",
                     "ปึ่ม 7" := "ยา 33",
                     "ปึ่ม 8" := "ยา 34",
                     "ปึ่ม 9" := "ยา 35",
                     "ปึ่ม 10" := "ยา 36",
                     "ปึ่ม 11" := "ยา 37",
                     "ปึ่ม 12" := "ยา 38",
                     "ปึ่ม 13" := "ยา 39",
                     "ปึ่ม 14" := "ยา 40",
                     "ปึ่ม 15" := "ยา 41",
                     "ปึ่ม 16" := "ยา 42",
                     "ปึ่ม 17" := "ยา 43",
                     "ปึ่ม 18" := "ยา 44",
                     "ปึ่ม 19" := "ยา 45",
                     "ปึ่ม 20" := "ยา 46",
                     "ปึ่ม 21" := "ยา 47",
                     "ปึ่ม 22" := "ยา 48",
                     "ปึ่ม 23" := "ยา 49",
                     "ปึ่ม 24" := "ยา 50",
                     "ปึ่ม 25" := "ยา 51",
                     "ปึ่ม 26" := "ยา 52",
                     "เมื่ิอมีการกดปุ้ม" => "output Step motor No.3  2",
                     ENO => #_w3);
   IF #_w3 AND "output Step motor No.3  2" THEN
       "SR Step Motro 3  เบิกจ่าย 2" := TRUE;   // SR flip-flop
   END_IF;
   IF "Output No1,2 Blackword 2" OR "ปุ่มClear" THEN "SR Step Motro 3  เบิกจ่าย 2" := FALSE; END_IF;
   "button start"(EN := "SR Step Motro 3  เบิกจ่าย 2", Output => "Output ปุ่มยืนยันหน้า Screen", ENO => #_w5);
   #_w7 := #_w5 AND "Output ปุ่มยืนยันหน้า Screen";
   "ตัวเลือกยา (26)"("ปึ่ม 1" := "ยา 53",
                     "ปึ่ม 2" := "ยา 54",
                     "ปึ่ม 3" := "ยา 55",
                     "ปึ่ม 4" := "ยา 56",
                     "ปึ่ม 5" := "ยา 57",
                     "ปึ่ม 6" := "ยา 58",
                     "ปึ่ม 7" := "ยา 59",
                     "ปึ่ม 8" := "ยา 60",
                     "ปึ่ม 9" := "ยา 61",
                     "ปึ่ม 10" := "ยา 62",
                     "ปึ่ม 11" := "ยา 63",
                     "ปึ่ม 12" := "ยา 64",
                     "ปึ่ม 13" := "ยา 65",
                     "ปึ่ม 14" := "ยา 66",
                     "ปึ่ม 15" := "ยา 67",
                     "ปึ่ม 16" := "ยา 68",
                     "ปึ่ม 17" := "ยา 69",
                     "ปึ่ม 18" := "ยา 70",
                     "ปึ่ม 19" := "ยา 71",
                     "ปึ่ม 20" := "ยา 72",
                     "ปึ่ม 21" := "ยา 73",
                     "ปึ่ม 22" := "ยา 74",
                     "ปึ่ม 23" := "ยา 75",
                     "ปึ่ม 24" := "ยา 76",
                     "ปึ่ม 25" := "ยา 77",
                     "ปึ่ม 26" := "ยา 78",
                     "เมื่ิอมีการกดปุ้ม" => "output Step motor No.3  3",
                     ENO => #_w6);
   IF #_w6 AND "output Step motor No.3  3" THEN
       "SR Step Motro 3  เบิกจ่าย 3" := TRUE;   // SR flip-flop
   END_IF;
   IF "Output No1,2 Blackword 3" OR "ปุ่มClear" THEN "SR Step Motro 3  เบิกจ่าย 3" := FALSE; END_IF;
   "button start"(EN := "SR Step Motro 3  เบิกจ่าย 3", Output => "Output ปุ่มยืนยันหน้า Screen", ENO => #_w8);
   #_w10 := #_w8 AND "Output ปุ่มยืนยันหน้า Screen";
   "ตัวเลือกยา (26)"("ปึ่ม 1" := "ยา 79",
                     "ปึ่ม 2" := "ยา 80",
                     "ปึ่ม 3" := "ยา 81",
                     "ปึ่ม 4" := "ยา 82",
                     "ปึ่ม 5" := "ยา 83",
                     "ปึ่ม 6" := "ยา 84",
                     "ปึ่ม 7" := "ยา 85",
                     "ปึ่ม 8" := "ยา 86",
                     "ปึ่ม 9" := "ยา 87",
                     "ปึ่ม 10" := "ยา 88",
                     "ปึ่ม 11" := "ยา 89",
                     "ปึ่ม 12" := "ยา 90",
                     "ปึ่ม 13" := "ยา 91",
                     "ปึ่ม 14" := "ยา 92",
                     "ปึ่ม 15" := "ยา 93",
                     "ปึ่ม 16" := "ยา 94",
                     "ปึ่ม 17" := "ยา 95",
                     "ปึ่ม 18" := "ยา 96",
                     "ปึ่ม 19" := "ยา 97",
                     "ปึ่ม 20" := "ยา 98",
                     "ปึ่ม 21" := "ยา 99",
                     "ปึ่ม 22" := "ยา 100",
                     "ปึ่ม 23" := "ยา 101",
                     "ปึ่ม 24" := "ยา 102",
                     "ปึ่ม 25" := "ยา 103",
                     "ปึ่ม 26" := "ยา 104",
                     "เมื่ิอมีการกดปุ้ม" => "output Step motor No.3  4",
                     ENO => #_w9);
   IF #_w9 AND "output Step motor No.3  4" THEN
       "SR Step Motro 3  เบิกจ่าย 4" := TRUE;   // SR flip-flop
   END_IF;
   IF "Output No1,2 Blackword 4" OR "ปุ่มClear" THEN "SR Step Motro 3  เบิกจ่าย 4" := FALSE; END_IF;
   "button start"(EN := "SR Step Motro 3  เบิกจ่าย 4", Output => "Output ปุ่มยืนยันหน้า Screen", ENO => #_w11);
   #_w13 := #_w11 AND "Output ปุ่มยืนยันหน้า Screen";
   "ตัวเลือกยา (26)"("ปึ่ม 1" := "ยา 105",
                     "ปึ่ม 2" := "ยา 106",
                     "ปึ่ม 3" := "ยา 107",
                     "ปึ่ม 4" := "ยา 108",
                     "ปึ่ม 5" := "ยา 109",
                     "ปึ่ม 6" := "ยา 110",
                     "ปึ่ม 7" := "ยา 111",
                     "ปึ่ม 8" := "ยา 112",
                     "ปึ่ม 9" := "ยา 113",
                     "ปึ่ม 10" := "ยา 114",
                     "ปึ่ม 11" := "ยา 115",
                     "ปึ่ม 12" := "ยา 116",
                     "ปึ่ม 13" := "ยา 117",
                     "ปึ่ม 14" := "ยา 118",
                     "ปึ่ม 15" := "ยา 119",
                     "ปึ่ม 16" := "ยา 120",
                     "ปึ่ม 17" := "ยา 121",
                     "ปึ่ม 18" := "ยา 122",
                     "ปึ่ม 19" := "ยา 123",
                     "ปึ่ม 20" := "ยา 124",
                     "ปึ่ม 21" := "ยา 125",
                     "ปึ่ม 22" := "ยา 126",
                     "ปึ่ม 23" := "ยา 127",
                     "ปึ่ม 24" := "ยา 128",
                     "ปึ่ม 25" := "ยา 129",
                     "ปึ่ม 26" := "ยา 130",
                     "เมื่ิอมีการกดปุ้ม" => "output Step motor No.3  5",
                     ENO => #_w12);
   IF #_w12 AND "output Step motor No.3  5" THEN
       "SR Step Motro 3  เบิกจ่าย 5" := TRUE;   // SR flip-flop
   END_IF;
   IF "Output No1,2 Blackword 5" OR "ปุ่มClear" THEN "SR Step Motro 3  เบิกจ่าย 5" := FALSE; END_IF;
   "button start"(EN := "SR Step Motro 3  เบิกจ่าย 5", Output => "Output ปุ่มยืนยันหน้า Screen", ENO => #_w14);
   #_w16 := #_w14 AND "Output ปุ่มยืนยันหน้า Screen";
   "ตัวเลือกยา (26)"("ปึ่ม 1" := "ยา 131",
                     "ปึ่ม 2" := "ยา 132",
                     "ปึ่ม 3" := "ยา 133",
                     "ปึ่ม 4" := "ยา 134",
                     "ปึ่ม 5" := "ยา 135",
                     "ปึ่ม 6" := "ยา 136",
                     "ปึ่ม 7" := "ยา 137",
                     "ปึ่ม 8" := "ยา 138",
                     "ปึ่ม 9" := "ยา 139",
                     "ปึ่ม 10" := "ยา 140",
                     "ปึ่ม 11" := "ยา 141",
                     "ปึ่ม 12" := "ยา 142",
                     "ปึ่ม 13" := "ยา 143",
                     "ปึ่ม 14" := "ยา 144",
                     "ปึ่ม 15" := "ยา 145",
                     "ปึ่ม 16" := "ยา 146",
                     "ปึ่ม 17" := "ยา 147",
                     "ปึ่ม 18" := "ยา 148",
                     "ปึ่ม 19" := "ยา 149",
                     "ปึ่ม 20" := "ยา 150",
                     "ปึ่ม 21" := "ยา 151",
                     "ปึ่ม 22" := "ยา 152",
                     "ปึ่ม 23" := "ยา 153",
                     "ปึ่ม 24" := "ยา 154",
                     "ปึ่ม 25" := "ยา 155",
                     "ปึ่ม 26" := "ยา 156",
                     "เมื่ิอมีการกดปุ้ม" => "output Step motor No.3  6",
                     ENO => #_w15);
   IF #_w15 AND "output Step motor No.3  6" THEN
       "SR Step Motro 3  เบิกจ่าย 6" := TRUE;   // SR flip-flop
   END_IF;
   IF "Output No1,2 Blackword 6" OR "ปุ่มClear" THEN "SR Step Motro 3  เบิกจ่าย 6" := FALSE; END_IF;
   "button start"(EN := "SR Step Motro 3  เบิกจ่าย 6", Output => "Output ปุ่มยืนยันหน้า Screen", ENO => #_w17);
   #_w19 := #_w17 AND "Output ปุ่มยืนยันหน้า Screen";
   "ตัวเลือกยา (26)"("ปึ่ม 1" := "ยา 157",
                     "ปึ่ม 2" := "ยา 158",
                     "ปึ่ม 3" := "ยา 159",
                     "ปึ่ม 4" := "ยา 160",
                     "ปึ่ม 5" := "ยา 161",
                     "ปึ่ม 6" := "ยา 162",
                     "ปึ่ม 7" := "ยา 163",
                     "ปึ่ม 8" := "ยา 164",
                     "ปึ่ม 9" := "ยา 165",
                     "ปึ่ม 10" := "ยา 166",
                     "ปึ่ม 11" := "ยา 167",
                     "ปึ่ม 12" := "ยา 168",
                     "ปึ่ม 13" := "ยา 169",
                     "ปึ่ม 14" := "ยา 170",
                     "ปึ่ม 15" := "ยา 171",
                     "ปึ่ม 16" := "ยา 172",
                     "ปึ่ม 17" := "ยา 173",
                     "ปึ่ม 18" := "ยา 174",
                     "ปึ่ม 19" := "ยา 175",
                     "ปึ่ม 20" := "ยา 176",
                     "ปึ่ม 21" := "ยา 177",
                     "ปึ่ม 22" := "ยา 178",
                     "ปึ่ม 23" := "ยา 179",
                     "ปึ่ม 24" := "ยา 180",
                     "ปึ่ม 25" := "ยา 181",
                     "ปึ่ม 26" := "ยา 182",
                     "เมื่ิอมีการกดปุ้ม" => "output Step motor No.3  7",
                     ENO => #_w18);
   IF #_w18 AND "output Step motor No.3  7" THEN
       "SR Step Motro 3  เบิกจ่าย 7" := TRUE;   // SR flip-flop
   END_IF;
   IF "Output No1,2 Blackword 7" OR "ปุ่มClear" THEN "SR Step Motro 3  เบิกจ่าย 7" := FALSE; END_IF;
   "button start"(EN := "SR Step Motro 3  เบิกจ่าย 7", Output => "Output ปุ่มยืนยันหน้า Screen", ENO => #_w20);
   #_w22 := #_w20 AND "Output ปุ่มยืนยันหน้า Screen";
   "ตัวเลือกยา (26)"("ปึ่ม 1" := "ยา 183",
                     "ปึ่ม 2" := "ยา 184",
                     "ปึ่ม 3" := "ยา 185",
                     "ปึ่ม 4" := "ยา 186",
                     "ปึ่ม 5" := "ยา 187",
                     "ปึ่ม 6" := "ยา 188",
                     "ปึ่ม 7" := "ยา 189",
                     "ปึ่ม 8" := "ยา 190",
                     "ปึ่ม 9" := "ยา 191",
                     "ปึ่ม 10" := "ยา 192",
                     "ปึ่ม 11" := "ยา 193",
                     "ปึ่ม 12" := "ยา 194",
                     "ปึ่ม 13" := "ยา 195",
                     "ปึ่ม 14" := "ยา 196",
                     "ปึ่ม 15" := "ยา 197",
                     "ปึ่ม 16" := "ยา 198",
                     "ปึ่ม 17" := "ยา 199",
                     "ปึ่ม 18" := "ยา 200",
                     "ปึ่ม 19" := "ยา 201",
                     "ปึ่ม 20" := "ยา 202",
                     "ปึ่ม 21" := "ยา 203",
                     "ปึ่ม 22" := "ยา 204",
                     "ปึ่ม 23" := "ยา 205",
                     "ปึ่ม 24" := "ยา 206",
                     "ปึ่ม 25" := "ยา 207",
                     "ปึ่ม 26" := "ยา 208",
                     "เมื่ิอมีการกดปุ้ม" => "output Step motor No.3  8",
                     ENO => #_w21);
   IF #_w21 AND "output Step motor No.3  8" THEN
       "SR Step Motro 3  เบิกจ่าย 8" := TRUE;   // SR flip-flop
   END_IF;
   IF "Output No1,2 Blackword 8" OR "ปุ่มClear" THEN "SR Step Motro 3  เบิกจ่าย 8" := FALSE; END_IF;
   "button start"(EN := "SR Step Motro 3  เบิกจ่าย 8", Output => "Output ปุ่มยืนยันหน้า Screen", ENO => #_w23);
   #_w25 := #_w23 AND "Output ปุ่มยืนยันหน้า Screen";
   "ตัวเลือกยา (26)"("ปึ่ม 1" := "ยา 209",
                     "ปึ่ม 2" := "ยา 210",
                     "ปึ่ม 3" := "ยา 211",
                     "ปึ่ม 4" := "ยา 212",
                     "ปึ่ม 5" := "ยา 213",
                     "ปึ่ม 6" := "ยา 214",
                     "ปึ่ม 7" := "ยา 215",
                     "ปึ่ม 8" := "ยา 216",
                     "ปึ่ม 9" := "ยา 217",
                     "ปึ่ม 10" := "ยา 218",
                     "ปึ่ม 11" := "ยา 219",
                     "ปึ่ม 12" := "ยา 220",
                     "ปึ่ม 13" := "ยา 221",
                     "ปึ่ม 14" := "ยา 222",
                     "ปึ่ม 15" := "ยา 223",
                     "ปึ่ม 16" := "ยา 224",
                     "ปึ่ม 17" := "ยา 225",
                     "ปึ่ม 18" := "ยา 226",
                     "ปึ่ม 19" := "ยา 227",
                     "ปึ่ม 20" := "ยา 228",
                     "ปึ่ม 21" := "ยา 229",
                     "ปึ่ม 22" := "ยา 230",
                     "ปึ่ม 23" := "ยา 231",
                     "ปึ่ม 24" := "ยา 232",
                     "ปึ่ม 25" := "ยา 233",
                     "ปึ่ม 26" := "ยา 234",
                     "เมื่ิอมีการกดปุ้ม" => "output Step motor No.3  9",
                     ENO => #_w24);
   IF #_w24 AND "output Step motor No.3  9" THEN
       "SR Step Motro 3  เบิกจ่าย 9" := TRUE;   // SR flip-flop
   END_IF;
   IF "Output No1,2 Blackword 9" OR "ปุ่มClear" THEN "SR Step Motro 3  เบิกจ่าย 9" := FALSE; END_IF;
   "button start"(EN := "SR Step Motro 3  เบิกจ่าย 9", Output => "Output ปุ่มยืนยันหน้า Screen", ENO => #_w26);
   #_w28 := #_w26 AND "Output ปุ่มยืนยันหน้า Screen";
   "ตัวเลือกยา (26)"("ปึ่ม 1" := "ยา 235",
                     "ปึ่ม 2" := "ยา 236",
                     "ปึ่ม 3" := "ยา 234",
                     "ปึ่ม 4" := "ยา 238",
                     "ปึ่ม 5" := "ยา 239",
                     "ปึ่ม 6" := "ยา 240",
                     "ปึ่ม 7" := "ยา 241",
                     "ปึ่ม 8" := "ยา 242",
                     "ปึ่ม 9" := "ยา 243",
                     "ปึ่ม 10" := "ยา 244",
                     "ปึ่ม 11" := "ยา 245",
                     "ปึ่ม 12" := "ยา 246",
                     "ปึ่ม 13" := "ยา 247",
                     "ปึ่ม 14" := "ยา 248",
                     "ปึ่ม 15" := "ยา 249",
                     "ปึ่ม 16" := "ยา 250",
                     "ปึ่ม 17" := "ยา 251",
                     "ปึ่ม 18" := "ยา 252",
                     "ปึ่ม 19" := "ยา 253",
                     "ปึ่ม 20" := "ยา 254",
                     "ปึ่ม 21" := "ยา 255",
                     "ปึ่ม 22" := "ยา 256",
                     "ปึ่ม 23" := "ยา 257",
                     "ปึ่ม 24" := "ยา 258",
                     "ปึ่ม 25" := "ยา 259",
                     "ปึ่ม 26" := "ยา 260",
                     "เมื่ิอมีการกดปุ้ม" => "output Step motor No.3  10",
                     ENO => #_w27);
   IF #_w27 AND "output Step motor No.3  10" THEN
       "SR Step Motro 3  เบิกจ่าย 10" := TRUE;   // SR flip-flop
   END_IF;
   IF "Output No1,2 Blackword 10" OR "ปุ่มClear" THEN "SR Step Motro 3  เบิกจ่าย 10" := FALSE; END_IF;
   "button start"(EN := "SR Step Motro 3  เบิกจ่าย 10", Output => "Output ปุ่มยืนยันหน้า Screen", ENO => #_w29);
   #_w31 := #_w29 AND "Output ปุ่มยืนยันหน้า Screen";
   "ตัวเลือกยา (26)"("ปึ่ม 1" := "ยา 261",
                     "ปึ่ม 2" := "ยา 262",
                     "ปึ่ม 3" := "ยา 263",
                     "ปึ่ม 4" := "ยา 264",
                     "ปึ่ม 5" := "ยา 265",
                     "ปึ่ม 6" := "ยา 266",
                     "ปึ่ม 7" := "ยา 267",
                     "ปึ่ม 8" := "ยา 268",
                     "ปึ่ม 9" := "ยา 269",
                     "ปึ่ม 10" := "ยา 270",
                     "ปึ่ม 11" := "ยา 271",
                     "ปึ่ม 12" := "ยา 272",
                     "ปึ่ม 13" := "ยา 273",
                     "ปึ่ม 14" := "ยา 274",
                     "ปึ่ม 15" := "ยา 275",
                     "ปึ่ม 16" := "ยา 276",
                     "ปึ่ม 17" := "ยา 277",
                     "ปึ่ม 18" := "ยา 278",
                     "ปึ่ม 19" := "ยา 279",
                     "ปึ่ม 20" := "ยา 280",
                     "ปึ่ม 21" := "ยา 281",
                     "ปึ่ม 22" := "ยา 282",
                     "ปึ่ม 23" := "ยา 283",
                     "ปึ่ม 24" := "ยา 284",
                     "ปึ่ม 25" := "ยา 285",
                     "ปึ่ม 26" := "ยา 286",
                     "เมื่ิอมีการกดปุ้ม" => "output Step motor No.3  11",
                     ENO => #_w30);
   IF #_w30 AND "output Step motor No.3  11" THEN
       "SR Step Motro 3  เบิกจ่าย 11" := TRUE;   // SR flip-flop
   END_IF;
   IF "Output No1,2 Blackword 11" OR "ปุ่มClear" THEN "SR Step Motro 3  เบิกจ่าย 11" := FALSE; END_IF;
   "button start"(EN := "SR Step Motro 3  เบิกจ่าย 11", Output => "Output ปุ่มยืนยันหน้า Screen", ENO => #_w32);
   #_w34 := #_w32 AND "Output ปุ่มยืนยันหน้า Screen";
   "ตัวเลือกยา (26)"("ปึ่ม 1" := "ยา 287",
                     "ปึ่ม 2" := "ยา 288",
                     "ปึ่ม 3" := "ยา 289",
                     "ปึ่ม 4" := "ยา 290",
                     "ปึ่ม 5" := "ยา 291",
                     "ปึ่ม 6" := "ยา 292",
                     "ปึ่ม 7" := "ยา 293",
                     "ปึ่ม 8" := "ยา 294",
                     "ปึ่ม 9" := "ยา 295",
                     "ปึ่ม 10" := "ยา 296",
                     "ปึ่ม 11" := "ยา 297",
                     "ปึ่ม 12" := "ยา 298",
                     "ปึ่ม 13" := "ยา 299",
                     "ปึ่ม 14" := "ยา 300",
                     "ปึ่ม 15" := "ยา 301",
                     "ปึ่ม 16" := "ยา 302",
                     "ปึ่ม 17" := "ยา 303",
                     "ปึ่ม 18" := "ยา 304",
                     "ปึ่ม 19" := "ยา 305",
                     "ปึ่ม 20" := "ยา 306",
                     "ปึ่ม 21" := "ยา 307",
                     "ปึ่ม 22" := "ยา 308",
                     "ปึ่ม 23" := "ยา 309",
                     "ปึ่ม 24" := "ยา 310",
                     "ปึ่ม 25" := "ยา 311",
                     "ปึ่ม 26" := "ยา 312",
                     "เมื่ิอมีการกดปุ้ม" => "output Step motor No.3  12",
                     ENO => #_w33);
   IF #_w33 AND "output Step motor No.3  12" THEN
       "SR Step Motro 3  เบิกจ่าย 12" := TRUE;   // SR flip-flop
   END_IF;
   IF "Output No1,2 Blackword 12" OR "ปุ่มClear" THEN "SR Step Motro 3  เบิกจ่าย 12" := FALSE; END_IF;
   "button start"(EN := "SR Step Motro 3  เบิกจ่าย 12", Output => "Output ปุ่มยืนยันหน้า Screen", ENO => #_w35);
   #_w37 := #_w35 AND "Output ปุ่มยืนยันหน้า Screen";
   "ตัวเลือกยา (26)"("ปึ่ม 1" := "ยา 313",
                     "ปึ่ม 2" := "ยา 314",
                     "ปึ่ม 3" := "ยา 315",
                     "ปึ่ม 4" := "ยา 316",
                     "ปึ่ม 5" := "ยา 317",
                     "ปึ่ม 6" := "ยา 318",
                     "ปึ่ม 7" := "ยา 319",
                     "ปึ่ม 8" := "ยา 320",
                     "ปึ่ม 9" := "ยา 321",
                     "ปึ่ม 10" := "ยา 322",
                     "ปึ่ม 11" := "ยา 323",
                     "ปึ่ม 12" := "ยา 324",
                     "ปึ่ม 13" := "ยา 325",
                     "ปึ่ม 14" := "ยา 326",
                     "ปึ่ม 15" := "ยา 327",
                     "ปึ่ม 16" := "ยา 328",
                     "ปึ่ม 17" := "ยา 329",
                     "ปึ่ม 18" := "ยา 330",
                     "ปึ่ม 19" := "ยา 331",
                     "ปึ่ม 20" := "ยา 332",
                     "ปึ่ม 21" := "ยา 333",
                     "ปึ่ม 22" := "ยา 334",
                     "ปึ่ม 23" := "ยา 335",
                     "ปึ่ม 24" := "ยา 336",
                     "ปึ่ม 25" := "ยา 337",
                     "ปึ่ม 26" := "ยา 338",
                     "เมื่ิอมีการกดปุ้ม" => "output Step motor No.3  13",
                     ENO => #_w36);
   IF #_w36 AND "output Step motor No.3  13" THEN
       "SR Step Motro 3  เบิกจ่าย 13" := TRUE;   // SR flip-flop
   END_IF;
   IF "Output No1,2 Blackword 13" OR "ปุ่มClear" THEN "SR Step Motro 3  เบิกจ่าย 13" := FALSE; END_IF;
   "button start"(EN := "SR Step Motro 3  เบิกจ่าย 13", Output => "Output ปุ่มยืนยันหน้า Screen", ENO => #_w38);
   #_w40 := #_w38 AND "Output ปุ่มยืนยันหน้า Screen";
   "ตัวเลือกยา (26)"("ปึ่ม 1" := "ยา 339",
                     "ปึ่ม 2" := "ยา 340",
                     "ปึ่ม 3" := "ยา 341",
                     "ปึ่ม 4" := "ยา 342",
                     "ปึ่ม 5" := "ยา 343",
                     "ปึ่ม 6" := "ยา 344",
                     "ปึ่ม 7" := "ยา 345",
                     "ปึ่ม 8" := "ยา 345",
                     "ปึ่ม 9" := "ยา 347",
                     "ปึ่ม 10" := "ยา 348",
                     "ปึ่ม 11" := "ยา 349",
                     "ปึ่ม 12" := "ยา 350",
                     "ปึ่ม 13" := "ยา 351",
                     "ปึ่ม 14" := "ยา 352",
                     "ปึ่ม 15" := "ยา 353",
                     "ปึ่ม 16" := "ยา 354",
                     "ปึ่ม 17" := "ยา 355",
                     "ปึ่ม 18" := "ยา 356",
                     "ปึ่ม 19" := "ยา 357",
                     "ปึ่ม 20" := "ยา 358",
                     "ปึ่ม 21" := "ยา 359",
                     "ปึ่ม 22" := "ยา 360",
                     "ปึ่ม 23" := "ยา 361",
                     "ปึ่ม 24" := "ยา 362",
                     "ปึ่ม 25" := "ยา 363",
                     "ปึ่ม 26" := "ยา 364",
                     "เมื่ิอมีการกดปุ้ม" => "output Step motor No.3  14",
                     ENO => #_w39);
   IF #_w39 AND "output Step motor No.3  14" THEN
       "SR Step Motro 3  เบิกจ่าย 14" := TRUE;   // SR flip-flop
   END_IF;
   IF "Output No1,2 Blackword 14" OR "ปุ่มClear" THEN "SR Step Motro 3  เบิกจ่าย 14" := FALSE; END_IF;
   "button start"(EN := "SR Step Motro 3  เบิกจ่าย 14", Output => "Output ปุ่มยืนยันหน้า Screen", ENO => #_w41);
   #_w43 := #_w41 AND "Output ปุ่มยืนยันหน้า Screen";
   "ตัวเลือกยา (26)"("ปึ่ม 1" := "ยา 365",
                     "ปึ่ม 2" := "ยา 365",
                     "ปึ่ม 3" := "ยา 367",
                     "ปึ่ม 4" := "ยา 368",
                     "ปึ่ม 5" := "ยา 369",
                     "ปึ่ม 6" := "ยา 370",
                     "ปึ่ม 7" := "ยา 371",
                     "ปึ่ม 8" := "ยา 372",
                     "ปึ่ม 9" := "ยา 373",
                     "ปึ่ม 10" := "ยา 374",
                     "ปึ่ม 11" := "ยา 375",
                     "ปึ่ม 12" := "ยา 376",
                     "ปึ่ม 13" := "ยา 377",
                     "ปึ่ม 14" := "ยา 378",
                     "ปึ่ม 15" := "ยา 379",
                     "ปึ่ม 16" := "ยา 380",
                     "ปึ่ม 17" := "ยา 381",
                     "ปึ่ม 18" := "ยา 382",
                     "ปึ่ม 19" := "ยา 383",
                     "ปึ่ม 20" := "ยา 384",
                     "ปึ่ม 21" := "ยา 385",
                     "ปึ่ม 22" := "ยา 386",
                     "ปึ่ม 23" := "ยา 387",
                     "ปึ่ม 24" := "ยา 388",
                     "ปึ่ม 25" := "ยา 389",
                     "ปึ่ม 26" := "ยา 390",
                     "เมื่ิอมีการกดปุ้ม" => "output Step motor No.3  15",
                     ENO => #_w42);
   IF #_w42 AND "output Step motor No.3  15" THEN
       "SR Step Motro 3  เบิกจ่าย 15" := TRUE;   // SR flip-flop
   END_IF;
   IF "Output No1,2 Blackword 15" OR "ปุ่มClear" THEN "SR Step Motro 3  เบิกจ่าย 15" := FALSE; END_IF;
   "button start"(EN := "SR Step Motro 3  เบิกจ่าย 15", Output => "Output ปุ่มยืนยันหน้า Screen", ENO => #_w44);
   #_w46 := #_w44 AND "Output ปุ่มยืนยันหน้า Screen";
   "ตัวเลือกยา (26)"("ปึ่ม 1" := "ยา 391",
                     "ปึ่ม 2" := "ยา 392",
                     "ปึ่ม 3" := "ยา 393",
                     "ปึ่ม 4" := "ยา 394",
                     "ปึ่ม 5" := "ยา 395",
                     "ปึ่ม 6" := "ยา 396",
                     "ปึ่ม 7" := "ยา 397",
                     "ปึ่ม 8" := "ยา 398",
                     "ปึ่ม 9" := "ยา 399",
                     "ปึ่ม 10" := "ยา 400",
                     "ปึ่ม 11" := "ยา 401",
                     "ปึ่ม 12" := "ยา 402",
                     "ปึ่ม 13" := "ยา 403",
                     "ปึ่ม 14" := "ยา 404",
                     "ปึ่ม 15" := "ยา 405",
                     "ปึ่ม 16" := "ยา 406",
                     "ปึ่ม 17" := "ยา 407",
                     "ปึ่ม 18" := "ยา 408",
                     "ปึ่ม 19" := "ยา 409",
                     "ปึ่ม 20" := "ยา 410",
                     "ปึ่ม 21" := "ยา 411",
                     "ปึ่ม 22" := "ยา 412",
                     "ปึ่ม 23" := "ยา 413",
                     "ปึ่ม 24" := "ยา 414",
                     "ปึ่ม 25" := "ยา 415",
                     "ปึ่ม 26" := "ยา 416",
                     "เมื่ิอมีการกดปุ้ม" => "output Step motor No.3  16",
                     ENO => #_w45);
   IF #_w45 AND "output Step motor No.3  16" THEN
       "SR Step Motro 3  เบิกจ่าย 16" := TRUE;   // SR flip-flop
   END_IF;
   IF "Output No1,2 Blackword 16" OR "ปุ่มClear" THEN "SR Step Motro 3  เบิกจ่าย 16" := FALSE; END_IF;
   "button start"(EN := "SR Step Motro 3  เบิกจ่าย 16", Output => "Output ปุ่มยืนยันหน้า Screen", ENO => #_w47);
   #_w49 := #_w47 AND "Output ปุ่มยืนยันหน้า Screen";
   "ตัวเลือกยา (26)"("ปึ่ม 1" := "ยา 417",
                     "ปึ่ม 2" := "ยา 418",
                     "ปึ่ม 3" := "ยา 419",
                     "ปึ่ม 4" := "ยา 420",
                     "ปึ่ม 5" := "ยา 421",
                     "ปึ่ม 6" := "ยา 422",
                     "ปึ่ม 7" := "ยา 423",
                     "ปึ่ม 8" := "ยา 424",
                     "ปึ่ม 9" := "ยา 425",
                     "ปึ่ม 10" := "ยา 426",
                     "ปึ่ม 11" := "ยา 427",
                     "ปึ่ม 12" := "ยา 428",
                     "ปึ่ม 13" := "ยา 429",
                     "ปึ่ม 14" := "ยา 430",
                     "ปึ่ม 15" := "ยา 431",
                     "ปึ่ม 16" := "ยา 432",
                     "ปึ่ม 17" := "ยา 433",
                     "ปึ่ม 18" := "ยา 434",
                     "ปึ่ม 19" := "ยา 435",
                     "ปึ่ม 20" := "ยา 436",
                     "ปึ่ม 21" := "ยา 437",
                     "ปึ่ม 22" := "ยา 438",
                     "ปึ่ม 23" := "ยา 439",
                     "ปึ่ม 24" := "ยา 440",
                     "ปึ่ม 25" := "ยา 441",
                     "ปึ่ม 26" := "ยา 442",
                     "เมื่ิอมีการกดปุ้ม" => "output Step motor No.3  17",
                     ENO => #_w48);
   IF #_w48 AND "output Step motor No.3  17" THEN
       "SR Step Motro 3  เบิกจ่าย 17" := TRUE;   // SR flip-flop
   END_IF;
   IF "Output No1,2 Blackword 17" OR "ปุ่มClear" THEN "SR Step Motro 3  เบิกจ่าย 17" := FALSE; END_IF;
   "button start"(EN := "SR Step Motro 3  เบิกจ่าย 17", Output => "Output ปุ่มยืนยันหน้า Screen", ENO => #_w50);
   #_w52 := #_w50 AND "Output ปุ่มยืนยันหน้า Screen";
   "ตัวเลือกยา (26)"("ปึ่ม 1" := "ยา 443",
                     "ปึ่ม 2" := "ยา 444",
                     "ปึ่ม 3" := "ยา 445",
                     "ปึ่ม 4" := "ยา 446",
                     "ปึ่ม 5" := "ยา 447",
                     "ปึ่ม 6" := "ยา 448",
                     "ปึ่ม 7" := "ยา 449",
                     "ปึ่ม 8" := "ยา 450",
                     "ปึ่ม 9" := "ยา 451",
                     "ปึ่ม 10" := "ยา 452",
                     "ปึ่ม 11" := "ยา 453",
                     "ปึ่ม 12" := "ยา 454",
                     "ปึ่ม 13" := "ยา 455",
                     "ปึ่ม 14" := "ยา 456",
                     "ปึ่ม 15" := "ยา 457",
                     "ปึ่ม 16" := "ยา 458",
                     "ปึ่ม 17" := "ยา 459",
                     "ปึ่ม 18" := "ยา 460",
                     "ปึ่ม 19" := "ยา 461",
                     "ปึ่ม 20" := "ยา 462",
                     "ปึ่ม 21" := "ยา 463",
                     "ปึ่ม 22" := "ยา 464",
                     "ปึ่ม 23" := "ยา 465",
                     "ปึ่ม 24" := "ยา 466",
                     "ปึ่ม 25" := "ยา 467",
                     "ปึ่ม 26" := "ยา 468",
                     "เมื่ิอมีการกดปุ้ม" => "output Step motor No.3  18",
                     ENO => #_w51);
   IF #_w51 AND "output Step motor No.3  18" THEN
       "SR Step Motro 3  เบิกจ่าย 18" := TRUE;   // SR flip-flop
   END_IF;
   IF "Output No1,2 Blackword 18" OR "ปุ่มClear" THEN "SR Step Motro 3  เบิกจ่าย 18" := FALSE; END_IF;
   "button start"(EN := "SR Step Motro 3  เบิกจ่าย 18", Output => "Output ปุ่มยืนยันหน้า Screen", ENO => #_w53);
   #_w55 := #_w53 AND "Output ปุ่มยืนยันหน้า Screen";
   "ตัวเลือกยา (26)"("ปึ่ม 1" := "ยา 469",
                     "ปึ่ม 2" := "ยา 470",
                     "ปึ่ม 3" := "ยา 471",
                     "ปึ่ม 4" := "ยา 472",
                     "ปึ่ม 5" := "ยา 473",
                     "ปึ่ม 6" := "ยา 474",
                     "ปึ่ม 7" := "ยา 475",
                     "ปึ่ม 8" := "ยา 476",
                     "ปึ่ม 9" := "ยา 477",
                     "ปึ่ม 10" := "ยา 478",
                     "ปึ่ม 11" := "ยา 479",
                     "ปึ่ม 12" := "ยา 480",
                     "ปึ่ม 13" := "ยา 481",
                     "ปึ่ม 14" := "ยา 482",
                     "ปึ่ม 15" := "ยา 483",
                     "ปึ่ม 16" := "ยา 484",
                     "ปึ่ม 17" := "ยา 485",
                     "ปึ่ม 18" := "ยา 486",
                     "ปึ่ม 19" := "ยา 487",
                     "ปึ่ม 20" := "ยา 488",
                     "ปึ่ม 21" := "ยา 489",
                     "ปึ่ม 22" := "ยา 490",
                     "ปึ่ม 23" := "ยา 491",
                     "ปึ่ม 24" := "ยา 492",
                     "ปึ่ม 25" := "ยา 493",
                     "ปึ่ม 26" := "ยา 494",
                     "เมื่ิอมีการกดปุ้ม" => "output Step motor No.3  19",
                     ENO => #_w54);
   IF #_w54 AND "output Step motor No.3  19" THEN
       "SR Step Motro 3  เบิกจ่าย 19" := TRUE;   // SR flip-flop
   END_IF;
   IF "Output No1,2 Blackword 19" OR "ปุ่มClear" THEN "SR Step Motro 3  เบิกจ่าย 19" := FALSE; END_IF;
   "button start"(EN := "SR Step Motro 3  เบิกจ่าย 19", Output => "Output ปุ่มยืนยันหน้า Screen", ENO => #_w56);
   #_w58 := #_w56 AND "Output ปุ่มยืนยันหน้า Screen";
   "ตัวเลือกยา (26)"("ปึ่ม 1" := "ยา 495",
                     "ปึ่ม 2" := "ยา 496",
                     "ปึ่ม 3" := "ยา 497",
                     "ปึ่ม 4" := "ยา 498",
                     "ปึ่ม 5" := "ยา 499",
                     "ปึ่ม 6" := "ยา 500",
                     "ปึ่ม 7" := "ยา 501",
                     "ปึ่ม 8" := "ยา 502",
                     "ปึ่ม 9" := "ยา 503",
                     "ปึ่ม 10" := "ยา 504",
                     "ปึ่ม 11" := "ยา 505",
                     "ปึ่ม 12" := "ยา 505",
                     "ปึ่ม 13" := "ยา 507",
                     "ปึ่ม 14" := "ยา 508",
                     "ปึ่ม 15" := "ยา 509",
                     "ปึ่ม 16" := "ยา 510",
                     "ปึ่ม 17" := "ยา 511",
                     "ปึ่ม 18" := "ยา 512",
                     "ปึ่ม 19" := "ยา 513",
                     "ปึ่ม 20" := "ยา 514",
                     "ปึ่ม 21" := "ยา 515",
                     "ปึ่ม 22" := "ยา 516",
                     "ปึ่ม 23" := "ยา 517",
                     "ปึ่ม 24" := "ยา 518",
                     "ปึ่ม 25" := "ยา 519",
                     "ปึ่ม 26" := "ยา 520",
                     "เมื่ิอมีการกดปุ้ม" => "output Step motor No.3  20",
                     ENO => #_w57);
   IF #_w57 AND "output Step motor No.3  20" THEN
       "SR Step Motro 3  เบิกจ่าย 20" := TRUE;   // SR flip-flop
   END_IF;
   IF "Output No1,2 Blackword 20" OR "ปุ่มClear" THEN "SR Step Motro 3  เบิกจ่าย 20" := FALSE; END_IF;
   "button start"(EN := "SR Step Motro 3  เบิกจ่าย 20", Output => "Output ปุ่มยืนยันหน้า Screen", ENO => #_w59);
   "IEC_Counter_0_DB_5".CTU(CU := (#_w4 OR #_w7 OR #_w10 OR #_w13 OR #_w16 OR #_w19 OR #_w22 OR #_w25 OR #_w28 OR #_w31 OR #_w34 OR #_w37 OR #_w40 OR #_w43 OR #_w46 OR #_w49 OR #_w52 OR #_w55 OR #_w58 OR (#_w59 AND "Output ปุ่มยืนยันหน้า Screen")) AND "Stepper Motor หยุดทำงาน หยุดสไลด์ ตัวงัดกล่องยาเข้า",
                           R := "Step Motor 3 Blackword_NO",
                           PV := 1);
   #"Stepper Motor  ทำงาน" := "IEC_Counter_0_DB_5".Q AND NOT "Step motor 1,2 NO" AND NOT "Stepper Motor ทำงาน สไลด์ ตัวงัดกล่องยาออก" AND NOT "Stepper Motor หยุดทำงาน หยุดสไลด์ ตัวงัดกล่องยาออก" AND NOT "Stepper Motor ทำงาน สไลด์ ตัวงัดกล่องยาเข้า" AND NOT "Stepper Motor หยุดทำงาน หยุดสไลด์ ตัวงัดกล่องยาเข้า";
END_REGION

